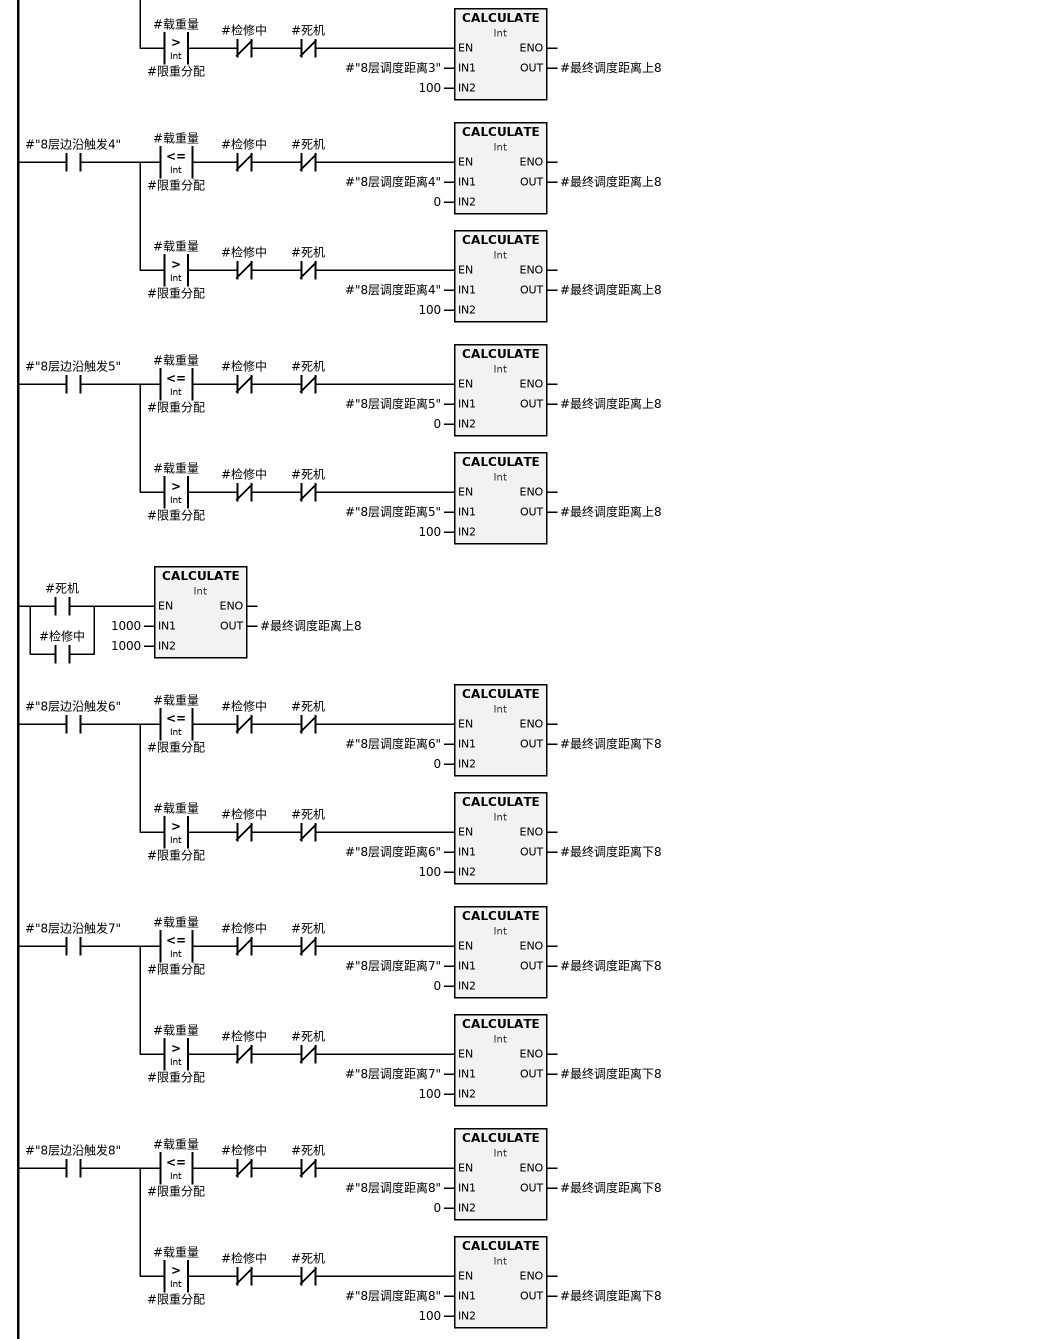
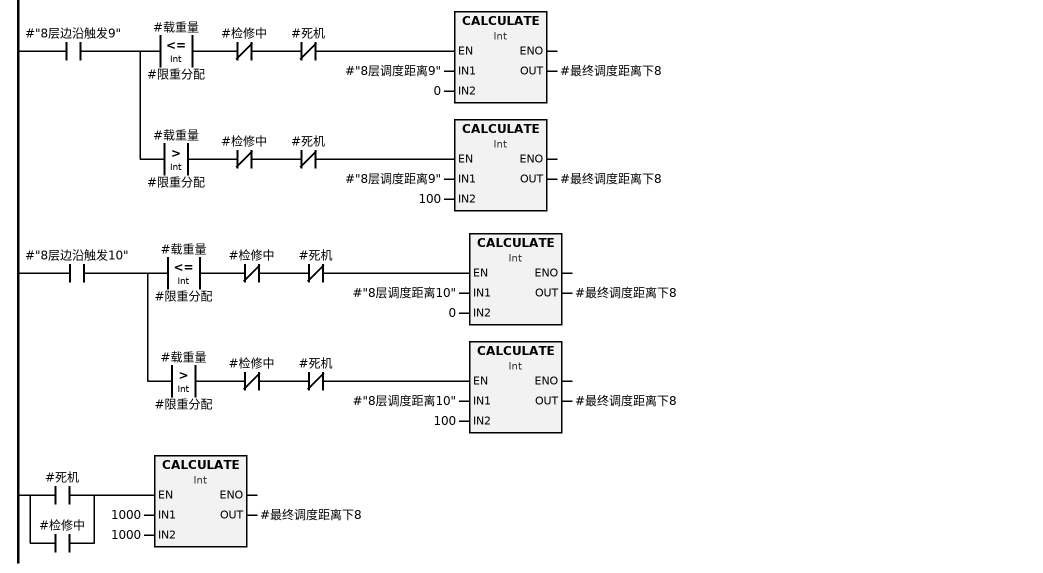
   RUNG wire#powerrail
      Contact( #上呼灯8 )
      wire#w1
      I_Contact( #上行指示 )
      I_Contact( #下行指示 )
      { S7_Templates := "SrcType := Int" } LE_Contact(in1 := #当前楼层, in2 := 8)
      wire#w2
      { S7_Templates := "SrcType := Int"; S7_Expression := "ABS(IN1-IN2)+IN3+IN3" } Calculate(in1 := #当前楼层, in2 := 8, in3 := #上行停站次数8, out => #"8层调度距离1")
      Coil( #"8层边沿触发1" )
   END_RUNG
   RUNG wire#w1
      Contact( #上行指示 )
      wire#w3
      { S7_Templates := "SrcType := Int" } EQ_Contact(in1 := 8, in2 := #当前楼层)
      Contact( #上下平层都为1 )
   END_RUNG wire#w2
   RUNG wire#w3
      { S7_Templates := "SrcType := Int" } GT_Contact(in1 := 8, in2 := #当前楼层)
   END_RUNG wire#w2
   RUNG wire#w1
      Contact( #下行指示 )
      wire#w4
      Contact( #外呼下面无目标8 )
      { S7_Templates := "SrcType := Int"; S7_Expression := "ABS(IN1-IN2)+IN3+IN3" } Calculate(in1 := #当前楼层, in2 := 8, in3 := #下行停站次数8, out => #"8层调度距离2")
      Coil( #"8层边沿触发2" )
   END_RUNG
   RUNG wire#w1
      I_Contact( #上行指示 )
      I_Contact( #下行指示 )
      { S7_Templates := "SrcType := Int" } GT_Contact(in1 := #当前楼层, in2 := 8)
   END_RUNG wire#w4
   RUNG wire#w1
      Contact( #下行指示 )
      Contact( #外呼下面有目标8 )
      { S7_Templates := "SrcType := Int"; S7_Expression := "ABS(IN3+IN3-IN1-IN2)+IN5+IN4+IN4+IN5+IN6" } Calculate(in1 := #当前楼层, in2 := 8, in3 := #外呼下面有目标最小数8, in4 := #上行停站次数8, in5 := #下行停站次数1, in6 := 2, out => #"8层调度距离3")
      Coil( #"8层边沿触发3" )
   END_RUNG
   RUNG wire#w1
      Contact( #上行指示 )
      wire#w5
      { S7_Templates := "SrcType := Int" } EQ_Contact(in1 := 8, in2 := #当前楼层)
      I_Contact( #上下平层都为1 )
      wire#w6
      Contact( #外呼下面有目标8 )
      { S7_Templates := "SrcType := Int"; S7_Expression := "ABS(IN3-IN1+IN3-IN6+IN2-IN6)+IN5+IN4+IN4+IN5+IN7+IN7" } Calculate(in1 := #当前楼层, in2 := 8, in3 := #外呼上面有目标最大数8, in4 := #上行停站次数10, in5 := #上行停站次数8, in6 := #外呼下面有目标最小数8, in7 := #下行停站次数1, in8 := 4, out => #"8层调度距离4")
      Coil( #"8层边沿触发4" )
   END_RUNG
   RUNG wire#w5
      { S7_Templates := "SrcType := Int" } LT_Contact(in1 := 8, in2 := #当前楼层)
   END_RUNG wire#w6
   RUNG wire#w6
      Contact( #外呼下面无目标8 )
      { S7_Templates := "SrcType := Int"; S7_Expression := "ABS(IN3-IN1+IN3-IN2)+IN5+IN4+IN4+IN5+IN6" } Calculate(in1 := #当前楼层, in2 := 8, in3 := #外呼上面有目标最大数8, in4 := #上行停站次数10, in5 := #下行停站次数8, in6 := 2, out => #"8层调度距离5")
      Coil( #"8层边沿触发5" )
   END_RUNG
   RUNG wire#powerrail
      Contact( #下呼灯8 )
      wire#w7
      I_Contact( #上行指示 )
      I_Contact( #下行指示 )
      { S7_Templates := "SrcType := Int" } GE_Contact(in1 := #当前楼层, in2 := 8)
      wire#w8
      { S7_Templates := "SrcType := Int"; S7_Expression := "ABS(IN1-IN2)+IN3+IN3" } Calculate(in1 := #当前楼层, in2 := 8, in3 := #下行停站次数8, out => #"8层调度距离6")
      Coil( #"8层边沿触发6" )
   END_RUNG
   RUNG wire#w7
      Contact( #下行指示 )
      wire#w9
      { S7_Templates := "SrcType := Int" } EQ_Contact(in1 := 8, in2 := #当前楼层)
      Contact( #上下平层都为1 )
   END_RUNG wire#w8
   RUNG wire#w9
      { S7_Templates := "SrcType := Int" } LT_Contact(in1 := 8, in2 := #当前楼层)
   END_RUNG wire#w8
   RUNG wire#w7
      Contact( #上行指示 )
      wire#w10
      Contact( #外呼上面无目标8 )
      { S7_Templates := "SrcType := Int"; S7_Expression := "ABS(IN1-IN2)+IN3+IN3" } Calculate(in1 := #当前楼层, in2 := 8, in3 := #上行停站次数8, out => #"8层调度距离7")
      Coil( #"8层边沿触发7" )
   END_RUNG
   RUNG wire#w7
      I_Contact( #上行指示 )
      I_Contact( #下行指示 )
      { S7_Templates := "SrcType := Int" } LT_Contact(in1 := #当前楼层, in2 := 8)
   END_RUNG wire#w10
   RUNG wire#w7
      Contact( #上行指示 )
      Contact( #外呼上面有目标8 )
      { S7_Templates := "SrcType := Int"; S7_Expression := "ABS(IN3+IN3-IN1-IN2)+IN4+IN5+IN4+IN5+IN6" } Calculate(in1 := #当前楼层, in2 := 8, in3 := #外呼上面有目标最大数8, in4 := #下行停站次数8, in5 := #上行停站次数10, in6 := 2, out => #"8层调度距离8")
      Coil( #"8层边沿触发8" )
   END_RUNG
   RUNG wire#w7
      Contact( #下行指示 )
      wire#w11
      { S7_Templates := "SrcType := Int" } EQ_Contact(in1 := 8, in2 := #当前楼层)
      I_Contact( #上下平层都为1 )
      wire#w12
      Contact( #外呼上面有目标8 )
      { S7_Templates := "SrcType := Int"; S7_Expression := "ABS(IN1-IN6+IN3-IN6+IN3-IN2)+IN5+IN4+IN4+IN5+IN7+IN7+IN8" } Calculate(in1 := #当前楼层, in2 := 8, in3 := #外呼上面有目标最大数8, in4 := #下行停站次数8, in5 := #下行停站次数1, in6 := #外呼下面有目标最小数8, in7 := #上行停站次数10, in8 := 4, out => #"8层调度距离9")
      Coil( #"8层边沿触发9" )
   END_RUNG
   RUNG wire#w11
      { S7_Templates := "SrcType := Int" } GT_Contact(in1 := 8, in2 := #当前楼层)
   END_RUNG wire#w12
   RUNG wire#w12
      Contact( #外呼上面无目标8 )
      { S7_Templates := "SrcType := Int"; S7_Expression := "ABS(IN1-IN3+IN2-IN3)+IN5+IN4+IN4+IN5+IN6" } Calculate(in1 := #当前楼层, in2 := 8, in3 := #外呼下面有目标最小数8, in4 := #上行停站次数8, in5 := #下行停站次数1, in6 := 2, out => #"8层调度距离10")
      Coil( #"8层边沿触发10" )
   END_RUNG
   RUNG wire#powerrail
      Contact( #"8层边沿触发1" )
      wire#w13
      { S7_Templates := "SrcType := Int" } LE_Contact(in1 := #载重量, in2 := #限重分配)
      I_Contact( #检修中 )
      I_Contact( #死机 )
      { S7_Templates := "SrcType := Int"; S7_Expression := "ABS(IN1+IN2)" } Calculate(in1 := #"8层调度距离1", in2 := 0, out => #最终调度距离上8)
   END_RUNG
   RUNG wire#w13
      { S7_Templates := "SrcType := Int" } GT_Contact(in1 := #载重量, in2 := #限重分配)
      I_Contact( #检修中 )
      I_Contact( #死机 )
      { S7_Templates := "SrcType := Int"; S7_Expression := "ABS(IN1+IN2)" } Calculate(in1 := #"8层调度距离1", in2 := 100, out => #最终调度距离上8)
   END_RUNG
   RUNG wire#powerrail
      Contact( #"8层边沿触发2" )
      wire#w14
      { S7_Templates := "SrcType := Int" } LE_Contact(in1 := #载重量, in2 := #限重分配)
      I_Contact( #检修中 )
      I_Contact( #死机 )
      { S7_Templates := "SrcType := Int"; S7_Expression := "ABS(IN1+IN2)" } Calculate(in1 := #"8层调度距离2", in2 := 0, out => #最终调度距离上8)
   END_RUNG
   RUNG wire#w14
      { S7_Templates := "SrcType := Int" } GT_Contact(in1 := #载重量, in2 := #限重分配)
      I_Contact( #检修中 )
      I_Contact( #死机 )
      { S7_Templates := "SrcType := Int"; S7_Expression := "ABS(IN1+IN2)" } Calculate(in1 := #"8层调度距离2", in2 := 100, out => #最终调度距离上8)
   END_RUNG
   RUNG wire#powerrail
      Contact( #"8层边沿触发3" )
      wire#w15
      { S7_Templates := "SrcType := Int" } LE_Contact(in1 := #载重量, in2 := #限重分配)
      I_Contact( #检修中 )
      I_Contact( #死机 )
      { S7_Templates := "SrcType := Int"; S7_Expression := "ABS(IN1+IN2)" } Calculate(in1 := #"8层调度距离3", in2 := 0, out => #最终调度距离上8)
   END_RUNG
   RUNG wire#w15
      { S7_Templates := "SrcType := Int" } GT_Contact(in1 := #载重量, in2 := #限重分配)
      I_Contact( #检修中 )
      I_Contact( #死机 )
      { S7_Templates := "SrcType := Int"; S7_Expression := "ABS(IN1+IN2)" } Calculate(in1 := #"8层调度距离3", in2 := 100, out => #最终调度距离上8)
   END_RUNG
   RUNG wire#powerrail
      Contact( #"8层边沿触发4" )
      wire#w16
      { S7_Templates := "SrcType := Int" } LE_Contact(in1 := #载重量, in2 := #限重分配)
      I_Contact( #检修中 )
      I_Contact( #死机 )
      { S7_Templates := "SrcType := Int"; S7_Expression := "ABS(IN1+IN2)" } Calculate(in1 := #"8层调度距离4", in2 := 0, out => #最终调度距离上8)
   END_RUNG
   RUNG wire#w16
      { S7_Templates := "SrcType := Int" } GT_Contact(in1 := #载重量, in2 := #限重分配)
      I_Contact( #检修中 )
      I_Contact( #死机 )
      { S7_Templates := "SrcType := Int"; S7_Expression := "ABS(IN1+IN2)" } Calculate(in1 := #"8层调度距离4", in2 := 100, out => #最终调度距离上8)
   END_RUNG
   RUNG wire#powerrail
      Contact( #"8层边沿触发5" )
      wire#w17
      { S7_Templates := "SrcType := Int" } LE_Contact(in1 := #载重量, in2 := #限重分配)
      I_Contact( #检修中 )
      I_Contact( #死机 )
      { S7_Templates := "SrcType := Int"; S7_Expression := "ABS(IN1+IN2)" } Calculate(in1 := #"8层调度距离5", in2 := 0, out => #最终调度距离上8)
   END_RUNG
   RUNG wire#w17
      { S7_Templates := "SrcType := Int" } GT_Contact(in1 := #载重量, in2 := #限重分配)
      I_Contact( #检修中 )
      I_Contact( #死机 )
      { S7_Templates := "SrcType := Int"; S7_Expression := "ABS(IN1+IN2)" } Calculate(in1 := #"8层调度距离5", in2 := 100, out => #最终调度距离上8)
   END_RUNG
   RUNG wire#powerrail
      Contact( #死机 )
      wire#w18
      { S7_Templates := "SrcType := Int"; S7_Expression := "ABS(IN1+IN2)" } Calculate(in1 := 1000, in2 := 1000, out => #最终调度距离上8)
   END_RUNG
   RUNG wire#powerrail
      Contact( #检修中 )
   END_RUNG wire#w18
   RUNG wire#powerrail
      Contact( #"8层边沿触发6" )
      wire#w19
      { S7_Templates := "SrcType := Int" } LE_Contact(in1 := #载重量, in2 := #限重分配)
      I_Contact( #检修中 )
      I_Contact( #死机 )
      { S7_Templates := "SrcType := Int"; S7_Expression := "ABS(IN1+IN2)" } Calculate(in1 := #"8层调度距离6", in2 := 0, out => #最终调度距离下8)
   END_RUNG
   RUNG wire#w19
      { S7_Templates := "SrcType := Int" } GT_Contact(in1 := #载重量, in2 := #限重分配)
      I_Contact( #检修中 )
      I_Contact( #死机 )
      { S7_Templates := "SrcType := Int"; S7_Expression := "ABS(IN1+IN2)" } Calculate(in1 := #"8层调度距离6", in2 := 100, out => #最终调度距离下8)
   END_RUNG
   RUNG wire#powerrail
      Contact( #"8层边沿触发7" )
      wire#w20
      { S7_Templates := "SrcType := Int" } LE_Contact(in1 := #载重量, in2 := #限重分配)
      I_Contact( #检修中 )
      I_Contact( #死机 )
      { S7_Templates := "SrcType := Int"; S7_Expression := "ABS(IN1+IN2)" } Calculate(in1 := #"8层调度距离7", in2 := 0, out => #最终调度距离下8)
   END_RUNG
   RUNG wire#w20
      { S7_Templates := "SrcType := Int" } GT_Contact(in1 := #载重量, in2 := #限重分配)
      I_Contact( #检修中 )
      I_Contact( #死机 )
      { S7_Templates := "SrcType := Int"; S7_Expression := "ABS(IN1+IN2)" } Calculate(in1 := #"8层调度距离7", in2 := 100, out => #最终调度距离下8)
   END_RUNG
   RUNG wire#powerrail
      Contact( #"8层边沿触发8" )
      wire#w21
      { S7_Templates := "SrcType := Int" } LE_Contact(in1 := #载重量, in2 := #限重分配)
      I_Contact( #检修中 )
      I_Contact( #死机 )
      { S7_Templates := "SrcType := Int"; S7_Expression := "ABS(IN1+IN2)" } Calculate(in1 := #"8层调度距离8", in2 := 0, out => #最终调度距离下8)
   END_RUNG
   RUNG wire#w21
      { S7_Templates := "SrcType := Int" } GT_Contact(in1 := #载重量, in2 := #限重分配)
      I_Contact( #检修中 )
      I_Contact( #死机 )
      { S7_Templates := "SrcType := Int"; S7_Expression := "ABS(IN1+IN2)" } Calculate(in1 := #"8层调度距离8", in2 := 100, out => #最终调度距离下8)
   END_RUNG
   RUNG wire#powerrail
      Contact( #"8层边沿触发9" )
      wire#w22
      { S7_Templates := "SrcType := Int" } LE_Contact(in1 := #载重量, in2 := #限重分配)
      I_Contact( #检修中 )
      I_Contact( #死机 )
      { S7_Templates := "SrcType := Int"; S7_Expression := "ABS(IN1+IN2)" } Calculate(in1 := #"8层调度距离9", in2 := 0, out => #最终调度距离下8)
   END_RUNG
   RUNG wire#w22
      { S7_Templates := "SrcType := Int" } GT_Contact(in1 := #载重量, in2 := #限重分配)
      I_Contact( #检修中 )
      I_Contact( #死机 )
      { S7_Templates := "SrcType := Int"; S7_Expression := "ABS(IN1+IN2)" } Calculate(in1 := #"8层调度距离9", in2 := 100, out => #最终调度距离下8)
   END_RUNG
   RUNG wire#powerrail
      Contact( #"8层边沿触发10" )
      wire#w23
      { S7_Templates := "SrcType := Int" } LE_Contact(in1 := #载重量, in2 := #限重分配)
      I_Contact( #检修中 )
      I_Contact( #死机 )
      { S7_Templates := "SrcType := Int"; S7_Expression := "ABS(IN1+IN2)" } Calculate(in1 := #"8层调度距离10", in2 := 0, out => #最终调度距离下8)
   END_RUNG
   RUNG wire#w23
      { S7_Templates := "SrcType := Int" } GT_Contact(in1 := #载重量, in2 := #限重分配)
      I_Contact( #检修中 )
      I_Contact( #死机 )
      { S7_Templates := "SrcType := Int"; S7_Expression := "ABS(IN1+IN2)" } Calculate(in1 := #"8层调度距离10", in2 := 100, out => #最终调度距离下8)
   END_RUNG
   RUNG wire#powerrail
      Contact( #死机 )
      wire#w24
      { S7_Templates := "SrcType := Int"; S7_Expression := "ABS(IN1+IN2)" } Calculate(in1 := 1000, in2 := 1000, out => #最终调度距离下8)
   END_RUNG
   RUNG wire#powerrail
      Contact( #检修中 )
   END_RUNG wire#w24
   // the same network as SCL:
   #_w1 := #上呼灯8 AND ((NOT #上行指示 AND NOT #下行指示 AND (#当前楼层 <= 8)) OR (#上行指示 AND (((8 = #当前楼层) AND #上下平层都为1) OR (8 > #当前楼层))));
   IF #_w1 THEN #"8层调度距离1" := ABS(#当前楼层-8)+#上行停站次数8+#上行停站次数8; END_IF;
   #"8层边沿触发1" := #_w1;
   #_w2 := #上呼灯8 AND (#下行指示 OR (NOT #上行指示 AND NOT #下行指示 AND (#当前楼层 > 8))) AND #外呼下面无目标8;
   IF #_w2 THEN #"8层调度距离2" := ABS(#当前楼层-8)+#下行停站次数8+#下行停站次数8; END_IF;
   #"8层边沿触发2" := #_w2;
   #_w3 := #上呼灯8 AND #下行指示 AND #外呼下面有目标8;
   IF #_w3 THEN
       #"8层调度距离3" := ABS(#外呼下面有目标最小数8+#外呼下面有目标最小数8-#当前楼层-8)+#下行停站次数1+#上行停站次数8+#上行停站次数8+#下行停站次数1+2;
   END_IF;
   #"8层边沿触发3" := #_w3;
   #_w4 := #上呼灯8 AND #上行指示 AND (((8 = #当前楼层) AND NOT #上下平层都为1) OR (8 < #当前楼层));
   #_w5 := #_w4 AND #外呼下面有目标8;
   IF #_w5 THEN
       #"8层调度距离4" := ABS(#外呼上面有目标最大数8-#当前楼层+#外呼上面有目标最大数8-#外呼下面有目标最小数8+8-#外呼下面有目标最小数8)+#上行停站次数8+#上行停站次数10+#上行停站次数10+#上行停站次数8+#下行停站次数1+#下行停站次数1;
   END_IF;
   #"8层边沿触发4" := #_w5;
   #_w6 := #_w4 AND #外呼下面无目标8;
   IF #_w6 THEN
       #"8层调度距离5" := ABS(#外呼上面有目标最大数8-#当前楼层+#外呼上面有目标最大数8-8)+#下行停站次数8+#上行停站次数10+#上行停站次数10+#下行停站次数8+2;
   END_IF;
   #"8层边沿触发5" := #_w6;
   #_w7 := #下呼灯8 AND ((NOT #上行指示 AND NOT #下行指示 AND (#当前楼层 >= 8)) OR (#下行指示 AND (((8 = #当前楼层) AND #上下平层都为1) OR (8 < #当前楼层))));
   IF #_w7 THEN #"8层调度距离6" := ABS(#当前楼层-8)+#下行停站次数8+#下行停站次数8; END_IF;
   #"8层边沿触发6" := #_w7;
   #_w8 := #下呼灯8 AND (#上行指示 OR (NOT #上行指示 AND NOT #下行指示 AND (#当前楼层 < 8))) AND #外呼上面无目标8;
   IF #_w8 THEN #"8层调度距离7" := ABS(#当前楼层-8)+#上行停站次数8+#上行停站次数8; END_IF;
   #"8层边沿触发7" := #_w8;
   #_w9 := #下呼灯8 AND #上行指示 AND #外呼上面有目标8;
   IF #_w9 THEN
       #"8层调度距离8" := ABS(#外呼上面有目标最大数8+#外呼上面有目标最大数8-#当前楼层-8)+#下行停站次数8+#上行停站次数10+#下行停站次数8+#上行停站次数10+2;
   END_IF;
   #"8层边沿触发8" := #_w9;
   #_w10 := #下呼灯8 AND #下行指示 AND (((8 = #当前楼层) AND NOT #上下平层都为1) OR (8 > #当前楼层));
   #_w11 := #_w10 AND #外呼上面有目标8;
   IF #_w11 THEN
       #"8层调度距离9" := ABS(#当前楼层-#外呼下面有目标最小数8+#外呼上面有目标最大数8-#外呼下面有目标最小数8+#外呼上面有目标最大数8-8)+#下行停站次数1+#下行停站次数8+#下行停站次数8+#下行停站次数1+#上行停站次数10+#上行停站次数10+4;
   END_IF;
   #"8层边沿触发9" := #_w11;
   #_w12 := #_w10 AND #外呼上面无目标8;
   IF #_w12 THEN
       #"8层调度距离10" := ABS(#当前楼层-#外呼下面有目标最小数8+8-#外呼下面有目标最小数8)+#下行停站次数1+#上行停站次数8+#上行停站次数8+#下行停站次数1+2;
   END_IF;
   #"8层边沿触发10" := #_w12;
   IF #"8层边沿触发1" AND (#载重量 <= #限重分配) AND NOT #检修中 AND NOT #死机 THEN #最终调度距离上8 := ABS(#"8层调度距离1"+0); END_IF;
   IF #"8层边沿触发1" AND (#载重量 > #限重分配) AND NOT #检修中 AND NOT #死机 THEN #最终调度距离上8 := ABS(#"8层调度距离1"+100); END_IF;
   IF #"8层边沿触发2" AND (#载重量 <= #限重分配) AND NOT #检修中 AND NOT #死机 THEN #最终调度距离上8 := ABS(#"8层调度距离2"+0); END_IF;
   IF #"8层边沿触发2" AND (#载重量 > #限重分配) AND NOT #检修中 AND NOT #死机 THEN #最终调度距离上8 := ABS(#"8层调度距离2"+100); END_IF;
   IF #"8层边沿触发3" AND (#载重量 <= #限重分配) AND NOT #检修中 AND NOT #死机 THEN #最终调度距离上8 := ABS(#"8层调度距离3"+0); END_IF;
   IF #"8层边沿触发3" AND (#载重量 > #限重分配) AND NOT #检修中 AND NOT #死机 THEN #最终调度距离上8 := ABS(#"8层调度距离3"+100); END_IF;
   IF #"8层边沿触发4" AND (#载重量 <= #限重分配) AND NOT #检修中 AND NOT #死机 THEN #最终调度距离上8 := ABS(#"8层调度距离4"+0); END_IF;
   IF #"8层边沿触发4" AND (#载重量 > #限重分配) AND NOT #检修中 AND NOT #死机 THEN #最终调度距离上8 := ABS(#"8层调度距离4"+100); END_IF;
   IF #"8层边沿触发5" AND (#载重量 <= #限重分配) AND NOT #检修中 AND NOT #死机 THEN #最终调度距离上8 := ABS(#"8层调度距离5"+0); END_IF;
   IF #"8层边沿触发5" AND (#载重量 > #限重分配) AND NOT #检修中 AND NOT #死机 THEN #最终调度距离上8 := ABS(#"8层调度距离5"+100); END_IF;
   IF #死机 OR #检修中 THEN #最终调度距离上8 := ABS(1000+1000); END_IF;
   IF #"8层边沿触发6" AND (#载重量 <= #限重分配) AND NOT #检修中 AND NOT #死机 THEN #最终调度距离下8 := ABS(#"8层调度距离6"+0); END_IF;
   IF #"8层边沿触发6" AND (#载重量 > #限重分配) AND NOT #检修中 AND NOT #死机 THEN #最终调度距离下8 := ABS(#"8层调度距离6"+100); END_IF;
   IF #"8层边沿触发7" AND (#载重量 <= #限重分配) AND NOT #检修中 AND NOT #死机 THEN #最终调度距离下8 := ABS(#"8层调度距离7"+0); END_IF;
   IF #"8层边沿触发7" AND (#载重量 > #限重分配) AND NOT #检修中 AND NOT #死机 THEN #最终调度距离下8 := ABS(#"8层调度距离7"+100); END_IF;
   IF #"8层边沿触发8" AND (#载重量 <= #限重分配) AND NOT #检修中 AND NOT #死机 THEN #最终调度距离下8 := ABS(#"8层调度距离8"+0); END_IF;
   IF #"8层边沿触发8" AND (#载重量 > #限重分配) AND NOT #检修中 AND NOT #死机 THEN #最终调度距离下8 := ABS(#"8层调度距离8"+100); END_IF;
   IF #"8层边沿触发9" AND (#载重量 <= #限重分配) AND NOT #检修中 AND NOT #死机 THEN #最终调度距离下8 := ABS(#"8层调度距离9"+0); END_IF;
   IF #"8层边沿触发9" AND (#载重量 > #限重分配) AND NOT #检修中 AND NOT #死机 THEN #最终调度距离下8 := ABS(#"8层调度距离9"+100); END_IF;
   IF #"8层边沿触发10" AND (#载重量 <= #限重分配) AND NOT #检修中 AND NOT #死机 THEN #最终调度距离下8 := ABS(#"8层调度距离10"+0); END_IF;
   IF #"8层边沿触发10" AND (#载重量 > #限重分配) AND NOT #检修中 AND NOT #死机 THEN #最终调度距离下8 := ABS(#"8层调度距离10"+100); END_IF;
   IF #死机 OR #检修中 THEN #最终调度距离下8 := ABS(1000+1000); END_IF;
END_REGION

REGION Network 8: 9层调度距离
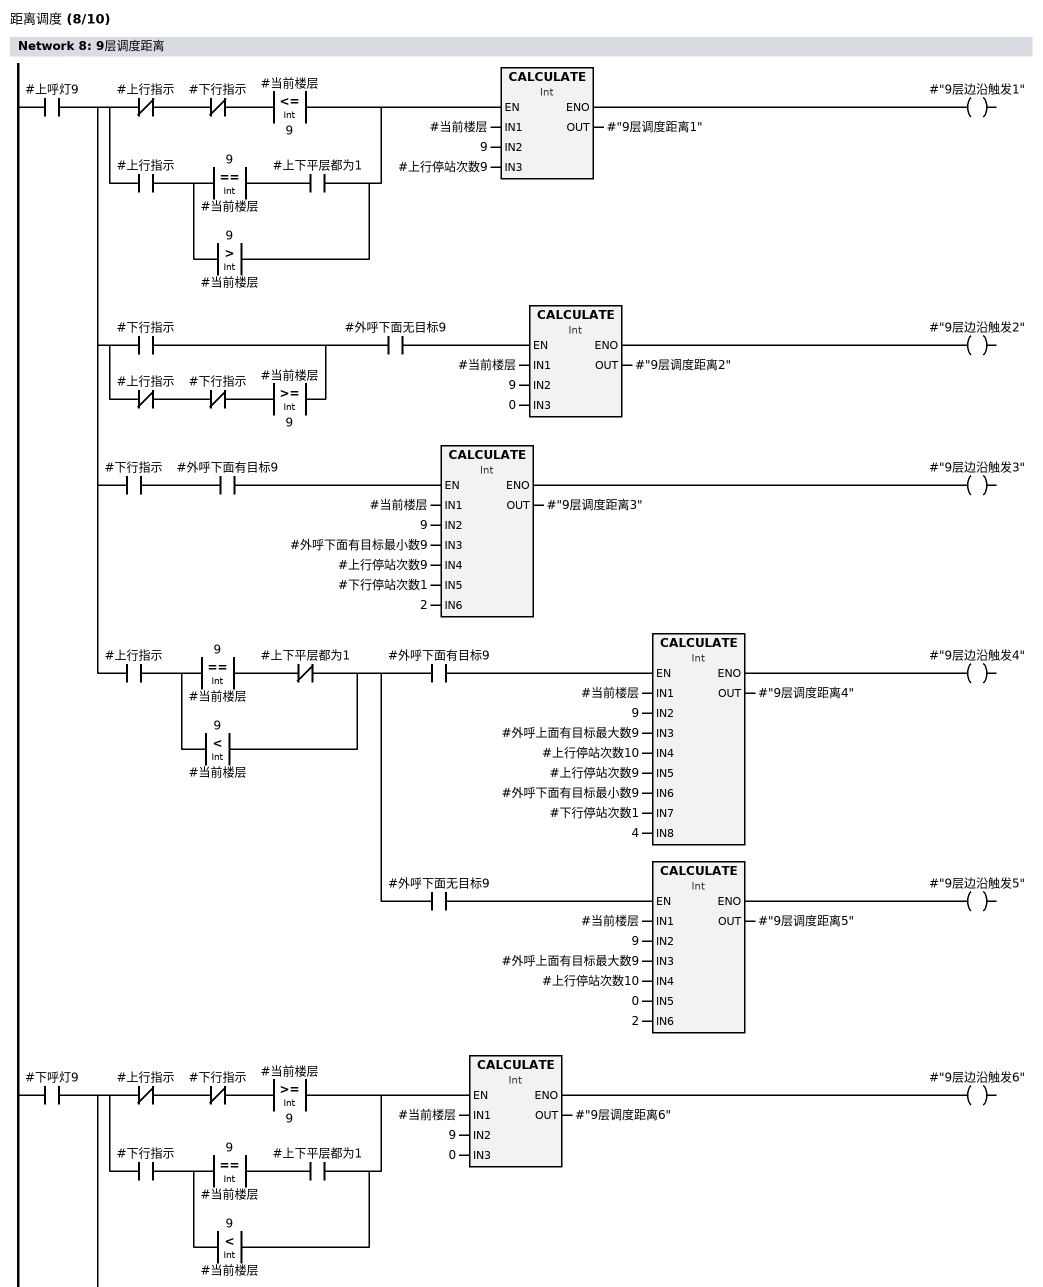
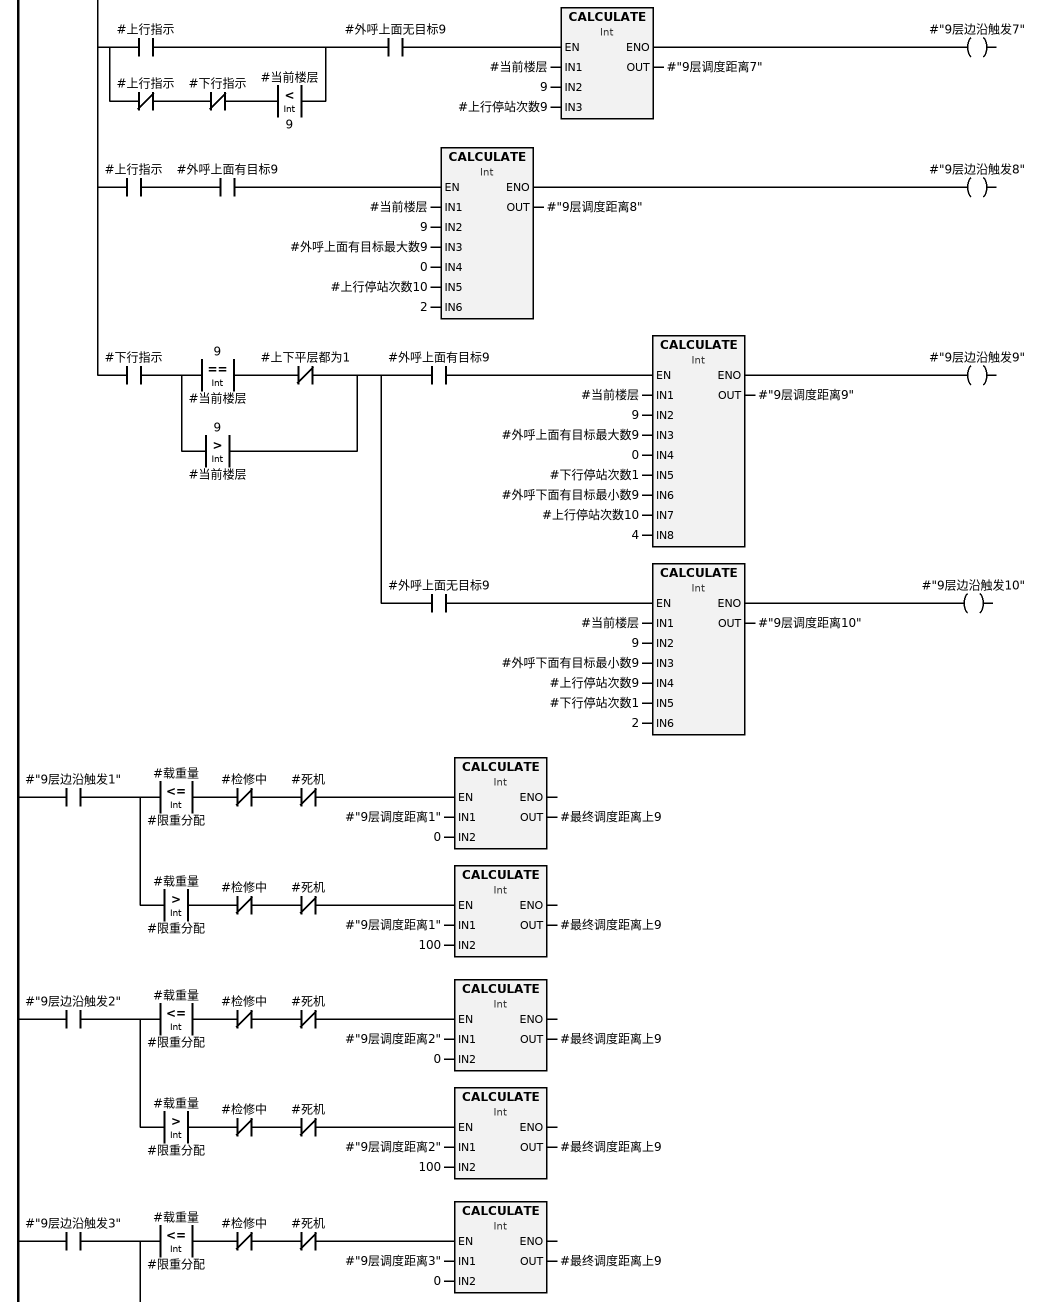
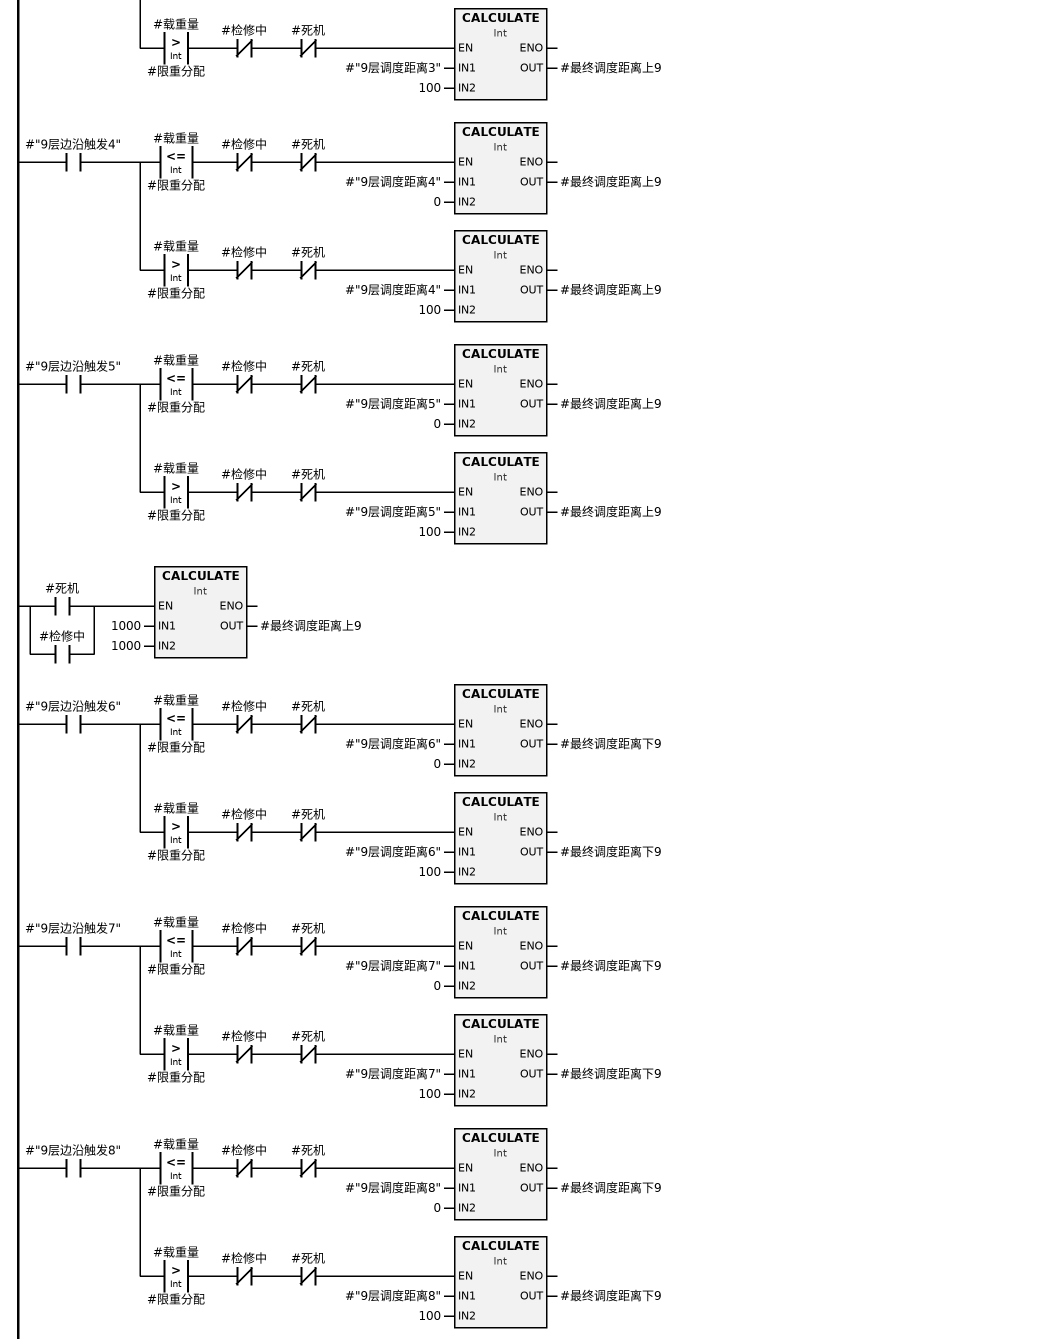
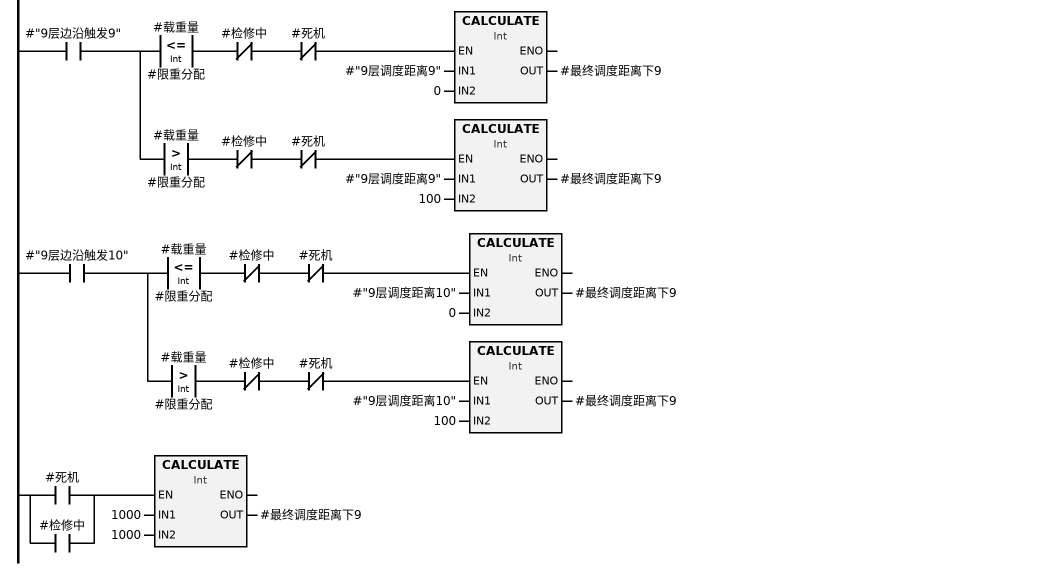
   RUNG wire#powerrail
      Contact( #上呼灯9 )
      wire#w1
      I_Contact( #上行指示 )
      I_Contact( #下行指示 )
      { S7_Templates := "SrcType := Int" } LE_Contact(in1 := #当前楼层, in2 := 9)
      wire#w2
      { S7_Templates := "SrcType := Int"; S7_Expression := "ABS(IN1-IN2)+IN3+IN3" } Calculate(in1 := #当前楼层, in2 := 9, in3 := #上行停站次数9, out => #"9层调度距离1")
      Coil( #"9层边沿触发1" )
   END_RUNG
   RUNG wire#w1
      Contact( #上行指示 )
      wire#w3
      { S7_Templates := "SrcType := Int" } EQ_Contact(in1 := 9, in2 := #当前楼层)
      Contact( #上下平层都为1 )
   END_RUNG wire#w2
   RUNG wire#w3
      { S7_Templates := "SrcType := Int" } GT_Contact(in1 := 9, in2 := #当前楼层)
   END_RUNG wire#w2
   RUNG wire#w1
      Contact( #下行指示 )
      wire#w4
      Contact( #外呼下面无目标9 )
      { S7_Templates := "SrcType := Int"; S7_Expression := "ABS(IN1-IN2)+IN3+IN3" } Calculate(in1 := #当前楼层, in2 := 9, in3 := 0, out => #"9层调度距离2")
      Coil( #"9层边沿触发2" )
   END_RUNG
   RUNG wire#w1
      I_Contact( #上行指示 )
      I_Contact( #下行指示 )
      { S7_Templates := "SrcType := Int" } GE_Contact(in1 := #当前楼层, in2 := 9)
   END_RUNG wire#w4
   RUNG wire#w1
      Contact( #下行指示 )
      Contact( #外呼下面有目标9 )
      { S7_Templates := "SrcType := Int"; S7_Expression := "ABS(IN3+IN3-IN1-IN2)+IN5+IN4+IN4+IN5+IN6" } Calculate(in1 := #当前楼层, in2 := 9, in3 := #外呼下面有目标最小数9, in4 := #上行停站次数9, in5 := #下行停站次数1, in6 := 2, out => #"9层调度距离3")
      Coil( #"9层边沿触发3" )
   END_RUNG
   RUNG wire#w1
      Contact( #上行指示 )
      wire#w5
      { S7_Templates := "SrcType := Int" } EQ_Contact(in1 := 9, in2 := #当前楼层)
      I_Contact( #上下平层都为1 )
      wire#w6
      Contact( #外呼下面有目标9 )
      { S7_Templates := "SrcType := Int"; S7_Expression := "ABS(IN3-IN1+IN3-IN6+IN2-IN6)+IN5+IN4+IN4+IN5+IN7+IN7+IN8" } Calculate(in1 := #当前楼层, in2 := 9, in3 := #外呼上面有目标最大数9, in4 := #上行停站次数10, in5 := #上行停站次数9, in6 := #外呼下面有目标最小数9, in7 := #下行停站次数1, in8 := 4, out => #"9层调度距离4")
      Coil( #"9层边沿触发4" )
   END_RUNG
   RUNG wire#w5
      { S7_Templates := "SrcType := Int" } LT_Contact(in1 := 9, in2 := #当前楼层)
   END_RUNG wire#w6
   RUNG wire#w6
      Contact( #外呼下面无目标9 )
      { S7_Templates := "SrcType := Int"; S7_Expression := "ABS(IN3-IN1+IN3-IN2)+IN5+IN4+IN4+IN5+IN6" } Calculate(in1 := #当前楼层, in2 := 9, in3 := #外呼上面有目标最大数9, in4 := #上行停站次数10, in5 := 0, in6 := 2, out => #"9层调度距离5")
      Coil( #"9层边沿触发5" )
   END_RUNG
   RUNG wire#powerrail
      Contact( #下呼灯9 )
      wire#w7
      I_Contact( #上行指示 )
      I_Contact( #下行指示 )
      { S7_Templates := "SrcType := Int" } GE_Contact(in1 := #当前楼层, in2 := 9)
      wire#w8
      { S7_Templates := "SrcType := Int"; S7_Expression := "ABS(IN1-IN2)+IN3+IN3" } Calculate(in1 := #当前楼层, in2 := 9, in3 := 0, out => #"9层调度距离6")
      Coil( #"9层边沿触发6" )
   END_RUNG
   RUNG wire#w7
      Contact( #下行指示 )
      wire#w9
      { S7_Templates := "SrcType := Int" } EQ_Contact(in1 := 9, in2 := #当前楼层)
      Contact( #上下平层都为1 )
   END_RUNG wire#w8
   RUNG wire#w9
      { S7_Templates := "SrcType := Int" } LT_Contact(in1 := 9, in2 := #当前楼层)
   END_RUNG wire#w8
   RUNG wire#w7
      Contact( #上行指示 )
      wire#w10
      Contact( #外呼上面无目标9 )
      { S7_Templates := "SrcType := Int"; S7_Expression := "ABS(IN1-IN2)+IN3+IN3" } Calculate(in1 := #当前楼层, in2 := 9, in3 := #上行停站次数9, out => #"9层调度距离7")
      Coil( #"9层边沿触发7" )
   END_RUNG
   RUNG wire#w7
      I_Contact( #上行指示 )
      I_Contact( #下行指示 )
      { S7_Templates := "SrcType := Int" } LT_Contact(in1 := #当前楼层, in2 := 9)
   END_RUNG wire#w10
   RUNG wire#w7
      Contact( #上行指示 )
      Contact( #外呼上面有目标9 )
      { S7_Templates := "SrcType := Int"; S7_Expression := "ABS(IN3+IN3-IN1-IN2)+IN4+IN5+IN4+IN5+IN6" } Calculate(in1 := #当前楼层, in2 := 9, in3 := #外呼上面有目标最大数9, in4 := 0, in5 := #上行停站次数10, in6 := 2, out => #"9层调度距离8")
      Coil( #"9层边沿触发8" )
   END_RUNG
   RUNG wire#w7
      Contact( #下行指示 )
      wire#w11
      { S7_Templates := "SrcType := Int" } EQ_Contact(in1 := 9, in2 := #当前楼层)
      I_Contact( #上下平层都为1 )
      wire#w12
      Contact( #外呼上面有目标9 )
      { S7_Templates := "SrcType := Int"; S7_Expression := "ABS(IN1-IN6+IN3-IN6+IN3-IN2)+IN5+IN4+IN4+IN5+IN7+IN7+IN8" } Calculate(in1 := #当前楼层, in2 := 9, in3 := #外呼上面有目标最大数9, in4 := 0, in5 := #下行停站次数1, in6 := #外呼下面有目标最小数9, in7 := #上行停站次数10, in8 := 4, out => #"9层调度距离9")
      Coil( #"9层边沿触发9" )
   END_RUNG
   RUNG wire#w11
      { S7_Templates := "SrcType := Int" } GT_Contact(in1 := 9, in2 := #当前楼层)
   END_RUNG wire#w12
   RUNG wire#w12
      Contact( #外呼上面无目标9 )
      { S7_Templates := "SrcType := Int"; S7_Expression := "ABS(IN1-IN3+IN2-IN3)+IN5+IN4+IN4+IN5+IN6" } Calculate(in1 := #当前楼层, in2 := 9, in3 := #外呼下面有目标最小数9, in4 := #上行停站次数9, in5 := #下行停站次数1, in6 := 2, out => #"9层调度距离10")
      Coil( #"9层边沿触发10" )
   END_RUNG
   RUNG wire#powerrail
      Contact( #"9层边沿触发1" )
      wire#w13
      { S7_Templates := "SrcType := Int" } LE_Contact(in1 := #载重量, in2 := #限重分配)
      I_Contact( #检修中 )
      I_Contact( #死机 )
      { S7_Templates := "SrcType := Int"; S7_Expression := "ABS(IN1+IN2)" } Calculate(in1 := #"9层调度距离1", in2 := 0, out => #最终调度距离上9)
   END_RUNG
   RUNG wire#w13
      { S7_Templates := "SrcType := Int" } GT_Contact(in1 := #载重量, in2 := #限重分配)
      I_Contact( #检修中 )
      I_Contact( #死机 )
      { S7_Templates := "SrcType := Int"; S7_Expression := "ABS(IN1+IN2)" } Calculate(in1 := #"9层调度距离1", in2 := 100, out => #最终调度距离上9)
   END_RUNG
   RUNG wire#powerrail
      Contact( #"9层边沿触发2" )
      wire#w14
      { S7_Templates := "SrcType := Int" } LE_Contact(in1 := #载重量, in2 := #限重分配)
      I_Contact( #检修中 )
      I_Contact( #死机 )
      { S7_Templates := "SrcType := Int"; S7_Expression := "ABS(IN1+IN2)" } Calculate(in1 := #"9层调度距离2", in2 := 0, out => #最终调度距离上9)
   END_RUNG
   RUNG wire#w14
      { S7_Templates := "SrcType := Int" } GT_Contact(in1 := #载重量, in2 := #限重分配)
      I_Contact( #检修中 )
      I_Contact( #死机 )
      { S7_Templates := "SrcType := Int"; S7_Expression := "ABS(IN1+IN2)" } Calculate(in1 := #"9层调度距离2", in2 := 100, out => #最终调度距离上9)
   END_RUNG
   RUNG wire#powerrail
      Contact( #"9层边沿触发3" )
      wire#w15
      { S7_Templates := "SrcType := Int" } LE_Contact(in1 := #载重量, in2 := #限重分配)
      I_Contact( #检修中 )
      I_Contact( #死机 )
      { S7_Templates := "SrcType := Int"; S7_Expression := "ABS(IN1+IN2)" } Calculate(in1 := #"9层调度距离3", in2 := 0, out => #最终调度距离上9)
   END_RUNG
   RUNG wire#w15
      { S7_Templates := "SrcType := Int" } GT_Contact(in1 := #载重量, in2 := #限重分配)
      I_Contact( #检修中 )
      I_Contact( #死机 )
      { S7_Templates := "SrcType := Int"; S7_Expression := "ABS(IN1+IN2)" } Calculate(in1 := #"9层调度距离3", in2 := 100, out => #最终调度距离上9)
   END_RUNG
   RUNG wire#powerrail
      Contact( #"9层边沿触发4" )
      wire#w16
      { S7_Templates := "SrcType := Int" } LE_Contact(in1 := #载重量, in2 := #限重分配)
      I_Contact( #检修中 )
      I_Contact( #死机 )
      { S7_Templates := "SrcType := Int"; S7_Expression := "ABS(IN1+IN2)" } Calculate(in1 := #"9层调度距离4", in2 := 0, out => #最终调度距离上9)
   END_RUNG
   RUNG wire#w16
      { S7_Templates := "SrcType := Int" } GT_Contact(in1 := #载重量, in2 := #限重分配)
      I_Contact( #检修中 )
      I_Contact( #死机 )
      { S7_Templates := "SrcType := Int"; S7_Expression := "ABS(IN1+IN2)" } Calculate(in1 := #"9层调度距离4", in2 := 100, out => #最终调度距离上9)
   END_RUNG
   RUNG wire#powerrail
      Contact( #"9层边沿触发5" )
      wire#w17
      { S7_Templates := "SrcType := Int" } LE_Contact(in1 := #载重量, in2 := #限重分配)
      I_Contact( #检修中 )
      I_Contact( #死机 )
      { S7_Templates := "SrcType := Int"; S7_Expression := "ABS(IN1+IN2)" } Calculate(in1 := #"9层调度距离5", in2 := 0, out => #最终调度距离上9)
   END_RUNG
   RUNG wire#w17
      { S7_Templates := "SrcType := Int" } GT_Contact(in1 := #载重量, in2 := #限重分配)
      I_Contact( #检修中 )
      I_Contact( #死机 )
      { S7_Templates := "SrcType := Int"; S7_Expression := "ABS(IN1+IN2)" } Calculate(in1 := #"9层调度距离5", in2 := 100, out => #最终调度距离上9)
   END_RUNG
   RUNG wire#powerrail
      Contact( #死机 )
      wire#w18
      { S7_Templates := "SrcType := Int"; S7_Expression := "ABS(IN1+IN2)" } Calculate(in1 := 1000, in2 := 1000, out => #最终调度距离上9)
   END_RUNG
   RUNG wire#powerrail
      Contact( #检修中 )
   END_RUNG wire#w18
   RUNG wire#powerrail
      Contact( #"9层边沿触发6" )
      wire#w19
      { S7_Templates := "SrcType := Int" } LE_Contact(in1 := #载重量, in2 := #限重分配)
      I_Contact( #检修中 )
      I_Contact( #死机 )
      { S7_Templates := "SrcType := Int"; S7_Expression := "ABS(IN1+IN2)" } Calculate(in1 := #"9层调度距离6", in2 := 0, out => #最终调度距离下9)
   END_RUNG
   RUNG wire#w19
      { S7_Templates := "SrcType := Int" } GT_Contact(in1 := #载重量, in2 := #限重分配)
      I_Contact( #检修中 )
      I_Contact( #死机 )
      { S7_Templates := "SrcType := Int"; S7_Expression := "ABS(IN1+IN2)" } Calculate(in1 := #"9层调度距离6", in2 := 100, out => #最终调度距离下9)
   END_RUNG
   RUNG wire#powerrail
      Contact( #"9层边沿触发7" )
      wire#w20
      { S7_Templates := "SrcType := Int" } LE_Contact(in1 := #载重量, in2 := #限重分配)
      I_Contact( #检修中 )
      I_Contact( #死机 )
      { S7_Templates := "SrcType := Int"; S7_Expression := "ABS(IN1+IN2)" } Calculate(in1 := #"9层调度距离7", in2 := 0, out => #最终调度距离下9)
   END_RUNG
   RUNG wire#w20
      { S7_Templates := "SrcType := Int" } GT_Contact(in1 := #载重量, in2 := #限重分配)
      I_Contact( #检修中 )
      I_Contact( #死机 )
      { S7_Templates := "SrcType := Int"; S7_Expression := "ABS(IN1+IN2)" } Calculate(in1 := #"9层调度距离7", in2 := 100, out => #最终调度距离下9)
   END_RUNG
   RUNG wire#powerrail
      Contact( #"9层边沿触发8" )
      wire#w21
      { S7_Templates := "SrcType := Int" } LE_Contact(in1 := #载重量, in2 := #限重分配)
      I_Contact( #检修中 )
      I_Contact( #死机 )
      { S7_Templates := "SrcType := Int"; S7_Expression := "ABS(IN1+IN2)" } Calculate(in1 := #"9层调度距离8", in2 := 0, out => #最终调度距离下9)
   END_RUNG
   RUNG wire#w21
      { S7_Templates := "SrcType := Int" } GT_Contact(in1 := #载重量, in2 := #限重分配)
      I_Contact( #检修中 )
      I_Contact( #死机 )
      { S7_Templates := "SrcType := Int"; S7_Expression := "ABS(IN1+IN2)" } Calculate(in1 := #"9层调度距离8", in2 := 100, out => #最终调度距离下9)
   END_RUNG
   RUNG wire#powerrail
      Contact( #"9层边沿触发9" )
      wire#w22
      { S7_Templates := "SrcType := Int" } LE_Contact(in1 := #载重量, in2 := #限重分配)
      I_Contact( #检修中 )
      I_Contact( #死机 )
      { S7_Templates := "SrcType := Int"; S7_Expression := "ABS(IN1+IN2)" } Calculate(in1 := #"9层调度距离9", in2 := 0, out => #最终调度距离下9)
   END_RUNG
   RUNG wire#w22
      { S7_Templates := "SrcType := Int" } GT_Contact(in1 := #载重量, in2 := #限重分配)
      I_Contact( #检修中 )
      I_Contact( #死机 )
      { S7_Templates := "SrcType := Int"; S7_Expression := "ABS(IN1+IN2)" } Calculate(in1 := #"9层调度距离9", in2 := 100, out => #最终调度距离下9)
   END_RUNG
   RUNG wire#powerrail
      Contact( #"9层边沿触发10" )
      wire#w23
      { S7_Templates := "SrcType := Int" } LE_Contact(in1 := #载重量, in2 := #限重分配)
      I_Contact( #检修中 )
      I_Contact( #死机 )
      { S7_Templates := "SrcType := Int"; S7_Expression := "ABS(IN1+IN2)" } Calculate(in1 := #"9层调度距离10", in2 := 0, out => #最终调度距离下9)
   END_RUNG
   RUNG wire#w23
      { S7_Templates := "SrcType := Int" } GT_Contact(in1 := #载重量, in2 := #限重分配)
      I_Contact( #检修中 )
      I_Contact( #死机 )
      { S7_Templates := "SrcType := Int"; S7_Expression := "ABS(IN1+IN2)" } Calculate(in1 := #"9层调度距离10", in2 := 100, out => #最终调度距离下9)
   END_RUNG
   RUNG wire#powerrail
      Contact( #死机 )
      wire#w24
      { S7_Templates := "SrcType := Int"; S7_Expression := "ABS(IN1+IN2)" } Calculate(in1 := 1000, in2 := 1000, out => #最终调度距离下9)
   END_RUNG
   RUNG wire#powerrail
      Contact( #检修中 )
   END_RUNG wire#w24
   // the same network as SCL:
   #_w1 := #上呼灯9 AND ((NOT #上行指示 AND NOT #下行指示 AND (#当前楼层 <= 9)) OR (#上行指示 AND (((9 = #当前楼层) AND #上下平层都为1) OR (9 > #当前楼层))));
   IF #_w1 THEN #"9层调度距离1" := ABS(#当前楼层-9)+#上行停站次数9+#上行停站次数9; END_IF;
   #"9层边沿触发1" := #_w1;
   #_w2 := #上呼灯9 AND (#下行指示 OR (NOT #上行指示 AND NOT #下行指示 AND (#当前楼层 >= 9))) AND #外呼下面无目标9;
   IF #_w2 THEN #"9层调度距离2" := ABS(#当前楼层-9)+0+0; END_IF;
   #"9层边沿触发2" := #_w2;
   #_w3 := #上呼灯9 AND #下行指示 AND #外呼下面有目标9;
   IF #_w3 THEN
       #"9层调度距离3" := ABS(#外呼下面有目标最小数9+#外呼下面有目标最小数9-#当前楼层-9)+#下行停站次数1+#上行停站次数9+#上行停站次数9+#下行停站次数1+2;
   END_IF;
   #"9层边沿触发3" := #_w3;
   #_w4 := #上呼灯9 AND #上行指示 AND (((9 = #当前楼层) AND NOT #上下平层都为1) OR (9 < #当前楼层));
   #_w5 := #_w4 AND #外呼下面有目标9;
   IF #_w5 THEN
       #"9层调度距离4" := ABS(#外呼上面有目标最大数9-#当前楼层+#外呼上面有目标最大数9-#外呼下面有目标最小数9+9-#外呼下面有目标最小数9)+#上行停站次数9+#上行停站次数10+#上行停站次数10+#上行停站次数9+#下行停站次数1+#下行停站次数1+4;
   END_IF;
   #"9层边沿触发4" := #_w5;
   #_w6 := #_w4 AND #外呼下面无目标9;
   IF #_w6 THEN #"9层调度距离5" := ABS(#外呼上面有目标最大数9-#当前楼层+#外呼上面有目标最大数9-9)+0+#上行停站次数10+#上行停站次数10+0+2; END_IF;
   #"9层边沿触发5" := #_w6;
   #_w7 := #下呼灯9 AND ((NOT #上行指示 AND NOT #下行指示 AND (#当前楼层 >= 9)) OR (#下行指示 AND (((9 = #当前楼层) AND #上下平层都为1) OR (9 < #当前楼层))));
   IF #_w7 THEN #"9层调度距离6" := ABS(#当前楼层-9)+0+0; END_IF;
   #"9层边沿触发6" := #_w7;
   #_w8 := #下呼灯9 AND (#上行指示 OR (NOT #上行指示 AND NOT #下行指示 AND (#当前楼层 < 9))) AND #外呼上面无目标9;
   IF #_w8 THEN #"9层调度距离7" := ABS(#当前楼层-9)+#上行停站次数9+#上行停站次数9; END_IF;
   #"9层边沿触发7" := #_w8;
   #_w9 := #下呼灯9 AND #上行指示 AND #外呼上面有目标9;
   IF #_w9 THEN #"9层调度距离8" := ABS(#外呼上面有目标最大数9+#外呼上面有目标最大数9-#当前楼层-9)+0+#上行停站次数10+0+#上行停站次数10+2; END_IF;
   #"9层边沿触发8" := #_w9;
   #_w10 := #下呼灯9 AND #下行指示 AND (((9 = #当前楼层) AND NOT #上下平层都为1) OR (9 > #当前楼层));
   #_w11 := #_w10 AND #外呼上面有目标9;
   IF #_w11 THEN
       #"9层调度距离9" := ABS(#当前楼层-#外呼下面有目标最小数9+#外呼上面有目标最大数9-#外呼下面有目标最小数9+#外呼上面有目标最大数9-9)+#下行停站次数1+0+0+#下行停站次数1+#上行停站次数10+#上行停站次数10+4;
   END_IF;
   #"9层边沿触发9" := #_w11;
   #_w12 := #_w10 AND #外呼上面无目标9;
   IF #_w12 THEN
       #"9层调度距离10" := ABS(#当前楼层-#外呼下面有目标最小数9+9-#外呼下面有目标最小数9)+#下行停站次数1+#上行停站次数9+#上行停站次数9+#下行停站次数1+2;
   END_IF;
   #"9层边沿触发10" := #_w12;
   IF #"9层边沿触发1" AND (#载重量 <= #限重分配) AND NOT #检修中 AND NOT #死机 THEN #最终调度距离上9 := ABS(#"9层调度距离1"+0); END_IF;
   IF #"9层边沿触发1" AND (#载重量 > #限重分配) AND NOT #检修中 AND NOT #死机 THEN #最终调度距离上9 := ABS(#"9层调度距离1"+100); END_IF;
   IF #"9层边沿触发2" AND (#载重量 <= #限重分配) AND NOT #检修中 AND NOT #死机 THEN #最终调度距离上9 := ABS(#"9层调度距离2"+0); END_IF;
   IF #"9层边沿触发2" AND (#载重量 > #限重分配) AND NOT #检修中 AND NOT #死机 THEN #最终调度距离上9 := ABS(#"9层调度距离2"+100); END_IF;
   IF #"9层边沿触发3" AND (#载重量 <= #限重分配) AND NOT #检修中 AND NOT #死机 THEN #最终调度距离上9 := ABS(#"9层调度距离3"+0); END_IF;
   IF #"9层边沿触发3" AND (#载重量 > #限重分配) AND NOT #检修中 AND NOT #死机 THEN #最终调度距离上9 := ABS(#"9层调度距离3"+100); END_IF;
   IF #"9层边沿触发4" AND (#载重量 <= #限重分配) AND NOT #检修中 AND NOT #死机 THEN #最终调度距离上9 := ABS(#"9层调度距离4"+0); END_IF;
   IF #"9层边沿触发4" AND (#载重量 > #限重分配) AND NOT #检修中 AND NOT #死机 THEN #最终调度距离上9 := ABS(#"9层调度距离4"+100); END_IF;
   IF #"9层边沿触发5" AND (#载重量 <= #限重分配) AND NOT #检修中 AND NOT #死机 THEN #最终调度距离上9 := ABS(#"9层调度距离5"+0); END_IF;
   IF #"9层边沿触发5" AND (#载重量 > #限重分配) AND NOT #检修中 AND NOT #死机 THEN #最终调度距离上9 := ABS(#"9层调度距离5"+100); END_IF;
   IF #死机 OR #检修中 THEN #最终调度距离上9 := ABS(1000+1000); END_IF;
   IF #"9层边沿触发6" AND (#载重量 <= #限重分配) AND NOT #检修中 AND NOT #死机 THEN #最终调度距离下9 := ABS(#"9层调度距离6"+0); END_IF;
   IF #"9层边沿触发6" AND (#载重量 > #限重分配) AND NOT #检修中 AND NOT #死机 THEN #最终调度距离下9 := ABS(#"9层调度距离6"+100); END_IF;
   IF #"9层边沿触发7" AND (#载重量 <= #限重分配) AND NOT #检修中 AND NOT #死机 THEN #最终调度距离下9 := ABS(#"9层调度距离7"+0); END_IF;
   IF #"9层边沿触发7" AND (#载重量 > #限重分配) AND NOT #检修中 AND NOT #死机 THEN #最终调度距离下9 := ABS(#"9层调度距离7"+100); END_IF;
   IF #"9层边沿触发8" AND (#载重量 <= #限重分配) AND NOT #检修中 AND NOT #死机 THEN #最终调度距离下9 := ABS(#"9层调度距离8"+0); END_IF;
   IF #"9层边沿触发8" AND (#载重量 > #限重分配) AND NOT #检修中 AND NOT #死机 THEN #最终调度距离下9 := ABS(#"9层调度距离8"+100); END_IF;
   IF #"9层边沿触发9" AND (#载重量 <= #限重分配) AND NOT #检修中 AND NOT #死机 THEN #最终调度距离下9 := ABS(#"9层调度距离9"+0); END_IF;
   IF #"9层边沿触发9" AND (#载重量 > #限重分配) AND NOT #检修中 AND NOT #死机 THEN #最终调度距离下9 := ABS(#"9层调度距离9"+100); END_IF;
   IF #"9层边沿触发10" AND (#载重量 <= #限重分配) AND NOT #检修中 AND NOT #死机 THEN #最终调度距离下9 := ABS(#"9层调度距离10"+0); END_IF;
   IF #"9层边沿触发10" AND (#载重量 > #限重分配) AND NOT #检修中 AND NOT #死机 THEN #最终调度距离下9 := ABS(#"9层调度距离10"+100); END_IF;
   IF #死机 OR #检修中 THEN #最终调度距离下9 := ABS(1000+1000); END_IF;
END_REGION

REGION Network 9: 1层调度距离
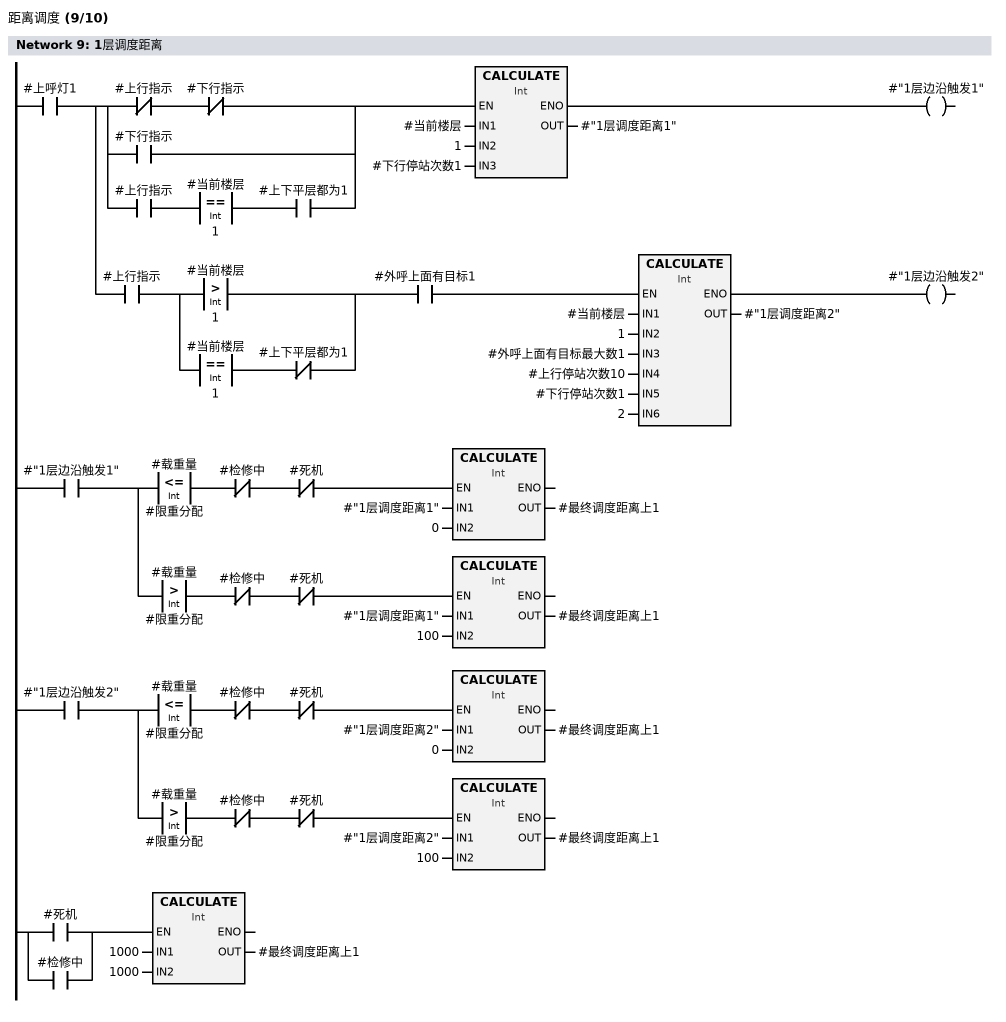
   RUNG wire#powerrail
      Contact( #上呼灯1 )
      wire#w1
      I_Contact( #上行指示 )
      I_Contact( #下行指示 )
      wire#w2
      { S7_Templates := "SrcType := Int"; S7_Expression := "ABS(IN1-IN2)+IN3+IN3" } Calculate(in1 := #当前楼层, in2 := 1, in3 := #下行停站次数1, out => #"1层调度距离1")
      Coil( #"1层边沿触发1" )
   END_RUNG
   RUNG wire#w1
      Contact( #下行指示 )
   END_RUNG wire#w2
   RUNG wire#w1
      Contact( #上行指示 )
      { S7_Templates := "SrcType := Int" } EQ_Contact(in1 := #当前楼层, in2 := 1)
      Contact( #上下平层都为1 )
   END_RUNG wire#w2
   RUNG wire#w1
      Contact( #上行指示 )
      wire#w3
      { S7_Templates := "SrcType := Int" } GT_Contact(in1 := #当前楼层, in2 := 1)
      wire#w4
      Contact( #外呼上面有目标1 )
      { S7_Templates := "SrcType := Int"; S7_Expression := "ABS(IN3+IN3-IN2-IN1)+IN4+IN5+IN4+IN5+IN6" } Calculate(in1 := #当前楼层, in2 := 1, in3 := #外呼上面有目标最大数1, in4 := #上行停站次数10, in5 := #下行停站次数1, in6 := 2, out => #"1层调度距离2")
      Coil( #"1层边沿触发2" )
   END_RUNG
   RUNG wire#w3
      { S7_Templates := "SrcType := Int" } EQ_Contact(in1 := #当前楼层, in2 := 1)
      I_Contact( #上下平层都为1 )
   END_RUNG wire#w4
   RUNG wire#powerrail
      Contact( #"1层边沿触发1" )
      wire#w5
      { S7_Templates := "SrcType := Int" } LE_Contact(in1 := #载重量, in2 := #限重分配)
      I_Contact( #检修中 )
      I_Contact( #死机 )
      { S7_Templates := "SrcType := Int"; S7_Expression := "ABS(IN1+IN2)" } Calculate(in1 := #"1层调度距离1", in2 := 0, out => #最终调度距离上1)
   END_RUNG
   RUNG wire#w5
      { S7_Templates := "SrcType := Int" } GT_Contact(in1 := #载重量, in2 := #限重分配)
      I_Contact( #检修中 )
      I_Contact( #死机 )
      { S7_Templates := "SrcType := Int"; S7_Expression := "ABS(IN1+IN2)" } Calculate(in1 := #"1层调度距离1", in2 := 100, out => #最终调度距离上1)
   END_RUNG
   RUNG wire#powerrail
      Contact( #"1层边沿触发2" )
      wire#w6
      { S7_Templates := "SrcType := Int" } LE_Contact(in1 := #载重量, in2 := #限重分配)
      I_Contact( #检修中 )
      I_Contact( #死机 )
      { S7_Templates := "SrcType := Int"; S7_Expression := "ABS(IN1+IN2)" } Calculate(in1 := #"1层调度距离2", in2 := 0, out => #最终调度距离上1)
   END_RUNG
   RUNG wire#w6
      { S7_Templates := "SrcType := Int" } GT_Contact(in1 := #载重量, in2 := #限重分配)
      I_Contact( #检修中 )
      I_Contact( #死机 )
      { S7_Templates := "SrcType := Int"; S7_Expression := "ABS(IN1+IN2)" } Calculate(in1 := #"1层调度距离2", in2 := 100, out => #最终调度距离上1)
   END_RUNG
   RUNG wire#powerrail
      Contact( #死机 )
      wire#w7
      { S7_Templates := "SrcType := Int"; S7_Expression := "ABS(IN1+IN2)" } Calculate(in1 := 1000, in2 := 1000, out => #最终调度距离上1)
   END_RUNG
   RUNG wire#powerrail
      Contact( #检修中 )
   END_RUNG wire#w7
   // the same network as SCL:
   #_w1 := #上呼灯1 AND ((NOT #上行指示 AND NOT #下行指示) OR #下行指示 OR (#上行指示 AND (#当前楼层 = 1) AND #上下平层都为1));
   IF #_w1 THEN #"1层调度距离1" := ABS(#当前楼层-1)+#下行停站次数1+#下行停站次数1; END_IF;
   #"1层边沿触发1" := #_w1;
   #_w2 := #上呼灯1 AND #上行指示 AND ((#当前楼层 > 1) OR ((#当前楼层 = 1) AND NOT #上下平层都为1)) AND #外呼上面有目标1;
   IF #_w2 THEN
       #"1层调度距离2" := ABS(#外呼上面有目标最大数1+#外呼上面有目标最大数1-1-#当前楼层)+#上行停站次数10+#下行停站次数1+#上行停站次数10+#下行停站次数1+2;
   END_IF;
   #"1层边沿触发2" := #_w2;
   IF #"1层边沿触发1" AND (#载重量 <= #限重分配) AND NOT #检修中 AND NOT #死机 THEN #最终调度距离上1 := ABS(#"1层调度距离1"+0); END_IF;
   IF #"1层边沿触发1" AND (#载重量 > #限重分配) AND NOT #检修中 AND NOT #死机 THEN #最终调度距离上1 := ABS(#"1层调度距离1"+100); END_IF;
   IF #"1层边沿触发2" AND (#载重量 <= #限重分配) AND NOT #检修中 AND NOT #死机 THEN #最终调度距离上1 := ABS(#"1层调度距离2"+0); END_IF;
   IF #"1层边沿触发2" AND (#载重量 > #限重分配) AND NOT #检修中 AND NOT #死机 THEN #最终调度距离上1 := ABS(#"1层调度距离2"+100); END_IF;
   IF #死机 OR #检修中 THEN #最终调度距离上1 := ABS(1000+1000); END_IF;
END_REGION

REGION Network 10: 10层调度距离
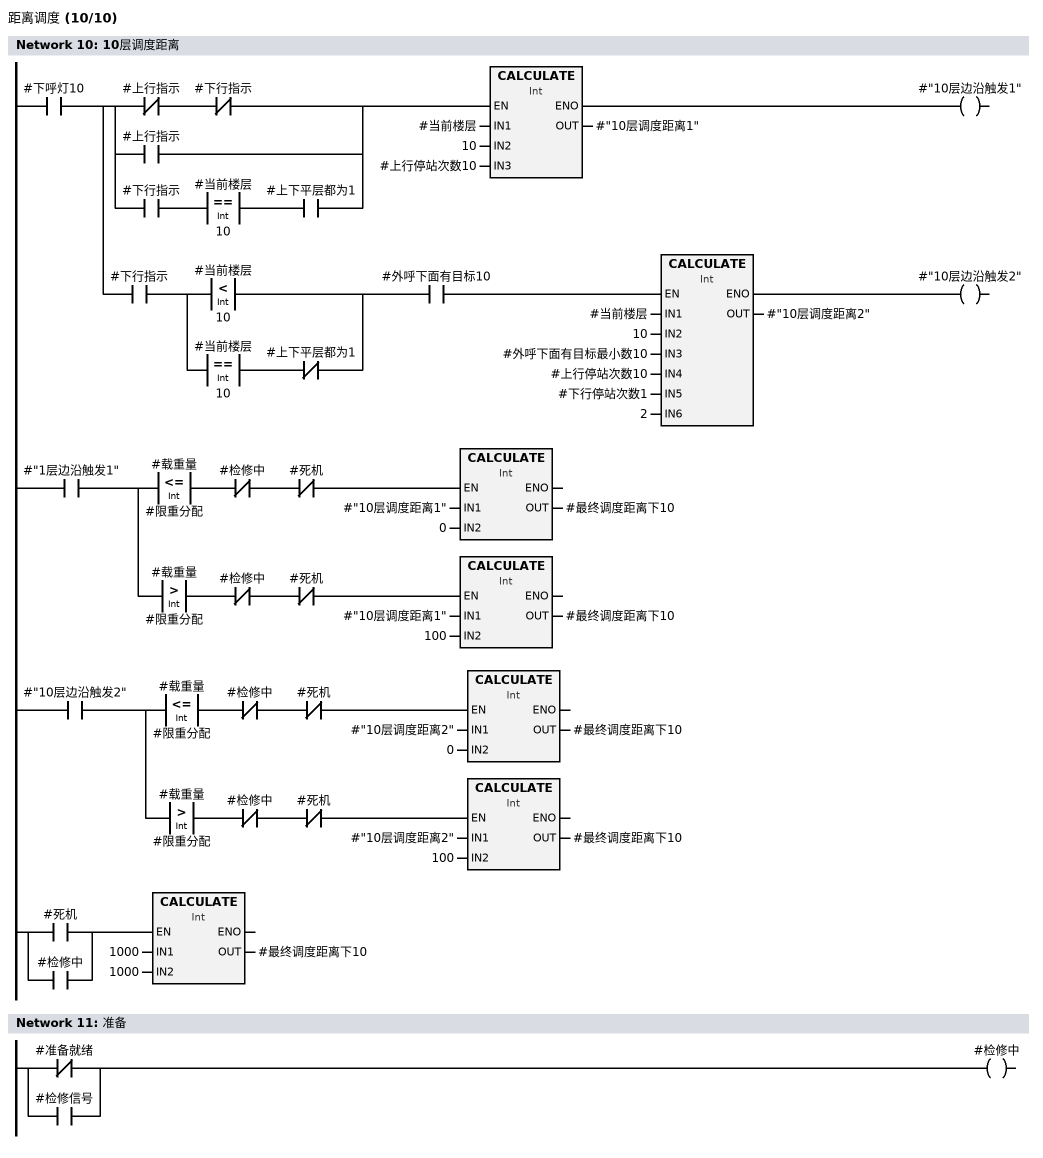
   RUNG wire#powerrail
      Contact( #下呼灯10 )
      wire#w1
      I_Contact( #上行指示 )
      I_Contact( #下行指示 )
      wire#w2
      { S7_Templates := "SrcType := Int"; S7_Expression := "ABS(IN1-IN2)+IN3+IN3" } Calculate(in1 := #当前楼层, in2 := 10, in3 := #上行停站次数10, out => #"10层调度距离1")
      Coil( #"10层边沿触发1" )
   END_RUNG
   RUNG wire#w1
      Contact( #上行指示 )
   END_RUNG wire#w2
   RUNG wire#w1
      Contact( #下行指示 )
      { S7_Templates := "SrcType := Int" } EQ_Contact(in1 := #当前楼层, in2 := 10)
      Contact( #上下平层都为1 )
   END_RUNG wire#w2
   RUNG wire#w1
      Contact( #下行指示 )
      wire#w3
      { S7_Templates := "SrcType := Int" } LT_Contact(in1 := #当前楼层, in2 := 10)
      wire#w4
      Contact( #外呼下面有目标10 )
      { S7_Templates := "SrcType := Int"; S7_Expression := "ABS(IN3+IN3-IN1-IN2)+IN4+IN4+IN5+IN5+IN6" } Calculate(in1 := #当前楼层, in2 := 10, in3 := #外呼下面有目标最小数10, in4 := #上行停站次数10, in5 := #下行停站次数1, in6 := 2, out => #"10层调度距离2")
      Coil( #"10层边沿触发2" )
   END_RUNG
   RUNG wire#w3
      { S7_Templates := "SrcType := Int" } EQ_Contact(in1 := #当前楼层, in2 := 10)
      I_Contact( #上下平层都为1 )
   END_RUNG wire#w4
   RUNG wire#powerrail
      Contact( #"1层边沿触发1" )
      wire#w5
      { S7_Templates := "SrcType := Int" } LE_Contact(in1 := #载重量, in2 := #限重分配)
      I_Contact( #检修中 )
      I_Contact( #死机 )
      { S7_Templates := "SrcType := Int"; S7_Expression := "ABS(IN1+IN2)" } Calculate(in1 := #"10层调度距离1", in2 := 0, out => #最终调度距离下10)
   END_RUNG
   RUNG wire#w5
      { S7_Templates := "SrcType := Int" } GT_Contact(in1 := #载重量, in2 := #限重分配)
      I_Contact( #检修中 )
      I_Contact( #死机 )
      { S7_Templates := "SrcType := Int"; S7_Expression := "ABS(IN1+IN2)" } Calculate(in1 := #"10层调度距离1", in2 := 100, out => #最终调度距离下10)
   END_RUNG
   RUNG wire#powerrail
      Contact( #"10层边沿触发2" )
      wire#w6
      { S7_Templates := "SrcType := Int" } LE_Contact(in1 := #载重量, in2 := #限重分配)
      I_Contact( #检修中 )
      I_Contact( #死机 )
      { S7_Templates := "SrcType := Int"; S7_Expression := "ABS(IN1+IN2)" } Calculate(in1 := #"10层调度距离2", in2 := 0, out => #最终调度距离下10)
   END_RUNG
   RUNG wire#w6
      { S7_Templates := "SrcType := Int" } GT_Contact(in1 := #载重量, in2 := #限重分配)
      I_Contact( #检修中 )
      I_Contact( #死机 )
      { S7_Templates := "SrcType := Int"; S7_Expression := "ABS(IN1+IN2)" } Calculate(in1 := #"10层调度距离2", in2 := 100, out => #最终调度距离下10)
   END_RUNG
   RUNG wire#powerrail
      Contact( #死机 )
      wire#w7
      { S7_Templates := "SrcType := Int"; S7_Expression := "ABS(IN1+IN2)" } Calculate(in1 := 1000, in2 := 1000, out => #最终调度距离下10)
   END_RUNG
   RUNG wire#powerrail
      Contact( #检修中 )
   END_RUNG wire#w7
   // the same network as SCL:
   #_w1 := #下呼灯10 AND ((NOT #上行指示 AND NOT #下行指示) OR #上行指示 OR (#下行指示 AND (#当前楼层 = 10) AND #上下平层都为1));
   IF #_w1 THEN #"10层调度距离1" := ABS(#当前楼层-10)+#上行停站次数10+#上行停站次数10; END_IF;
   #"10层边沿触发1" := #_w1;
   #_w2 := #下呼灯10 AND #下行指示 AND ((#当前楼层 < 10) OR ((#当前楼层 = 10) AND NOT #上下平层都为1)) AND #外呼下面有目标10;
   IF #_w2 THEN
       #"10层调度距离2" := ABS(#外呼下面有目标最小数10+#外呼下面有目标最小数10-#当前楼层-10)+#上行停站次数10+#上行停站次数10+#下行停站次数1+#下行停站次数1+2;
   END_IF;
   #"10层边沿触发2" := #_w2;
   IF #"1层边沿触发1" AND (#载重量 <= #限重分配) AND NOT #检修中 AND NOT #死机 THEN #最终调度距离下10 := ABS(#"10层调度距离1"+0); END_IF;
   IF #"1层边沿触发1" AND (#载重量 > #限重分配) AND NOT #检修中 AND NOT #死机 THEN #最终调度距离下10 := ABS(#"10层调度距离1"+100); END_IF;
   IF #"10层边沿触发2" AND (#载重量 <= #限重分配) AND NOT #检修中 AND NOT #死机 THEN #最终调度距离下10 := ABS(#"10层调度距离2"+0); END_IF;
   IF #"10层边沿触发2" AND (#载重量 > #限重分配) AND NOT #检修中 AND NOT #死机 THEN
       #最终调度距离下10 := ABS(#"10层调度距离2"+100);
   END_IF;
   IF #死机 OR #检修中 THEN #最终调度距离下10 := ABS(1000+1000); END_IF;
END_REGION

REGION Network 11: 准备
   RUNG wire#powerrail
      I_Contact( #准备就绪 )
      wire#w1
      Coil( #检修中 )
   END_RUNG
   RUNG wire#powerrail
      Contact( #检修信号 )
   END_RUNG wire#w1
   // the same network as SCL:
   #检修中 := NOT #准备就绪 OR #检修信号;
END_REGION
END_FUNCTION_BLOCK

FUNCTION_BLOCK "停层次数判断"   // FB33, LAD
{ S7_Optimized_Access := 'TRUE' }
VERSION : 0.1
   VAR_INPUT
      停梯截断完成开门 : Bool;
      上呼分配1 : Bool;
      上呼分配2 : Bool;
      上呼分配3 : Bool;
      上呼分配4 : Bool;
      上呼分配5 : Bool;
      上呼分配6 : Bool;
      上呼分配7 : Bool;
      上呼分配8 : Bool;
      上呼分配9 : Bool;
      下呼分配2 : Bool;
      下呼分配3 : Bool;
      下呼分配4 : Bool;
      下呼分配5 : Bool;
      下呼分配6 : Bool;
      下呼分配7 : Bool;
      下呼分配8 : Bool;
      下呼分配9 : Bool;
      下呼分配10 : Bool;
      内呼1 : Bool;
      内呼2 : Bool;
      内呼3 : Bool;
      内呼4 : Bool;
      内呼5 : Bool;
      内呼6 : Bool;
      内呼7 : Bool;
      内呼8 : Bool;
      内呼9 : Bool;
      内呼10 : Bool;
      当前楼层 : Int;
   END_VAR
   VAR_OUTPUT
      上行停站次数3 : Int;
      上行停站次数4 : Int;
      上行停站次数5 : Int;
      上行停站次数6 : Int;
      上行停站次数7 : Int;
      上行停站次数8 : Int;
      上行停站次数9 : Int;
      上行停站次数10 : Int;
      上行需折返停站次数10 : Int;
      下行停站次数1 : Int;
      下行停站次数2 : Int;
      下行停站次数3 : Int;
      下行停站次数4 : Int;
      下行停站次数5 : Int;
      下行停站次数6 : Int;
      下行停站次数7 : Int;
      下行停站次数8 : Int;
      下行需折返停站次数1 : Int;
   END_VAR
   VAR RETAIN
      IEC_Counter_0_Instance : CTUD_INT;
   END_VAR
   VAR
      上行过程需到达楼层2 : Bool;
      上行过程需到达楼层3 : Bool;
      上行过程需到达楼层4 : Bool;
      上行过程需到达楼层5 : Bool;
      上行过程需到达楼层6 : Bool;
      上行过程需到达楼层7 : Bool;
      上行过程需到达楼层8 : Bool;
      上行过程需到达楼层9 : Bool;
      上行过程需到达楼层10 : Bool;
      下行过程需到达楼层1 : Bool;
      下行过程需到达楼层2 : Bool;
      下行过程需到达楼层3 : Bool;
      下行过程需到达楼层4 : Bool;
      下行过程需到达楼层5 : Bool;
      下行过程需到达楼层6 : Bool;
      下行过程需到达楼层7 : Bool;
      下行过程需到达楼层8 : Bool;
      下行过程需到达楼层9 : Bool;
      上行计数1次1 : Int;
      上行计数1次2 : Int;
      上行计数1次3 : Int;
      上行计数1次4 : Int;
      上行计数1次5 : Int;
      上行计数1次6 : Int;
      上行计数1次7 : Int;
      上行计数1次8 : Int;
      上行计数1次9 : Int;
      上行计数1次10 : Int;
      下行计数一次1 : Int;
      下行计数一次2 : Int;
      下行计数一次3 : Int;
      下行计数一次4 : Int;
      下行计数一次5 : Int;
      下行计数一次6 : Int;
      下行计数一次7 : Int;
      下行计数一次8 : Int;
      下行计数一次9 : Int;
      下行计数一次10 : Int;
   END_VAR
   VAR RETAIN
      "IEC_Co unte r_0_Instance" : CTUD_INT;
      IEC_Counter_9_Instance : CTUD_INT;
      IEC_Counter_10_Instance : CTUD_INT;
      IEC_Counter_10_Instance上 : CTUD_INT;
      IEC_Counter_9_Instance上 : CTUD_INT;
      "IEC_Co unte r_1_Instance下" : CTUD_INT;
      "IEC_Co unte r_2_Instance下" : CTUD_INT;
      IEC_Counter_8_Instance上 : CTUD_INT;
      "IEC_Co unte r_3_Instance下" : CTUD_INT;
      IEC_Counter_7_Instance上 : CTUD_INT;
      IEC_Counter_6_Instance上 : CTUD_INT;
      IEC_Counter_5_Instance上 : CTUD_INT;
      IEC_Counter_4_Instance上 : CTUD_INT;
      IEC_Counter_3_Instance上 : CTUD_INT;
      "IEC_Co unte r_4_Instance下" : CTUD_INT;
      "IEC_Co unte r_5_Instance下" : CTUD_INT;
      "IEC_Co unte r_6_Instance下" : CTUD_INT;
      "IEC_Co unte r_7_Instance下" : CTUD_INT;
      "IEC_Co unte r_8_Instance下" : CTUD_INT;
   END_VAR
BEGIN

REGION Network 1: 上行目标转化
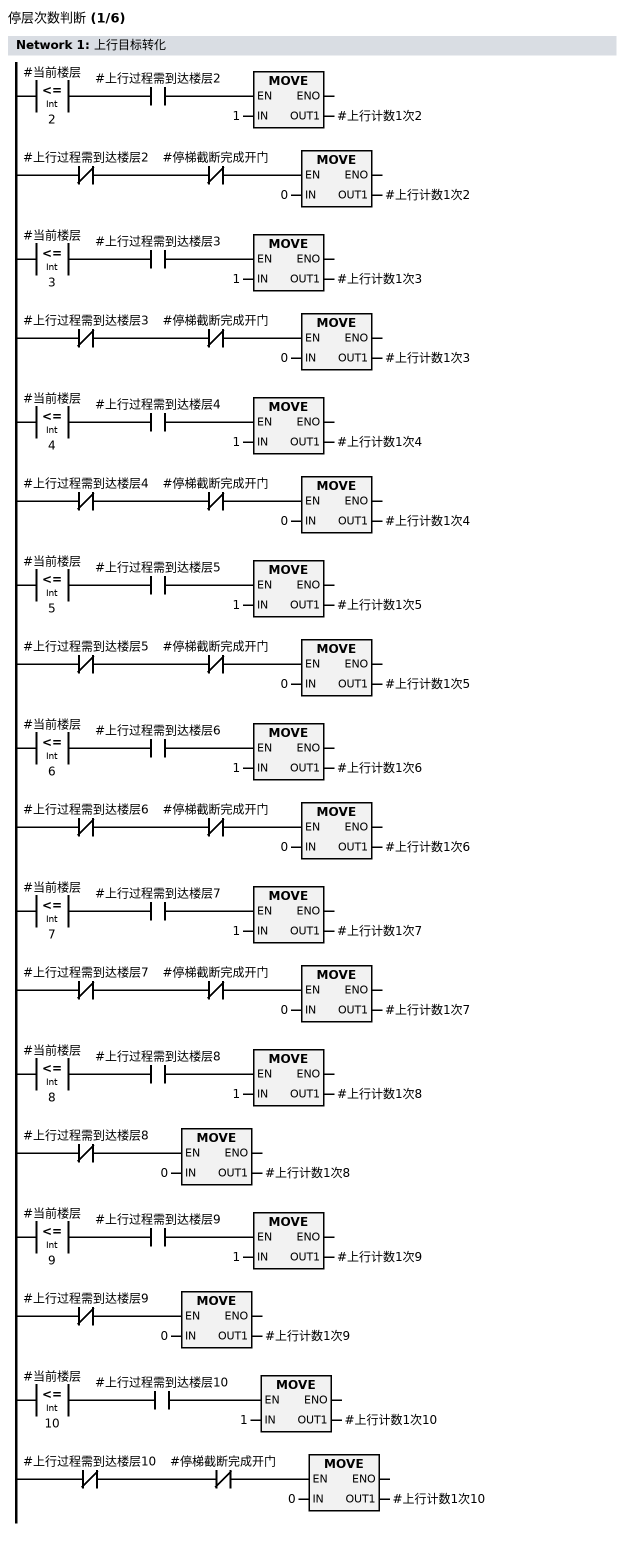
   RUNG wire#powerrail
      { S7_Templates := "SrcType := Int" } LE_Contact(in1 := #当前楼层, in2 := 2)
      Contact( #上行过程需到达楼层2 )
      Move(in := 1, out1 => #上行计数1次2)
   END_RUNG
   RUNG wire#powerrail
      I_Contact( #上行过程需到达楼层2 )
      I_Contact( #停梯截断完成开门 )
      Move(in := 0, out1 => #上行计数1次2)
   END_RUNG
   RUNG wire#powerrail
      { S7_Templates := "SrcType := Int" } LE_Contact(in1 := #当前楼层, in2 := 3)
      Contact( #上行过程需到达楼层3 )
      Move(in := 1, out1 => #上行计数1次3)
   END_RUNG
   RUNG wire#powerrail
      I_Contact( #上行过程需到达楼层3 )
      I_Contact( #停梯截断完成开门 )
      Move(in := 0, out1 => #上行计数1次3)
   END_RUNG
   RUNG wire#powerrail
      { S7_Templates := "SrcType := Int" } LE_Contact(in1 := #当前楼层, in2 := 4)
      Contact( #上行过程需到达楼层4 )
      Move(in := 1, out1 => #上行计数1次4)
   END_RUNG
   RUNG wire#powerrail
      I_Contact( #上行过程需到达楼层4 )
      I_Contact( #停梯截断完成开门 )
      Move(in := 0, out1 => #上行计数1次4)
   END_RUNG
   RUNG wire#powerrail
      { S7_Templates := "SrcType := Int" } LE_Contact(in1 := #当前楼层, in2 := 5)
      Contact( #上行过程需到达楼层5 )
      Move(in := 1, out1 => #上行计数1次5)
   END_RUNG
   RUNG wire#powerrail
      I_Contact( #上行过程需到达楼层5 )
      I_Contact( #停梯截断完成开门 )
      Move(in := 0, out1 => #上行计数1次5)
   END_RUNG
   RUNG wire#powerrail
      { S7_Templates := "SrcType := Int" } LE_Contact(in1 := #当前楼层, in2 := 6)
      Contact( #上行过程需到达楼层6 )
      Move(in := 1, out1 => #上行计数1次6)
   END_RUNG
   RUNG wire#powerrail
      I_Contact( #上行过程需到达楼层6 )
      I_Contact( #停梯截断完成开门 )
      Move(in := 0, out1 => #上行计数1次6)
   END_RUNG
   RUNG wire#powerrail
      { S7_Templates := "SrcType := Int" } LE_Contact(in1 := #当前楼层, in2 := 7)
      Contact( #上行过程需到达楼层7 )
      Move(in := 1, out1 => #上行计数1次7)
   END_RUNG
   RUNG wire#powerrail
      I_Contact( #上行过程需到达楼层7 )
      I_Contact( #停梯截断完成开门 )
      Move(in := 0, out1 => #上行计数1次7)
   END_RUNG
   RUNG wire#powerrail
      { S7_Templates := "SrcType := Int" } LE_Contact(in1 := #当前楼层, in2 := 8)
      Contact( #上行过程需到达楼层8 )
      Move(in := 1, out1 => #上行计数1次8)
   END_RUNG
   RUNG wire#powerrail
      I_Contact( #上行过程需到达楼层8 )
      Move(in := 0, out1 => #上行计数1次8)
   END_RUNG
   RUNG wire#powerrail
      { S7_Templates := "SrcType := Int" } LE_Contact(in1 := #当前楼层, in2 := 9)
      Contact( #上行过程需到达楼层9 )
      Move(in := 1, out1 => #上行计数1次9)
   END_RUNG
   RUNG wire#powerrail
      I_Contact( #上行过程需到达楼层9 )
      Move(in := 0, out1 => #上行计数1次9)
   END_RUNG
   RUNG wire#powerrail
      { S7_Templates := "SrcType := Int" } LE_Contact(in1 := #当前楼层, in2 := 10)
      Contact( #上行过程需到达楼层10 )
      Move(in := 1, out1 => #上行计数1次10)
   END_RUNG
   RUNG wire#powerrail
      I_Contact( #上行过程需到达楼层10 )
      I_Contact( #停梯截断完成开门 )
      Move(in := 0, out1 => #上行计数1次10)
   END_RUNG
   // the same network as SCL:
   IF (#当前楼层 <= 2) AND #上行过程需到达楼层2 THEN #上行计数1次2 := 1; END_IF;
   IF NOT #上行过程需到达楼层2 AND NOT #停梯截断完成开门 THEN #上行计数1次2 := 0; END_IF;
   IF (#当前楼层 <= 3) AND #上行过程需到达楼层3 THEN #上行计数1次3 := 1; END_IF;
   IF NOT #上行过程需到达楼层3 AND NOT #停梯截断完成开门 THEN #上行计数1次3 := 0; END_IF;
   IF (#当前楼层 <= 4) AND #上行过程需到达楼层4 THEN #上行计数1次4 := 1; END_IF;
   IF NOT #上行过程需到达楼层4 AND NOT #停梯截断完成开门 THEN #上行计数1次4 := 0; END_IF;
   IF (#当前楼层 <= 5) AND #上行过程需到达楼层5 THEN #上行计数1次5 := 1; END_IF;
   IF NOT #上行过程需到达楼层5 AND NOT #停梯截断完成开门 THEN #上行计数1次5 := 0; END_IF;
   IF (#当前楼层 <= 6) AND #上行过程需到达楼层6 THEN #上行计数1次6 := 1; END_IF;
   IF NOT #上行过程需到达楼层6 AND NOT #停梯截断完成开门 THEN #上行计数1次6 := 0; END_IF;
   IF (#当前楼层 <= 7) AND #上行过程需到达楼层7 THEN #上行计数1次7 := 1; END_IF;
   IF NOT #上行过程需到达楼层7 AND NOT #停梯截断完成开门 THEN #上行计数1次7 := 0; END_IF;
   IF (#当前楼层 <= 8) AND #上行过程需到达楼层8 THEN #上行计数1次8 := 1; END_IF;
   IF NOT #上行过程需到达楼层8 THEN #上行计数1次8 := 0; END_IF;
   IF (#当前楼层 <= 9) AND #上行过程需到达楼层9 THEN #上行计数1次9 := 1; END_IF;
   IF NOT #上行过程需到达楼层9 THEN #上行计数1次9 := 0; END_IF;
   IF (#当前楼层 <= 10) AND #上行过程需到达楼层10 THEN #上行计数1次10 := 1; END_IF;
   IF NOT #上行过程需到达楼层10 AND NOT #停梯截断完成开门 THEN #上行计数1次10 := 0; END_IF;
END_REGION

REGION Network 2: 上行计
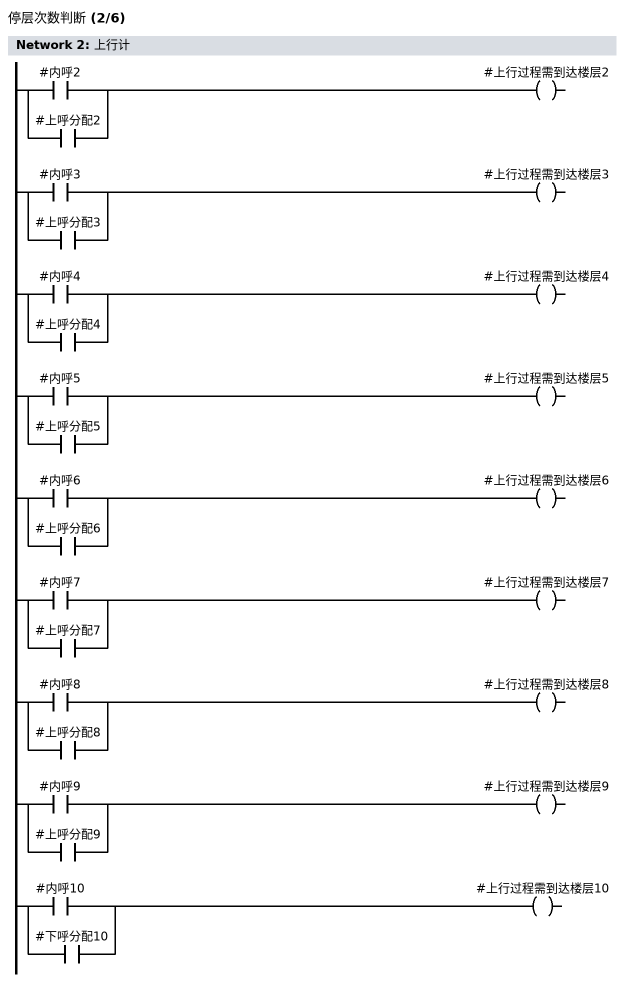
   RUNG wire#powerrail
      Contact( #内呼2 )
      wire#w1
      Coil( #上行过程需到达楼层2 )
   END_RUNG
   RUNG wire#powerrail
      Contact( #上呼分配2 )
   END_RUNG wire#w1
   RUNG wire#powerrail
      Contact( #内呼3 )
      wire#w2
      Coil( #上行过程需到达楼层3 )
   END_RUNG
   RUNG wire#powerrail
      Contact( #上呼分配3 )
   END_RUNG wire#w2
   RUNG wire#powerrail
      Contact( #内呼4 )
      wire#w3
      Coil( #上行过程需到达楼层4 )
   END_RUNG
   RUNG wire#powerrail
      Contact( #上呼分配4 )
   END_RUNG wire#w3
   RUNG wire#powerrail
      Contact( #内呼5 )
      wire#w4
      Coil( #上行过程需到达楼层5 )
   END_RUNG
   RUNG wire#powerrail
      Contact( #上呼分配5 )
   END_RUNG wire#w4
   RUNG wire#powerrail
      Contact( #内呼6 )
      wire#w5
      Coil( #上行过程需到达楼层6 )
   END_RUNG
   RUNG wire#powerrail
      Contact( #上呼分配6 )
   END_RUNG wire#w5
   RUNG wire#powerrail
      Contact( #内呼7 )
      wire#w6
      Coil( #上行过程需到达楼层7 )
   END_RUNG
   RUNG wire#powerrail
      Contact( #上呼分配7 )
   END_RUNG wire#w6
   RUNG wire#powerrail
      Contact( #内呼8 )
      wire#w7
      Coil( #上行过程需到达楼层8 )
   END_RUNG
   RUNG wire#powerrail
      Contact( #上呼分配8 )
   END_RUNG wire#w7
   RUNG wire#powerrail
      Contact( #内呼9 )
      wire#w8
      Coil( #上行过程需到达楼层9 )
   END_RUNG
   RUNG wire#powerrail
      Contact( #上呼分配9 )
   END_RUNG wire#w8
   RUNG wire#powerrail
      Contact( #内呼10 )
      wire#w9
      Coil( #上行过程需到达楼层10 )
   END_RUNG
   RUNG wire#powerrail
      Contact( #下呼分配10 )
   END_RUNG wire#w9
   // the same network as SCL:
   #上行过程需到达楼层2 := #内呼2 OR #上呼分配2;
   #上行过程需到达楼层3 := #内呼3 OR #上呼分配3;
   #上行过程需到达楼层4 := #内呼4 OR #上呼分配4;
   #上行过程需到达楼层5 := #内呼5 OR #上呼分配5;
   #上行过程需到达楼层6 := #内呼6 OR #上呼分配6;
   #上行过程需到达楼层7 := #内呼7 OR #上呼分配7;
   #上行过程需到达楼层8 := #内呼8 OR #上呼分配8;
   #上行过程需到达楼层9 := #内呼9 OR #上呼分配9;
   #上行过程需到达楼层10 := #内呼10 OR #下呼分配10;
END_REGION

REGION Network 3: 上行目标3--10层
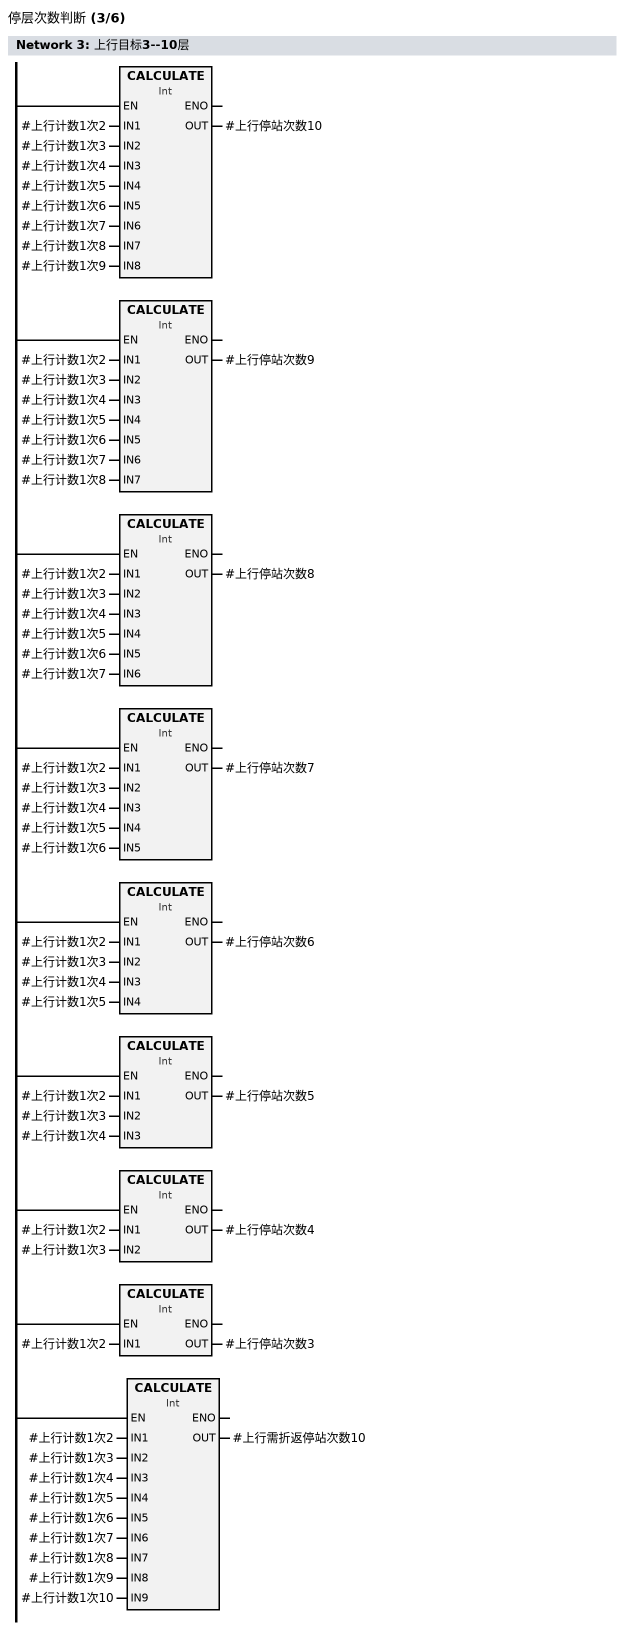
   RUNG wire#powerrail
      { S7_Templates := "SrcType := Int"; S7_Expression := "ABS(IN1+IN2+IN3+IN4+IN5+IN6+IN7+IN8)" } Calculate(in1 := #上行计数1次2, in2 := #上行计数1次3, in3 := #上行计数1次4, in4 := #上行计数1次5, in5 := #上行计数1次6, in6 := #上行计数1次7, in7 := #上行计数1次8, in8 := #上行计数1次9, out => #上行停站次数10)
   END_RUNG
   RUNG wire#powerrail
      { S7_Templates := "SrcType := Int"; S7_Expression := "ABS(IN1+IN2+IN3+IN4+IN5+IN6+IN7)" } Calculate(in1 := #上行计数1次2, in2 := #上行计数1次3, in3 := #上行计数1次4, in4 := #上行计数1次5, in5 := #上行计数1次6, in6 := #上行计数1次7, in7 := #上行计数1次8, out => #上行停站次数9)
   END_RUNG
   RUNG wire#powerrail
      { S7_Templates := "SrcType := Int"; S7_Expression := "ABS(IN1+IN2+IN3+IN4+IN5+IN6)" } Calculate(in1 := #上行计数1次2, in2 := #上行计数1次3, in3 := #上行计数1次4, in4 := #上行计数1次5, in5 := #上行计数1次6, in6 := #上行计数1次7, out => #上行停站次数8)
   END_RUNG
   RUNG wire#powerrail
      { S7_Templates := "SrcType := Int"; S7_Expression := "ABS(IN1+IN2+IN3+IN4+IN5)" } Calculate(in1 := #上行计数1次2, in2 := #上行计数1次3, in3 := #上行计数1次4, in4 := #上行计数1次5, in5 := #上行计数1次6, out => #上行停站次数7)
   END_RUNG
   RUNG wire#powerrail
      { S7_Templates := "SrcType := Int"; S7_Expression := "ABS(IN1+IN2+IN3+IN4)" } Calculate(in1 := #上行计数1次2, in2 := #上行计数1次3, in3 := #上行计数1次4, in4 := #上行计数1次5, out => #上行停站次数6)
   END_RUNG
   RUNG wire#powerrail
      { S7_Templates := "SrcType := Int"; S7_Expression := "ABS(IN1+IN2+IN3)" } Calculate(in1 := #上行计数1次2, in2 := #上行计数1次3, in3 := #上行计数1次4, out => #上行停站次数5)
   END_RUNG
   RUNG wire#powerrail
      { S7_Templates := "SrcType := Int"; S7_Expression := "ABS(IN1+IN2)" } Calculate(in1 := #上行计数1次2, in2 := #上行计数1次3, out => #上行停站次数4)
   END_RUNG
   RUNG wire#powerrail
      { S7_Templates := "SrcType := Int"; S7_Expression := "ABS(IN1)" } Calculate(in1 := #上行计数1次2, out => #上行停站次数3)
   END_RUNG
   RUNG wire#powerrail
      { S7_Templates := "SrcType := Int"; S7_Expression := "ABS(IN1+IN2+IN3+IN4+IN5+IN6+IN7+IN8+IN9)" } Calculate(in1 := #上行计数1次2, in2 := #上行计数1次3, in3 := #上行计数1次4, in4 := #上行计数1次5, in5 := #上行计数1次6, in6 := #上行计数1次7, in7 := #上行计数1次8, in8 := #上行计数1次9, in9 := #上行计数1次10, out => #上行需折返停站次数10)
   END_RUNG
   // the same network as SCL:
   #上行停站次数10 := ABS(#上行计数1次2+#上行计数1次3+#上行计数1次4+#上行计数1次5+#上行计数1次6+#上行计数1次7+#上行计数1次8+#上行计数1次9);
   #上行停站次数9 := ABS(#上行计数1次2+#上行计数1次3+#上行计数1次4+#上行计数1次5+#上行计数1次6+#上行计数1次7+#上行计数1次8);
   #上行停站次数8 := ABS(#上行计数1次2+#上行计数1次3+#上行计数1次4+#上行计数1次5+#上行计数1次6+#上行计数1次7);
   #上行停站次数7 := ABS(#上行计数1次2+#上行计数1次3+#上行计数1次4+#上行计数1次5+#上行计数1次6);
   #上行停站次数6 := ABS(#上行计数1次2+#上行计数1次3+#上行计数1次4+#上行计数1次5);
   #上行停站次数5 := ABS(#上行计数1次2+#上行计数1次3+#上行计数1次4);
   #上行停站次数4 := ABS(#上行计数1次2+#上行计数1次3);
   #上行停站次数3 := ABS(#上行计数1次2);
   #上行需折返停站次数10 := ABS(#上行计数1次2+#上行计数1次3+#上行计数1次4+#上行计数1次5+#上行计数1次6+#上行计数1次7+#上行计数1次8+#上行计数1次9+#上行计数1次10);
END_REGION

REGION Network 4: 下行目标转化
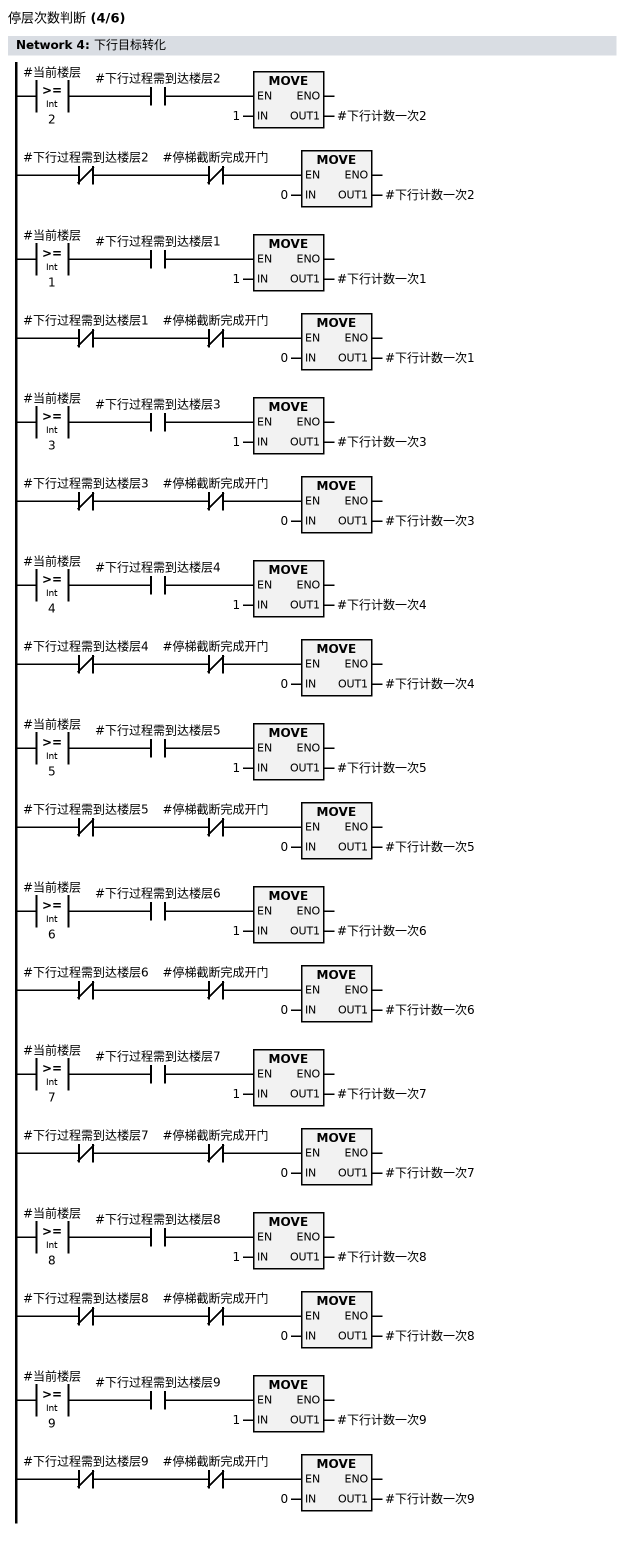
   RUNG wire#powerrail
      { S7_Templates := "SrcType := Int" } GE_Contact(in1 := #当前楼层, in2 := 2)
      Contact( #下行过程需到达楼层2 )
      Move(in := 1, out1 => #下行计数一次2)
   END_RUNG
   RUNG wire#powerrail
      I_Contact( #下行过程需到达楼层2 )
      I_Contact( #停梯截断完成开门 )
      Move(in := 0, out1 => #下行计数一次2)
   END_RUNG
   RUNG wire#powerrail
      { S7_Templates := "SrcType := Int" } GE_Contact(in1 := #当前楼层, in2 := 1)
      Contact( #下行过程需到达楼层1 )
      Move(in := 1, out1 => #下行计数一次1)
   END_RUNG
   RUNG wire#powerrail
      I_Contact( #下行过程需到达楼层1 )
      I_Contact( #停梯截断完成开门 )
      Move(in := 0, out1 => #下行计数一次1)
   END_RUNG
   RUNG wire#powerrail
      { S7_Templates := "SrcType := Int" } GE_Contact(in1 := #当前楼层, in2 := 3)
      Contact( #下行过程需到达楼层3 )
      Move(in := 1, out1 => #下行计数一次3)
   END_RUNG
   RUNG wire#powerrail
      I_Contact( #下行过程需到达楼层3 )
      I_Contact( #停梯截断完成开门 )
      Move(in := 0, out1 => #下行计数一次3)
   END_RUNG
   RUNG wire#powerrail
      { S7_Templates := "SrcType := Int" } GE_Contact(in1 := #当前楼层, in2 := 4)
      Contact( #下行过程需到达楼层4 )
      Move(in := 1, out1 => #下行计数一次4)
   END_RUNG
   RUNG wire#powerrail
      I_Contact( #下行过程需到达楼层4 )
      I_Contact( #停梯截断完成开门 )
      Move(in := 0, out1 => #下行计数一次4)
   END_RUNG
   RUNG wire#powerrail
      { S7_Templates := "SrcType := Int" } GE_Contact(in1 := #当前楼层, in2 := 5)
      Contact( #下行过程需到达楼层5 )
      Move(in := 1, out1 => #下行计数一次5)
   END_RUNG
   RUNG wire#powerrail
      I_Contact( #下行过程需到达楼层5 )
      I_Contact( #停梯截断完成开门 )
      Move(in := 0, out1 => #下行计数一次5)
   END_RUNG
   RUNG wire#powerrail
      { S7_Templates := "SrcType := Int" } GE_Contact(in1 := #当前楼层, in2 := 6)
      Contact( #下行过程需到达楼层6 )
      Move(in := 1, out1 => #下行计数一次6)
   END_RUNG
   RUNG wire#powerrail
      I_Contact( #下行过程需到达楼层6 )
      I_Contact( #停梯截断完成开门 )
      Move(in := 0, out1 => #下行计数一次6)
   END_RUNG
   RUNG wire#powerrail
      { S7_Templates := "SrcType := Int" } GE_Contact(in1 := #当前楼层, in2 := 7)
      Contact( #下行过程需到达楼层7 )
      Move(in := 1, out1 => #下行计数一次7)
   END_RUNG
   RUNG wire#powerrail
      I_Contact( #下行过程需到达楼层7 )
      I_Contact( #停梯截断完成开门 )
      Move(in := 0, out1 => #下行计数一次7)
   END_RUNG
   RUNG wire#powerrail
      { S7_Templates := "SrcType := Int" } GE_Contact(in1 := #当前楼层, in2 := 8)
      Contact( #下行过程需到达楼层8 )
      Move(in := 1, out1 => #下行计数一次8)
   END_RUNG
   RUNG wire#powerrail
      I_Contact( #下行过程需到达楼层8 )
      I_Contact( #停梯截断完成开门 )
      Move(in := 0, out1 => #下行计数一次8)
   END_RUNG
   RUNG wire#powerrail
      { S7_Templates := "SrcType := Int" } GE_Contact(in1 := #当前楼层, in2 := 9)
      Contact( #下行过程需到达楼层9 )
      Move(in := 1, out1 => #下行计数一次9)
   END_RUNG
   RUNG wire#powerrail
      I_Contact( #下行过程需到达楼层9 )
      I_Contact( #停梯截断完成开门 )
      Move(in := 0, out1 => #下行计数一次9)
   END_RUNG
   // the same network as SCL:
   IF (#当前楼层 >= 2) AND #下行过程需到达楼层2 THEN #下行计数一次2 := 1; END_IF;
   IF NOT #下行过程需到达楼层2 AND NOT #停梯截断完成开门 THEN #下行计数一次2 := 0; END_IF;
   IF (#当前楼层 >= 1) AND #下行过程需到达楼层1 THEN #下行计数一次1 := 1; END_IF;
   IF NOT #下行过程需到达楼层1 AND NOT #停梯截断完成开门 THEN #下行计数一次1 := 0; END_IF;
   IF (#当前楼层 >= 3) AND #下行过程需到达楼层3 THEN #下行计数一次3 := 1; END_IF;
   IF NOT #下行过程需到达楼层3 AND NOT #停梯截断完成开门 THEN #下行计数一次3 := 0; END_IF;
   IF (#当前楼层 >= 4) AND #下行过程需到达楼层4 THEN #下行计数一次4 := 1; END_IF;
   IF NOT #下行过程需到达楼层4 AND NOT #停梯截断完成开门 THEN #下行计数一次4 := 0; END_IF;
   IF (#当前楼层 >= 5) AND #下行过程需到达楼层5 THEN #下行计数一次5 := 1; END_IF;
   IF NOT #下行过程需到达楼层5 AND NOT #停梯截断完成开门 THEN #下行计数一次5 := 0; END_IF;
   IF (#当前楼层 >= 6) AND #下行过程需到达楼层6 THEN #下行计数一次6 := 1; END_IF;
   IF NOT #下行过程需到达楼层6 AND NOT #停梯截断完成开门 THEN #下行计数一次6 := 0; END_IF;
   IF (#当前楼层 >= 7) AND #下行过程需到达楼层7 THEN #下行计数一次7 := 1; END_IF;
   IF NOT #下行过程需到达楼层7 AND NOT #停梯截断完成开门 THEN #下行计数一次7 := 0; END_IF;
   IF (#当前楼层 >= 8) AND #下行过程需到达楼层8 THEN #下行计数一次8 := 1; END_IF;
   IF NOT #下行过程需到达楼层8 AND NOT #停梯截断完成开门 THEN #下行计数一次8 := 0; END_IF;
   IF (#当前楼层 >= 9) AND #下行过程需到达楼层9 THEN #下行计数一次9 := 1; END_IF;
   IF NOT #下行过程需到达楼层9 AND NOT #停梯截断完成开门 THEN #下行计数一次9 := 0; END_IF;
END_REGION

REGION Network 5: 下行计
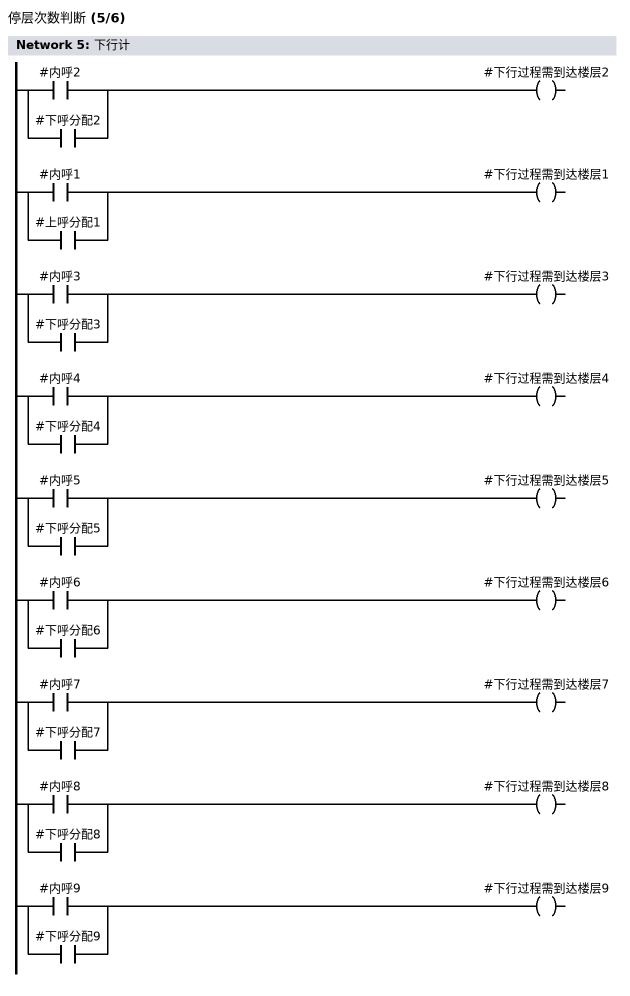
   RUNG wire#powerrail
      Contact( #内呼2 )
      wire#w1
      Coil( #下行过程需到达楼层2 )
   END_RUNG
   RUNG wire#powerrail
      Contact( #下呼分配2 )
   END_RUNG wire#w1
   RUNG wire#powerrail
      Contact( #内呼1 )
      wire#w2
      Coil( #下行过程需到达楼层1 )
   END_RUNG
   RUNG wire#powerrail
      Contact( #上呼分配1 )
   END_RUNG wire#w2
   RUNG wire#powerrail
      Contact( #内呼3 )
      wire#w3
      Coil( #下行过程需到达楼层3 )
   END_RUNG
   RUNG wire#powerrail
      Contact( #下呼分配3 )
   END_RUNG wire#w3
   RUNG wire#powerrail
      Contact( #内呼4 )
      wire#w4
      Coil( #下行过程需到达楼层4 )
   END_RUNG
   RUNG wire#powerrail
      Contact( #下呼分配4 )
   END_RUNG wire#w4
   RUNG wire#powerrail
      Contact( #内呼5 )
      wire#w5
      Coil( #下行过程需到达楼层5 )
   END_RUNG
   RUNG wire#powerrail
      Contact( #下呼分配5 )
   END_RUNG wire#w5
   RUNG wire#powerrail
      Contact( #内呼6 )
      wire#w6
      Coil( #下行过程需到达楼层6 )
   END_RUNG
   RUNG wire#powerrail
      Contact( #下呼分配6 )
   END_RUNG wire#w6
   RUNG wire#powerrail
      Contact( #内呼7 )
      wire#w7
      Coil( #下行过程需到达楼层7 )
   END_RUNG
   RUNG wire#powerrail
      Contact( #下呼分配7 )
   END_RUNG wire#w7
   RUNG wire#powerrail
      Contact( #内呼8 )
      wire#w8
      Coil( #下行过程需到达楼层8 )
   END_RUNG
   RUNG wire#powerrail
      Contact( #下呼分配8 )
   END_RUNG wire#w8
   RUNG wire#powerrail
      Contact( #内呼9 )
      wire#w9
      Coil( #下行过程需到达楼层9 )
   END_RUNG
   RUNG wire#powerrail
      Contact( #下呼分配9 )
   END_RUNG wire#w9
   // the same network as SCL:
   #下行过程需到达楼层2 := #内呼2 OR #下呼分配2;
   #下行过程需到达楼层1 := #内呼1 OR #上呼分配1;
   #下行过程需到达楼层3 := #内呼3 OR #下呼分配3;
   #下行过程需到达楼层4 := #内呼4 OR #下呼分配4;
   #下行过程需到达楼层5 := #内呼5 OR #下呼分配5;
   #下行过程需到达楼层6 := #内呼6 OR #下呼分配6;
   #下行过程需到达楼层7 := #内呼7 OR #下呼分配7;
   #下行过程需到达楼层8 := #内呼8 OR #下呼分配8;
   #下行过程需到达楼层9 := #内呼9 OR #下呼分配9;
END_REGION

REGION Network 6: 下行目标1--8层
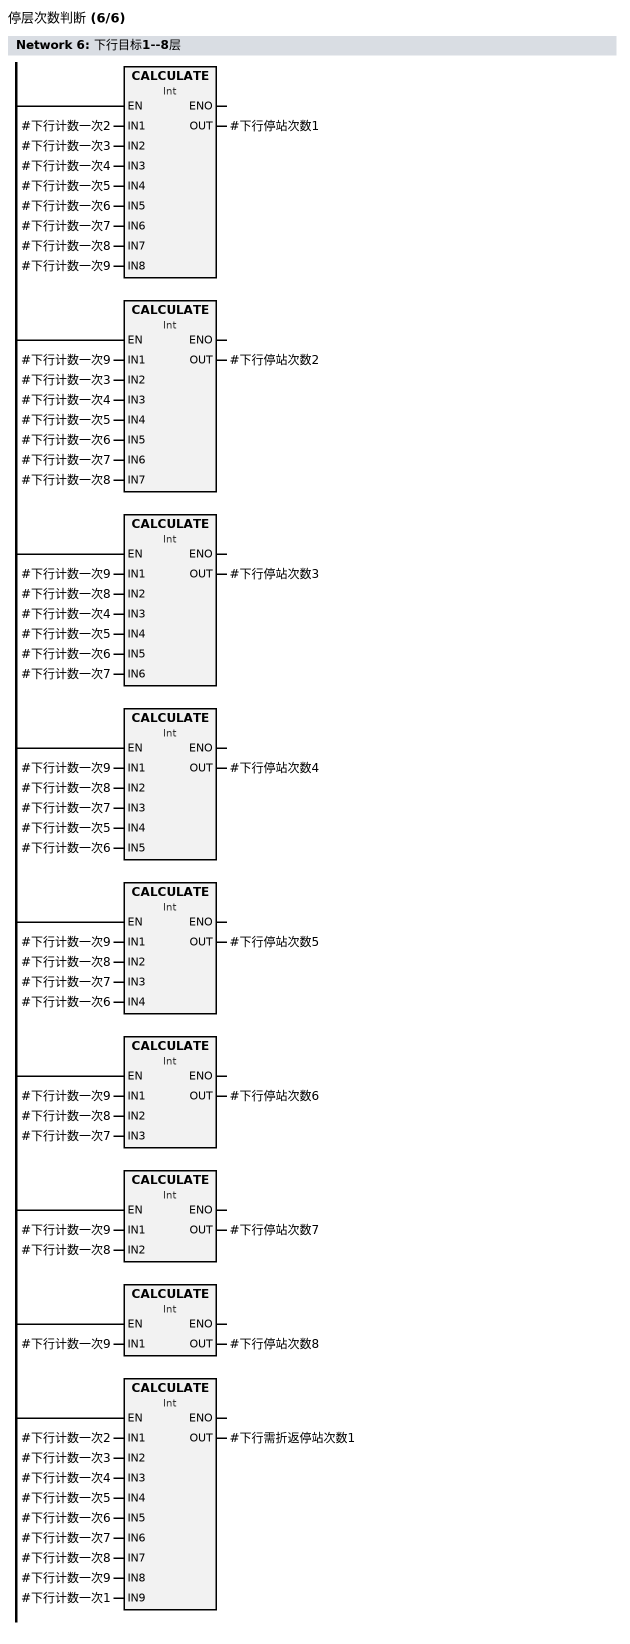
   RUNG wire#powerrail
      { S7_Templates := "SrcType := Int"; S7_Expression := "ABS(IN1+IN2+IN3+IN4+IN5+IN6+IN7+IN8)" } Calculate(in1 := #下行计数一次2, in2 := #下行计数一次3, in3 := #下行计数一次4, in4 := #下行计数一次5, in5 := #下行计数一次6, in6 := #下行计数一次7, in7 := #下行计数一次8, in8 := #下行计数一次9, out => #下行停站次数1)
   END_RUNG
   RUNG wire#powerrail
      { S7_Templates := "SrcType := Int"; S7_Expression := "ABS(IN1+IN2+IN3+IN4+IN5+IN6+IN7)" } Calculate(in1 := #下行计数一次9, in2 := #下行计数一次3, in3 := #下行计数一次4, in4 := #下行计数一次5, in5 := #下行计数一次6, in6 := #下行计数一次7, in7 := #下行计数一次8, out => #下行停站次数2)
   END_RUNG
   RUNG wire#powerrail
      { S7_Templates := "SrcType := Int"; S7_Expression := "ABS(IN1+IN2+IN3+IN4+IN5+IN6)" } Calculate(in1 := #下行计数一次9, in2 := #下行计数一次8, in3 := #下行计数一次4, in4 := #下行计数一次5, in5 := #下行计数一次6, in6 := #下行计数一次7, out => #下行停站次数3)
   END_RUNG
   RUNG wire#powerrail
      { S7_Templates := "SrcType := Int"; S7_Expression := "ABS(IN1+IN2+IN3+IN4+IN5)" } Calculate(in1 := #下行计数一次9, in2 := #下行计数一次8, in3 := #下行计数一次7, in4 := #下行计数一次5, in5 := #下行计数一次6, out => #下行停站次数4)
   END_RUNG
   RUNG wire#powerrail
      { S7_Templates := "SrcType := Int"; S7_Expression := "ABS(IN1+IN2+IN3+IN4)" } Calculate(in1 := #下行计数一次9, in2 := #下行计数一次8, in3 := #下行计数一次7, in4 := #下行计数一次6, out => #下行停站次数5)
   END_RUNG
   RUNG wire#powerrail
      { S7_Templates := "SrcType := Int"; S7_Expression := "ABS(IN1+IN2+IN3)" } Calculate(in1 := #下行计数一次9, in2 := #下行计数一次8, in3 := #下行计数一次7, out => #下行停站次数6)
   END_RUNG
   RUNG wire#powerrail
      { S7_Templates := "SrcType := Int"; S7_Expression := "ABS(IN1+IN2)" } Calculate(in1 := #下行计数一次9, in2 := #下行计数一次8, out => #下行停站次数7)
   END_RUNG
   RUNG wire#powerrail
      { S7_Templates := "SrcType := Int"; S7_Expression := "ABS(IN1)" } Calculate(in1 := #下行计数一次9, out => #下行停站次数8)
   END_RUNG
   RUNG wire#powerrail
      { S7_Templates := "SrcType := Int"; S7_Expression := "ABS(IN1+IN2+IN3+IN4+IN5+IN6+IN7+IN8+IN9)" } Calculate(in1 := #下行计数一次2, in2 := #下行计数一次3, in3 := #下行计数一次4, in4 := #下行计数一次5, in5 := #下行计数一次6, in6 := #下行计数一次7, in7 := #下行计数一次8, in8 := #下行计数一次9, in9 := #下行计数一次1, out => #下行需折返停站次数1)
   END_RUNG
   // the same network as SCL:
   #下行停站次数1 := ABS(#下行计数一次2+#下行计数一次3+#下行计数一次4+#下行计数一次5+#下行计数一次6+#下行计数一次7+#下行计数一次8+#下行计数一次9);
   #下行停站次数2 := ABS(#下行计数一次9+#下行计数一次3+#下行计数一次4+#下行计数一次5+#下行计数一次6+#下行计数一次7+#下行计数一次8);
   #下行停站次数3 := ABS(#下行计数一次9+#下行计数一次8+#下行计数一次4+#下行计数一次5+#下行计数一次6+#下行计数一次7);
   #下行停站次数4 := ABS(#下行计数一次9+#下行计数一次8+#下行计数一次7+#下行计数一次5+#下行计数一次6);
   #下行停站次数5 := ABS(#下行计数一次9+#下行计数一次8+#下行计数一次7+#下行计数一次6);
   #下行停站次数6 := ABS(#下行计数一次9+#下行计数一次8+#下行计数一次7);
   #下行停站次数7 := ABS(#下行计数一次9+#下行计数一次8);
   #下行停站次数8 := ABS(#下行计数一次9);
   #下行需折返停站次数1 := ABS(#下行计数一次2+#下行计数一次3+#下行计数一次4+#下行计数一次5+#下行计数一次6+#下行计数一次7+#下行计数一次8+#下行计数一次9+#下行计数一次1);
END_REGION
END_FUNCTION_BLOCK

FUNCTION_BLOCK "初始化"   // FB36, LAD
{ S7_Optimized_Access := 'TRUE' }
VERSION : 0.1
   VAR_INPUT
      自动运行信号 : Bool;
      初始化方向上行 : Bool;
      "1号梯上端站第1限位" : Bool;
      "1号梯下端站第1限位" : Bool;
      初始化方向下行 : Bool;
      当前楼层数 : Int;
      初始化楼层数 : Int := 1;
      检修信号 : Bool;
      高速延时 : Time;
      是否高速 : Bool;
      两平层同时为1 : Bool;
      检修楼层数 : Int;
   END_VAR
   VAR_OUTPUT
      初始化上行接触器 : Bool;
      初始化下行接触器 : Bool;
      "1号梯电机启动信号" : Bool;
      初始化低速运行 : Bool;
      准备就绪信号 : Bool;
      是否到达端限 : Bool;
      初始化将要停梯 : Bool;
      到达初始化楼层 : Bool;
      初始化高速运行 : Bool;
      "1号梯上行指示" : Bool;
      "1号梯下行指示" : Bool;
   END_VAR
   VAR
      检修方向上行 : Bool;
      检修方向下行 : Bool;
      完成过一次初始化 : Bool;
      现在在检修 : Bool;
      连接1 : Bool;
      连接2 : Bool;
      连接3 : Bool;
      连接4 : Bool;
      连接5 : Bool;
      连接6 : Bool;
      连接7 : Bool;
      连接8 : Bool;
      连接9 : Bool;
      "延迟 制动" : TON_TIME;
      稍后 : TON_TIME;
      确保初始化停稳 : TON_TIME;
      IEC_Timer_0_Instance : TON_TIME;
      IEC_Timer_0_Instance_1 : TON_TIME;
      IEC_Timer_0_Instance_2 : TON_TIME;
      记录检修 : Bool;
      中间连接 : Bool;
      检修完成 : Bool;
      "稍 后" : TON_TIME;
   END_VAR
   VAR RETAIN
      IEC_Counter_0_Instance : CTU_INT;
   END_VAR
   VAR
      IEC_Timer_0_Instance_3 : TP_TIME;
      IEC_Timer_0_Instance_4 : TON_TIME;
   END_VAR
   VAR RETAIN
      IEC_Counter_0_Instance_1 : CTU_INT;
   END_VAR
   VAR
      IEC_Timer_0_Instance_5 : TP_TIME;
      IEC_Timer_0_Instance_6 : TP_TIME;
      IEC_Timer_0_Instance_7 : TP_TIME;
      IEC_Timer_0_Instance_8 : TON_TIME;
      IEC_Timer_0_Instance_9 : TON_TIME;
      IEC_Timer_0_Instance_10 : TON_TIME;
   END_VAR
   VAR_TEMP   // added for the SCL form of the ladder/FBD networks
      _w1 : Bool;
      _w2 : Bool;
      _w3 : Bool;
      _w4 : Bool;
      _w5 : Bool;
      _w6 : Bool;
   END_VAR
BEGIN

REGION Network 1: 启动信号
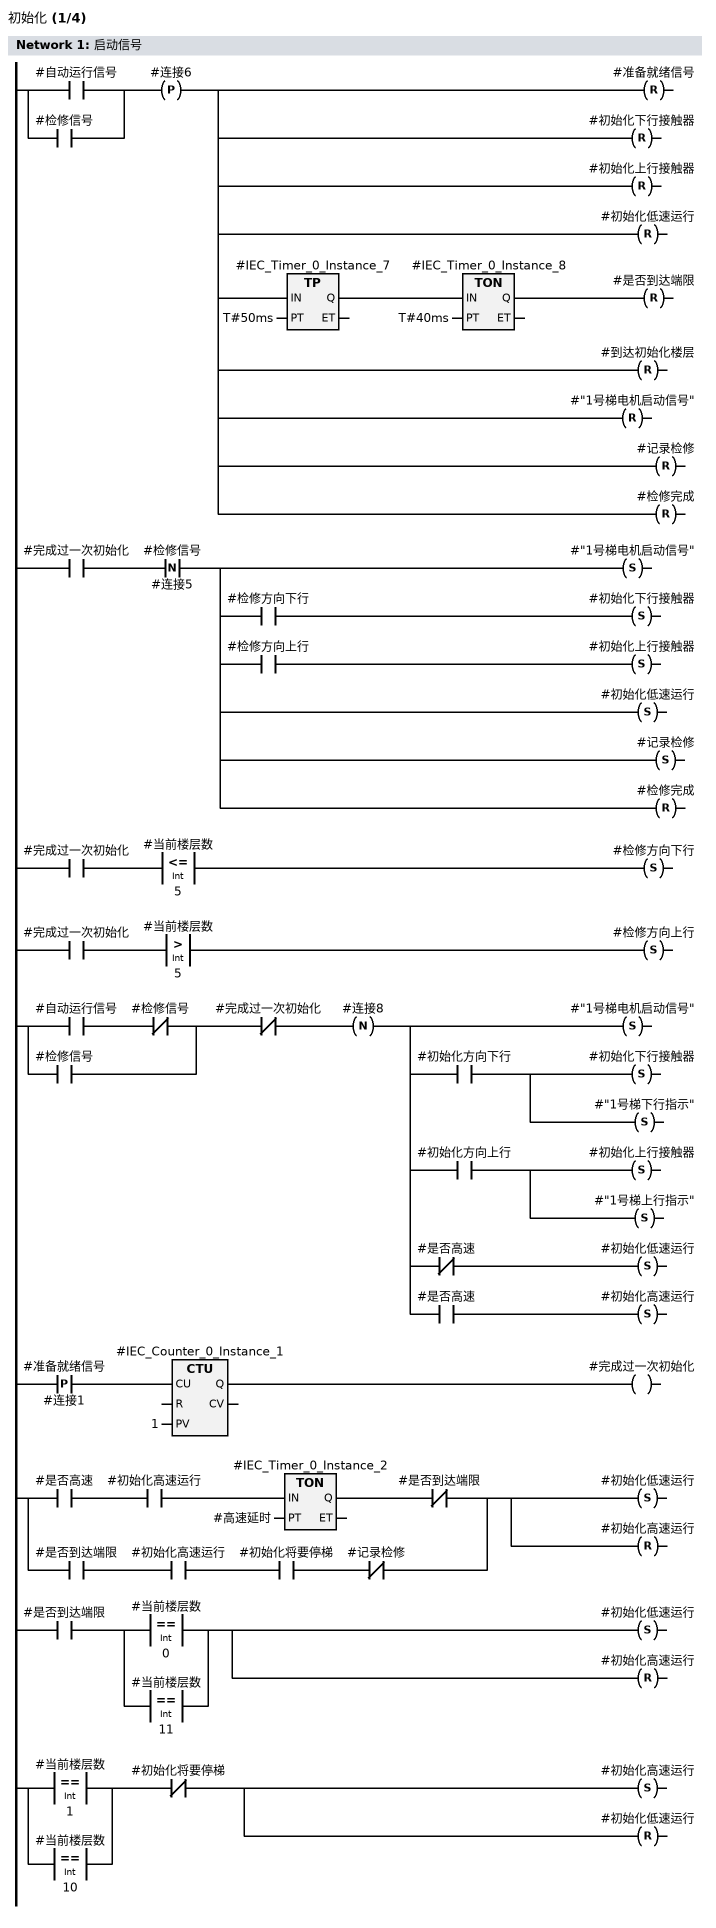
   #_w1 := #自动运行信号 OR #检修信号;
   #_w2 := #_w1 AND NOT #连接6;   // rising edge
   #连接6 := #_w1;
   IF #_w2 THEN
       #准备就绪信号 := FALSE;
       #初始化下行接触器 := FALSE;
       #初始化上行接触器 := FALSE;
       #初始化低速运行 := FALSE;
   END_IF;
   #IEC_Timer_0_Instance_7(IN := #_w2, PT := T#50ms);   // TP
   #IEC_Timer_0_Instance_8(IN := #IEC_Timer_0_Instance_7.Q, PT := T#40ms);   // TON
   IF #IEC_Timer_0_Instance_8.Q THEN #是否到达端限 := FALSE; END_IF;
   IF #_w2 THEN
       #到达初始化楼层 := FALSE;
       #"1号梯电机启动信号" := FALSE;
       #记录检修 := FALSE;
       #检修完成 := FALSE;
   END_IF;
   #_w3 := #完成过一次初始化 AND NOT #检修信号 AND #连接5;   // falling edge of #检修信号
   #连接5 := #检修信号;
   IF #_w3 THEN #"1号梯电机启动信号" := TRUE; END_IF;
   IF #_w3 AND #检修方向下行 THEN #初始化下行接触器 := TRUE; END_IF;
   IF #_w3 AND #检修方向上行 THEN #初始化上行接触器 := TRUE; END_IF;
   IF #_w3 THEN
       #初始化低速运行 := TRUE;
       #记录检修 := TRUE;
       #检修完成 := FALSE;
   END_IF;
   IF #完成过一次初始化 AND (#当前楼层数 <= 5) THEN #检修方向下行 := TRUE; END_IF;
   IF #完成过一次初始化 AND (#当前楼层数 > 5) THEN #检修方向上行 := TRUE; END_IF;
   #_w4 := ((#自动运行信号 AND NOT #检修信号) OR #检修信号) AND NOT #完成过一次初始化;
   #_w5 := NOT #_w4 AND #连接8;   // falling edge
   #连接8 := #_w4;
   IF #_w5 THEN #"1号梯电机启动信号" := TRUE; END_IF;
   IF #_w5 AND #初始化方向下行 THEN
       #初始化下行接触器 := TRUE;
       #"1号梯下行指示" := TRUE;
   END_IF;
   IF #_w5 AND #初始化方向上行 THEN
       #初始化上行接触器 := TRUE;
       #"1号梯上行指示" := TRUE;
   END_IF;
   IF #_w5 AND NOT #是否高速 THEN #初始化低速运行 := TRUE; END_IF;
   IF #_w5 AND #是否高速 THEN #初始化高速运行 := TRUE; END_IF;
   #_w6 := #准备就绪信号 AND NOT #连接1;   // rising edge of #准备就绪信号
   #连接1 := #准备就绪信号;
   #IEC_Counter_0_Instance_1(CU := #_w6, PV := 1);   // CTU
   #完成过一次初始化 := #IEC_Counter_0_Instance_1.Q;
   #IEC_Timer_0_Instance_2(IN := #是否高速 AND #初始化高速运行, PT := #高速延时);   // TON
   IF (#IEC_Timer_0_Instance_2.Q AND NOT #是否到达端限) OR (#是否到达端限 AND #初始化高速运行 AND #初始化将要停梯 AND NOT #记录检修) THEN
       #初始化低速运行 := TRUE;
       #初始化高速运行 := FALSE;
   END_IF;
   IF #是否到达端限 AND ((#当前楼层数 = 0) OR (#当前楼层数 = 11)) THEN
       #初始化低速运行 := TRUE;
       #初始化高速运行 := FALSE;
   END_IF;
   IF ((#当前楼层数 = 1) OR (#当前楼层数 = 10)) AND NOT #初始化将要停梯 THEN
       #初始化高速运行 := TRUE;
       #初始化低速运行 := FALSE;
   END_IF;
END_REGION

REGION Network 2: 到达端限，开始计算楼层
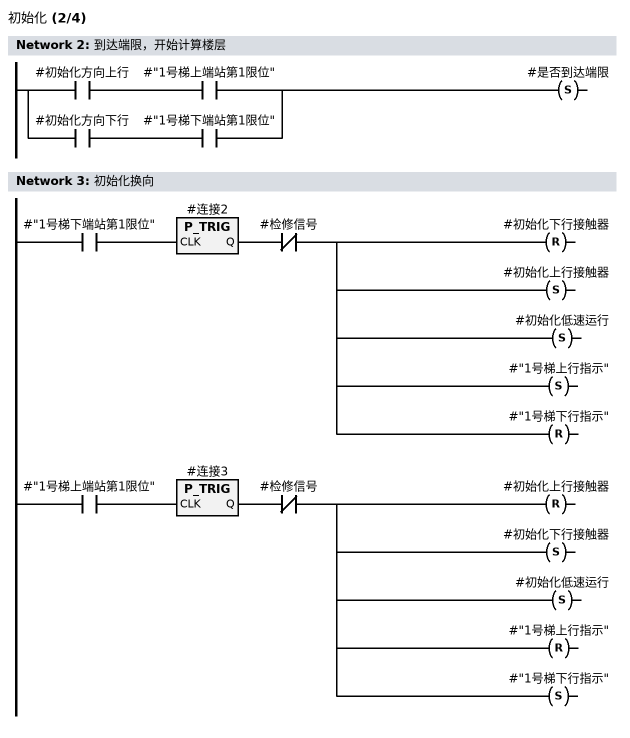
   RUNG wire#powerrail
      Contact( #初始化方向上行 )
      Contact( #"1号梯上端站第1限位" )
      wire#w1
      S_Coil( #是否到达端限 )
   END_RUNG
   RUNG wire#powerrail
      Contact( #初始化方向下行 )
      Contact( #"1号梯下端站第1限位" )
   END_RUNG wire#w1
   // the same network as SCL:
   IF (#初始化方向上行 AND #"1号梯上端站第1限位") OR (#初始化方向下行 AND #"1号梯下端站第1限位") THEN #是否到达端限 := TRUE; END_IF;
END_REGION

REGION Network 3: 初始化换向
   RUNG wire#powerrail
      Contact( #"1号梯下端站第1限位" )
      P_Trig( #连接2 )
      I_Contact( #检修信号 )
      wire#w1
      R_Coil( #初始化下行接触器 )
   END_RUNG
   RUNG wire#w1
      S_Coil( #初始化上行接触器 )
   END_RUNG
   RUNG wire#w1
      S_Coil( #初始化低速运行 )
   END_RUNG
   RUNG wire#w1
      S_Coil( #"1号梯上行指示" )
   END_RUNG
   RUNG wire#w1
      R_Coil( #"1号梯下行指示" )
   END_RUNG
   RUNG wire#powerrail
      Contact( #"1号梯上端站第1限位" )
      P_Trig( #连接3 )
      I_Contact( #检修信号 )
      wire#w2
      R_Coil( #初始化上行接触器 )
   END_RUNG
   RUNG wire#w2
      S_Coil( #初始化下行接触器 )
   END_RUNG
   RUNG wire#w2
      S_Coil( #初始化低速运行 )
   END_RUNG
   RUNG wire#w2
      R_Coil( #"1号梯上行指示" )
   END_RUNG
   RUNG wire#w2
      S_Coil( #"1号梯下行指示" )
   END_RUNG
   // the same network as SCL:
   #_w1 := #"1号梯下端站第1限位" AND NOT #连接2;   // rising edge
   #连接2 := #"1号梯下端站第1限位";
   IF #_w1 AND NOT #检修信号 THEN
       #初始化下行接触器 := FALSE;
       #初始化上行接触器 := TRUE;
       #初始化低速运行 := TRUE;
       #"1号梯上行指示" := TRUE;
       #"1号梯下行指示" := FALSE;
   END_IF;
   #_w2 := #"1号梯上端站第1限位" AND NOT #连接3;   // rising edge
   #连接3 := #"1号梯上端站第1限位";
   IF #_w2 AND NOT #检修信号 THEN
       #初始化上行接触器 := FALSE;
       #初始化下行接触器 := TRUE;
       #初始化低速运行 := TRUE;
       #"1号梯上行指示" := FALSE;
       #"1号梯下行指示" := TRUE;
   END_IF;
END_REGION

REGION Network 4: 初始化结束停车
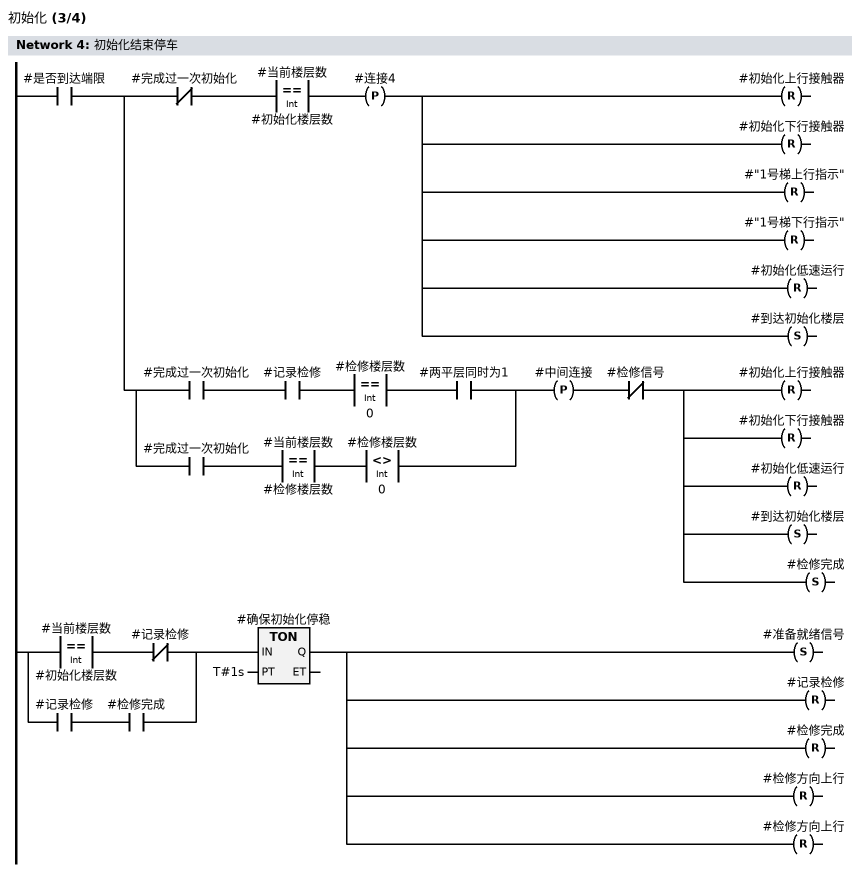
   #_w1 := #是否到达端限 AND NOT #完成过一次初始化 AND (#当前楼层数 = #初始化楼层数);
   #_w2 := #_w1 AND NOT #连接4;   // rising edge
   #连接4 := #_w1;
   IF #_w2 THEN
       #初始化上行接触器 := FALSE;
       #初始化下行接触器 := FALSE;
       #"1号梯上行指示" := FALSE;
       #"1号梯下行指示" := FALSE;
       #初始化低速运行 := FALSE;
       #到达初始化楼层 := TRUE;
   END_IF;
   #_w3 := #是否到达端限 AND ((#完成过一次初始化 AND #记录检修 AND (#检修楼层数 = 0) AND #两平层同时为1) OR (#完成过一次初始化 AND (#当前楼层数 = #检修楼层数) AND (#检修楼层数 <> 0)));
   #_w4 := #_w3 AND NOT #中间连接;   // rising edge
   #中间连接 := #_w3;
   IF #_w4 AND NOT #检修信号 THEN
       #初始化上行接触器 := FALSE;
       #初始化下行接触器 := FALSE;
       #初始化低速运行 := FALSE;
       #到达初始化楼层 := TRUE;
       #检修完成 := TRUE;
   END_IF;
   #确保初始化停稳(IN := ((#当前楼层数 = #初始化楼层数) AND NOT #记录检修) OR (#记录检修 AND #检修完成), PT := T#1s);   // TON
   IF #确保初始化停稳.Q THEN
       #准备就绪信号 := TRUE;
       #记录检修 := FALSE;
       #检修完成 := FALSE;
       #检修方向上行 := FALSE;
       #检修方向上行 := FALSE;
   END_IF;
END_REGION

REGION Network 5: 初始化刹车
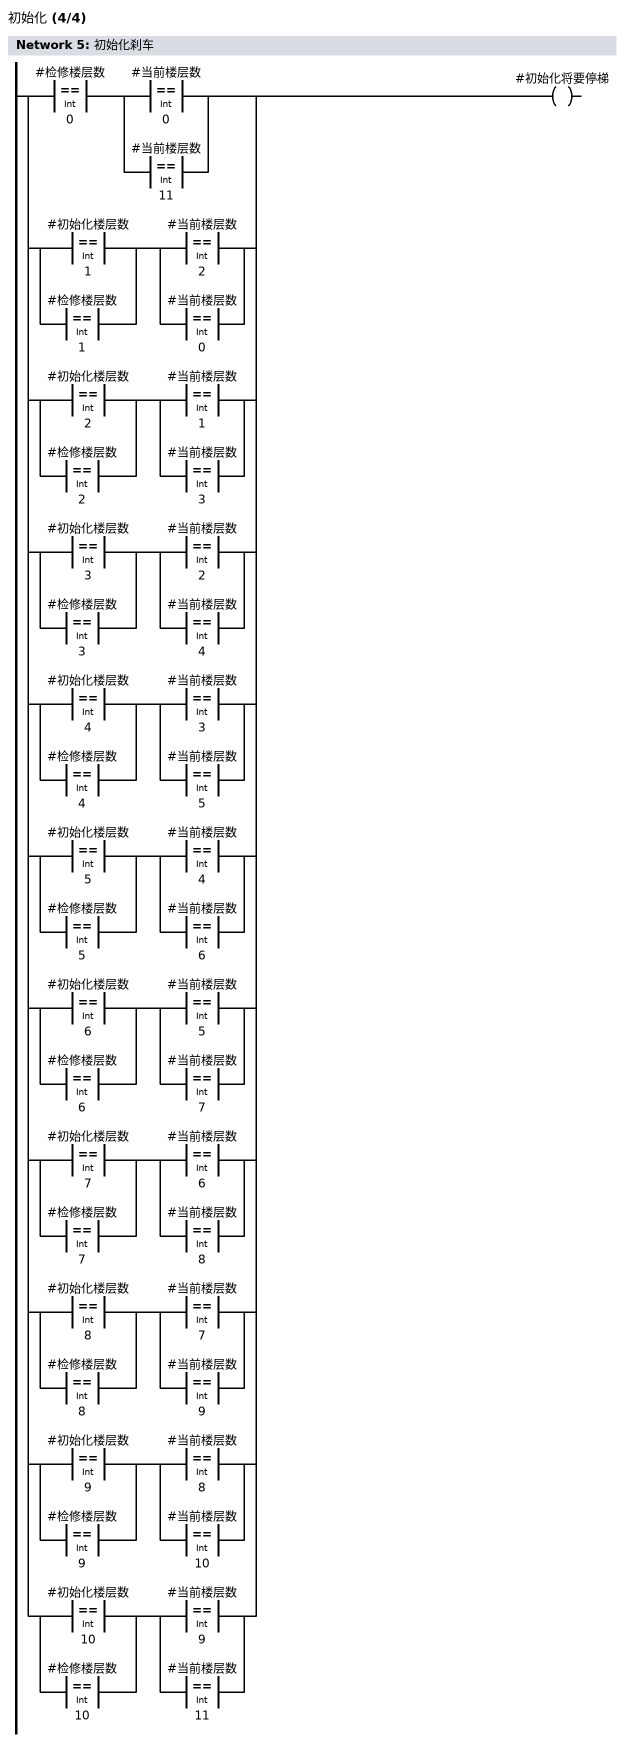
   RUNG wire#powerrail
      { S7_Templates := "SrcType := Int" } EQ_Contact(in1 := #检修楼层数, in2 := 0)
      wire#w1
      { S7_Templates := "SrcType := Int" } EQ_Contact(in1 := #当前楼层数, in2 := 0)
      wire#w2
      Coil( #初始化将要停梯 )
   END_RUNG
   RUNG wire#w1
      { S7_Templates := "SrcType := Int" } EQ_Contact(in1 := #当前楼层数, in2 := 11)
   END_RUNG wire#w2
   RUNG wire#powerrail
      { S7_Templates := "SrcType := Int" } EQ_Contact(in1 := #初始化楼层数, in2 := 1)
      wire#w3
      { S7_Templates := "SrcType := Int" } EQ_Contact(in1 := #当前楼层数, in2 := 2)
   END_RUNG wire#w2
   RUNG wire#powerrail
      { S7_Templates := "SrcType := Int" } EQ_Contact(in1 := #检修楼层数, in2 := 1)
   END_RUNG wire#w3
   RUNG wire#w3
      { S7_Templates := "SrcType := Int" } EQ_Contact(in1 := #当前楼层数, in2 := 0)
   END_RUNG wire#w2
   RUNG wire#powerrail
      { S7_Templates := "SrcType := Int" } EQ_Contact(in1 := #初始化楼层数, in2 := 2)
      wire#w4
      { S7_Templates := "SrcType := Int" } EQ_Contact(in1 := #当前楼层数, in2 := 1)
   END_RUNG wire#w2
   RUNG wire#powerrail
      { S7_Templates := "SrcType := Int" } EQ_Contact(in1 := #检修楼层数, in2 := 2)
   END_RUNG wire#w4
   RUNG wire#w4
      { S7_Templates := "SrcType := Int" } EQ_Contact(in1 := #当前楼层数, in2 := 3)
   END_RUNG wire#w2
   RUNG wire#powerrail
      { S7_Templates := "SrcType := Int" } EQ_Contact(in1 := #初始化楼层数, in2 := 3)
      wire#w5
      { S7_Templates := "SrcType := Int" } EQ_Contact(in1 := #当前楼层数, in2 := 2)
   END_RUNG wire#w2
   RUNG wire#powerrail
      { S7_Templates := "SrcType := Int" } EQ_Contact(in1 := #检修楼层数, in2 := 3)
   END_RUNG wire#w5
   RUNG wire#w5
      { S7_Templates := "SrcType := Int" } EQ_Contact(in1 := #当前楼层数, in2 := 4)
   END_RUNG wire#w2
   RUNG wire#powerrail
      { S7_Templates := "SrcType := Int" } EQ_Contact(in1 := #初始化楼层数, in2 := 4)
      wire#w6
      { S7_Templates := "SrcType := Int" } EQ_Contact(in1 := #当前楼层数, in2 := 3)
   END_RUNG wire#w2
   RUNG wire#powerrail
      { S7_Templates := "SrcType := Int" } EQ_Contact(in1 := #检修楼层数, in2 := 4)
   END_RUNG wire#w6
   RUNG wire#w6
      { S7_Templates := "SrcType := Int" } EQ_Contact(in1 := #当前楼层数, in2 := 5)
   END_RUNG wire#w2
   RUNG wire#powerrail
      { S7_Templates := "SrcType := Int" } EQ_Contact(in1 := #初始化楼层数, in2 := 5)
      wire#w7
      { S7_Templates := "SrcType := Int" } EQ_Contact(in1 := #当前楼层数, in2 := 4)
   END_RUNG wire#w2
   RUNG wire#powerrail
      { S7_Templates := "SrcType := Int" } EQ_Contact(in1 := #检修楼层数, in2 := 5)
   END_RUNG wire#w7
   RUNG wire#w7
      { S7_Templates := "SrcType := Int" } EQ_Contact(in1 := #当前楼层数, in2 := 6)
   END_RUNG wire#w2
   RUNG wire#powerrail
      { S7_Templates := "SrcType := Int" } EQ_Contact(in1 := #初始化楼层数, in2 := 6)
      wire#w8
      { S7_Templates := "SrcType := Int" } EQ_Contact(in1 := #当前楼层数, in2 := 5)
   END_RUNG wire#w2
   RUNG wire#powerrail
      { S7_Templates := "SrcType := Int" } EQ_Contact(in1 := #检修楼层数, in2 := 6)
   END_RUNG wire#w8
   RUNG wire#w8
      { S7_Templates := "SrcType := Int" } EQ_Contact(in1 := #当前楼层数, in2 := 7)
   END_RUNG wire#w2
   RUNG wire#powerrail
      { S7_Templates := "SrcType := Int" } EQ_Contact(in1 := #初始化楼层数, in2 := 7)
      wire#w9
      { S7_Templates := "SrcType := Int" } EQ_Contact(in1 := #当前楼层数, in2 := 6)
   END_RUNG wire#w2
   RUNG wire#powerrail
      { S7_Templates := "SrcType := Int" } EQ_Contact(in1 := #检修楼层数, in2 := 7)
   END_RUNG wire#w9
   RUNG wire#w9
      { S7_Templates := "SrcType := Int" } EQ_Contact(in1 := #当前楼层数, in2 := 8)
   END_RUNG wire#w2
   RUNG wire#powerrail
      { S7_Templates := "SrcType := Int" } EQ_Contact(in1 := #初始化楼层数, in2 := 8)
      wire#w10
      { S7_Templates := "SrcType := Int" } EQ_Contact(in1 := #当前楼层数, in2 := 7)
   END_RUNG wire#w2
   RUNG wire#powerrail
      { S7_Templates := "SrcType := Int" } EQ_Contact(in1 := #检修楼层数, in2 := 8)
   END_RUNG wire#w10
   RUNG wire#w10
      { S7_Templates := "SrcType := Int" } EQ_Contact(in1 := #当前楼层数, in2 := 9)
   END_RUNG wire#w2
   RUNG wire#powerrail
      { S7_Templates := "SrcType := Int" } EQ_Contact(in1 := #初始化楼层数, in2 := 9)
      wire#w11
      { S7_Templates := "SrcType := Int" } EQ_Contact(in1 := #当前楼层数, in2 := 8)
   END_RUNG wire#w2
   RUNG wire#powerrail
      { S7_Templates := "SrcType := Int" } EQ_Contact(in1 := #检修楼层数, in2 := 9)
   END_RUNG wire#w11
   RUNG wire#w11
      { S7_Templates := "SrcType := Int" } EQ_Contact(in1 := #当前楼层数, in2 := 10)
   END_RUNG wire#w2
   RUNG wire#powerrail
      { S7_Templates := "SrcType := Int" } EQ_Contact(in1 := #初始化楼层数, in2 := 10)
      wire#w12
      { S7_Templates := "SrcType := Int" } EQ_Contact(in1 := #当前楼层数, in2 := 9)
   END_RUNG wire#w2
   RUNG wire#powerrail
      { S7_Templates := "SrcType := Int" } EQ_Contact(in1 := #检修楼层数, in2 := 10)
   END_RUNG wire#w12
   RUNG wire#w12
      { S7_Templates := "SrcType := Int" } EQ_Contact(in1 := #当前楼层数, in2 := 11)
   END_RUNG wire#w2
   // the same network as SCL:
   #初始化将要停梯 := ((#检修楼层数 = 0) AND ((#当前楼层数 = 0) OR (#当前楼层数 = 11))) OR (((#初始化楼层数 = 1) OR (#检修楼层数 = 1)) AND ((#当前楼层数 = 2) OR (#当前楼层数 = 0))) OR (((#初始化楼层数 = 2) OR (#检修楼层数 = 2)) AND ((#当前楼层数 = 1) OR (#当前楼层数 = 3))) OR (((#初始化楼层数 = 3) OR (#检修楼层数 = 3)) AND ((#当前楼层数 = 2) OR (#当前楼层数 = 4))) OR (((#初始化楼层数 = 4) OR (#检修楼层数 = 4)) AND ((#当前楼层数 = 3) OR (#当前楼层数 = 5))) OR (((#初始化楼层数 = 5) OR (#检修楼层数 = 5)) AND ((#当前楼层数 = 4) OR (#当前楼层数 = 6))) OR (((#初始化楼层数 = 6) OR (#检修楼层数 = 6)) AND ((#当前楼层数 = 5) OR (#当前楼层数 = 7))) OR (((#初始化楼层数 = 7) OR (#检修楼层数 = 7)) AND ((#当前楼层数 = 6) OR (#当前楼层数 = 8))) OR (((#初始化楼层数 = 8) OR (#检修楼层数 = 8)) AND ((#当前楼层数 = 7) OR (#当前楼层数 = 9))) OR (((#初始化楼层数 = 9) OR (#检修楼层数 = 9)) AND ((#当前楼层数 = 8) OR (#当前楼层数 = 10))) OR (((#初始化楼层数 = 10) OR (#检修楼层数 = 10)) AND ((#当前楼层数 = 9) OR (#当前楼层数 = 11)));
END_REGION
END_FUNCTION_BLOCK

FUNCTION "比较筛选分配" : Void   // FC1, LAD
{ S7_Optimized_Access := 'TRUE' }
VERSION : 0.1
BEGIN

REGION Network 1: 1层上呼
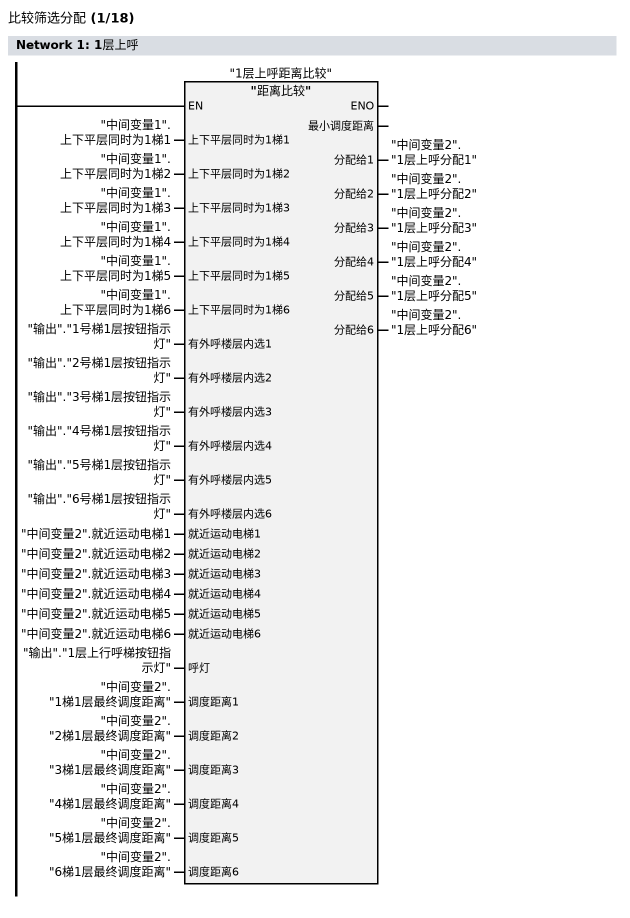
   RUNG wire#powerrail
      "1层上呼距离比较"(上下平层同时为1梯1 := "中间变量1".上下平层同时为1梯1, 上下平层同时为1梯2 := "中间变量1".上下平层同时为1梯2, 上下平层同时为1梯3 := "中间变量1".上下平层同时为1梯3, 上下平层同时为1梯4 := "中间变量1".上下平层同时为1梯4, 上下平层同时为1梯5 := "中间变量1".上下平层同时为1梯5, 上下平层同时为1梯6 := "中间变量1".上下平层同时为1梯6, 有外呼楼层内选1 := "输出"."1号梯1层按钮指示灯", 有外呼楼层内选2 := "输出"."2号梯1层按钮指示灯", 有外呼楼层内选3 := "输出"."3号梯1层按钮指示灯", 有外呼楼层内选4 := "输出"."4号梯1层按钮指示灯", 有外呼楼层内选5 := "输出"."5号梯1层按钮指示灯", 有外呼楼层内选6 := "输出"."6号梯1层按钮指示灯", 就近运动电梯1 := "中间变量2".就近运动电梯1, 就近运动电梯2 := "中间变量2".就近运动电梯2, 就近运动电梯3 := "中间变量2".就近运动电梯3, 就近运动电梯4 := "中间变量2".就近运动电梯4, 就近运动电梯5 := "中间变量2".就近运动电梯5, 就近运动电梯6 := "中间变量2".就近运动电梯6, 呼灯 := "输出"."1层上行呼梯按钮指示灯", 调度距离1 := "中间变量2"."1梯1层最终调度距离", 调度距离2 := "中间变量2"."2梯1层最终调度距离", 调度距离3 := "中间变量2"."3梯1层最终调度距离", 调度距离4 := "中间变量2"."4梯1层最终调度距离", 调度距离5 := "中间变量2"."5梯1层最终调度距离", 调度距离6 := "中间变量2"."6梯1层最终调度距离", 最小调度距离 =>, 分配给1 => "中间变量2"."1层上呼分配1", 分配给2 => "中间变量2"."1层上呼分配2", 分配给3 => "中间变量2"."1层上呼分配3", 分配给4 => "中间变量2"."1层上呼分配4", 分配给5 => "中间变量2"."1层上呼分配5", 分配给6 => "中间变量2"."1层上呼分配6")
   END_RUNG
   // the same network as SCL:
   "1层上呼距离比较"(上下平层同时为1梯1 := "中间变量1".上下平层同时为1梯1,   // "距离比较"
              上下平层同时为1梯2 := "中间变量1".上下平层同时为1梯2,
              上下平层同时为1梯3 := "中间变量1".上下平层同时为1梯3,
              上下平层同时为1梯4 := "中间变量1".上下平层同时为1梯4,
              上下平层同时为1梯5 := "中间变量1".上下平层同时为1梯5,
              上下平层同时为1梯6 := "中间变量1".上下平层同时为1梯6,
              有外呼楼层内选1 := "输出"."1号梯1层按钮指示灯",
              有外呼楼层内选2 := "输出"."2号梯1层按钮指示灯",
              有外呼楼层内选3 := "输出"."3号梯1层按钮指示灯",
              有外呼楼层内选4 := "输出"."4号梯1层按钮指示灯",
              有外呼楼层内选5 := "输出"."5号梯1层按钮指示灯",
              有外呼楼层内选6 := "输出"."6号梯1层按钮指示灯",
              就近运动电梯1 := "中间变量2".就近运动电梯1,
              就近运动电梯2 := "中间变量2".就近运动电梯2,
              就近运动电梯3 := "中间变量2".就近运动电梯3,
              就近运动电梯4 := "中间变量2".就近运动电梯4,
              就近运动电梯5 := "中间变量2".就近运动电梯5,
              就近运动电梯6 := "中间变量2".就近运动电梯6,
              呼灯 := "输出"."1层上行呼梯按钮指示灯",
              调度距离1 := "中间变量2"."1梯1层最终调度距离",
              调度距离2 := "中间变量2"."2梯1层最终调度距离",
              调度距离3 := "中间变量2"."3梯1层最终调度距离",
              调度距离4 := "中间变量2"."4梯1层最终调度距离",
              调度距离5 := "中间变量2"."5梯1层最终调度距离",
              调度距离6 := "中间变量2"."6梯1层最终调度距离",
              分配给1 => "中间变量2"."1层上呼分配1",
              分配给2 => "中间变量2"."1层上呼分配2",
              分配给3 => "中间变量2"."1层上呼分配3",
              分配给4 => "中间变量2"."1层上呼分配4",
              分配给5 => "中间变量2"."1层上呼分配5",
              分配给6 => "中间变量2"."1层上呼分配6");
END_REGION

REGION Network 2: 2层上呼
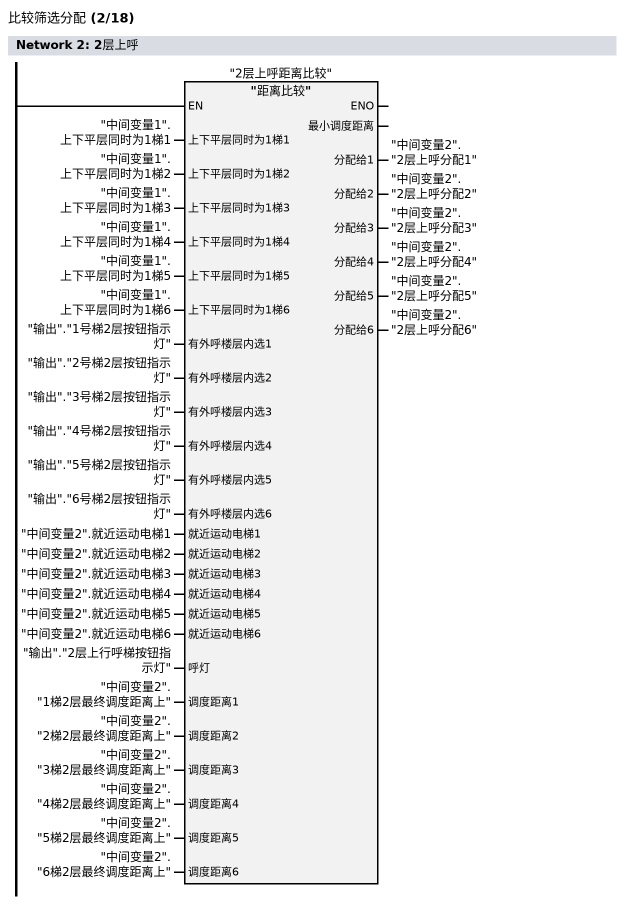
   RUNG wire#powerrail
      "2层上呼距离比较"(上下平层同时为1梯1 := "中间变量1".上下平层同时为1梯1, 上下平层同时为1梯2 := "中间变量1".上下平层同时为1梯2, 上下平层同时为1梯3 := "中间变量1".上下平层同时为1梯3, 上下平层同时为1梯4 := "中间变量1".上下平层同时为1梯4, 上下平层同时为1梯5 := "中间变量1".上下平层同时为1梯5, 上下平层同时为1梯6 := "中间变量1".上下平层同时为1梯6, 有外呼楼层内选1 := "输出"."1号梯2层按钮指示灯", 有外呼楼层内选2 := "输出"."2号梯2层按钮指示灯", 有外呼楼层内选3 := "输出"."3号梯2层按钮指示灯", 有外呼楼层内选4 := "输出"."4号梯2层按钮指示灯", 有外呼楼层内选5 := "输出"."5号梯2层按钮指示灯", 有外呼楼层内选6 := "输出"."6号梯2层按钮指示灯", 就近运动电梯1 := "中间变量2".就近运动电梯1, 就近运动电梯2 := "中间变量2".就近运动电梯2, 就近运动电梯3 := "中间变量2".就近运动电梯3, 就近运动电梯4 := "中间变量2".就近运动电梯4, 就近运动电梯5 := "中间变量2".就近运动电梯5, 就近运动电梯6 := "中间变量2".就近运动电梯6, 呼灯 := "输出"."2层上行呼梯按钮指示灯", 调度距离1 := "中间变量2"."1梯2层最终调度距离上", 调度距离2 := "中间变量2"."2梯2层最终调度距离上", 调度距离3 := "中间变量2"."3梯2层最终调度距离上", 调度距离4 := "中间变量2"."4梯2层最终调度距离上", 调度距离5 := "中间变量2"."5梯2层最终调度距离上", 调度距离6 := "中间变量2"."6梯2层最终调度距离上", 最小调度距离 =>, 分配给1 => "中间变量2"."2层上呼分配1", 分配给2 => "中间变量2"."2层上呼分配2", 分配给3 => "中间变量2"."2层上呼分配3", 分配给4 => "中间变量2"."2层上呼分配4", 分配给5 => "中间变量2"."2层上呼分配5", 分配给6 => "中间变量2"."2层上呼分配6")
   END_RUNG
   // the same network as SCL:
   "2层上呼距离比较"(上下平层同时为1梯1 := "中间变量1".上下平层同时为1梯1,   // "距离比较"
              上下平层同时为1梯2 := "中间变量1".上下平层同时为1梯2,
              上下平层同时为1梯3 := "中间变量1".上下平层同时为1梯3,
              上下平层同时为1梯4 := "中间变量1".上下平层同时为1梯4,
              上下平层同时为1梯5 := "中间变量1".上下平层同时为1梯5,
              上下平层同时为1梯6 := "中间变量1".上下平层同时为1梯6,
              有外呼楼层内选1 := "输出"."1号梯2层按钮指示灯",
              有外呼楼层内选2 := "输出"."2号梯2层按钮指示灯",
              有外呼楼层内选3 := "输出"."3号梯2层按钮指示灯",
              有外呼楼层内选4 := "输出"."4号梯2层按钮指示灯",
              有外呼楼层内选5 := "输出"."5号梯2层按钮指示灯",
              有外呼楼层内选6 := "输出"."6号梯2层按钮指示灯",
              就近运动电梯1 := "中间变量2".就近运动电梯1,
              就近运动电梯2 := "中间变量2".就近运动电梯2,
              就近运动电梯3 := "中间变量2".就近运动电梯3,
              就近运动电梯4 := "中间变量2".就近运动电梯4,
              就近运动电梯5 := "中间变量2".就近运动电梯5,
              就近运动电梯6 := "中间变量2".就近运动电梯6,
              呼灯 := "输出"."2层上行呼梯按钮指示灯",
              调度距离1 := "中间变量2"."1梯2层最终调度距离上",
              调度距离2 := "中间变量2"."2梯2层最终调度距离上",
              调度距离3 := "中间变量2"."3梯2层最终调度距离上",
              调度距离4 := "中间变量2"."4梯2层最终调度距离上",
              调度距离5 := "中间变量2"."5梯2层最终调度距离上",
              调度距离6 := "中间变量2"."6梯2层最终调度距离上",
              分配给1 => "中间变量2"."2层上呼分配1",
              分配给2 => "中间变量2"."2层上呼分配2",
              分配给3 => "中间变量2"."2层上呼分配3",
              分配给4 => "中间变量2"."2层上呼分配4",
              分配给5 => "中间变量2"."2层上呼分配5",
              分配给6 => "中间变量2"."2层上呼分配6");
END_REGION

REGION Network 3: 2层下呼
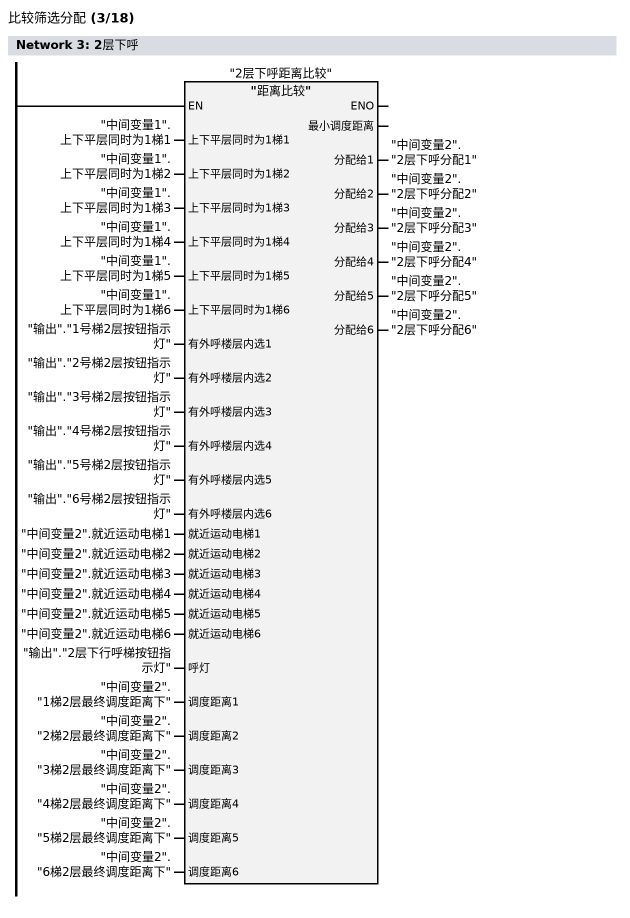
   RUNG wire#powerrail
      "2层下呼距离比较"(上下平层同时为1梯1 := "中间变量1".上下平层同时为1梯1, 上下平层同时为1梯2 := "中间变量1".上下平层同时为1梯2, 上下平层同时为1梯3 := "中间变量1".上下平层同时为1梯3, 上下平层同时为1梯4 := "中间变量1".上下平层同时为1梯4, 上下平层同时为1梯5 := "中间变量1".上下平层同时为1梯5, 上下平层同时为1梯6 := "中间变量1".上下平层同时为1梯6, 有外呼楼层内选1 := "输出"."1号梯2层按钮指示灯", 有外呼楼层内选2 := "输出"."2号梯2层按钮指示灯", 有外呼楼层内选3 := "输出"."3号梯2层按钮指示灯", 有外呼楼层内选4 := "输出"."4号梯2层按钮指示灯", 有外呼楼层内选5 := "输出"."5号梯2层按钮指示灯", 有外呼楼层内选6 := "输出"."6号梯2层按钮指示灯", 就近运动电梯1 := "中间变量2".就近运动电梯1, 就近运动电梯2 := "中间变量2".就近运动电梯2, 就近运动电梯3 := "中间变量2".就近运动电梯3, 就近运动电梯4 := "中间变量2".就近运动电梯4, 就近运动电梯5 := "中间变量2".就近运动电梯5, 就近运动电梯6 := "中间变量2".就近运动电梯6, 呼灯 := "输出"."2层下行呼梯按钮指示灯", 调度距离1 := "中间变量2"."1梯2层最终调度距离下", 调度距离2 := "中间变量2"."2梯2层最终调度距离下", 调度距离3 := "中间变量2"."3梯2层最终调度距离下", 调度距离4 := "中间变量2"."4梯2层最终调度距离下", 调度距离5 := "中间变量2"."5梯2层最终调度距离下", 调度距离6 := "中间变量2"."6梯2层最终调度距离下", 最小调度距离 =>, 分配给1 => "中间变量2"."2层下呼分配1", 分配给2 => "中间变量2"."2层下呼分配2", 分配给3 => "中间变量2"."2层下呼分配3", 分配给4 => "中间变量2"."2层下呼分配4", 分配给5 => "中间变量2"."2层下呼分配5", 分配给6 => "中间变量2"."2层下呼分配6")
   END_RUNG
   // the same network as SCL:
   "2层下呼距离比较"(上下平层同时为1梯1 := "中间变量1".上下平层同时为1梯1,   // "距离比较"
              上下平层同时为1梯2 := "中间变量1".上下平层同时为1梯2,
              上下平层同时为1梯3 := "中间变量1".上下平层同时为1梯3,
              上下平层同时为1梯4 := "中间变量1".上下平层同时为1梯4,
              上下平层同时为1梯5 := "中间变量1".上下平层同时为1梯5,
              上下平层同时为1梯6 := "中间变量1".上下平层同时为1梯6,
              有外呼楼层内选1 := "输出"."1号梯2层按钮指示灯",
              有外呼楼层内选2 := "输出"."2号梯2层按钮指示灯",
              有外呼楼层内选3 := "输出"."3号梯2层按钮指示灯",
              有外呼楼层内选4 := "输出"."4号梯2层按钮指示灯",
              有外呼楼层内选5 := "输出"."5号梯2层按钮指示灯",
              有外呼楼层内选6 := "输出"."6号梯2层按钮指示灯",
              就近运动电梯1 := "中间变量2".就近运动电梯1,
              就近运动电梯2 := "中间变量2".就近运动电梯2,
              就近运动电梯3 := "中间变量2".就近运动电梯3,
              就近运动电梯4 := "中间变量2".就近运动电梯4,
              就近运动电梯5 := "中间变量2".就近运动电梯5,
              就近运动电梯6 := "中间变量2".就近运动电梯6,
              呼灯 := "输出"."2层下行呼梯按钮指示灯",
              调度距离1 := "中间变量2"."1梯2层最终调度距离下",
              调度距离2 := "中间变量2"."2梯2层最终调度距离下",
              调度距离3 := "中间变量2"."3梯2层最终调度距离下",
              调度距离4 := "中间变量2"."4梯2层最终调度距离下",
              调度距离5 := "中间变量2"."5梯2层最终调度距离下",
              调度距离6 := "中间变量2"."6梯2层最终调度距离下",
              分配给1 => "中间变量2"."2层下呼分配1",
              分配给2 => "中间变量2"."2层下呼分配2",
              分配给3 => "中间变量2"."2层下呼分配3",
              分配给4 => "中间变量2"."2层下呼分配4",
              分配给5 => "中间变量2"."2层下呼分配5",
              分配给6 => "中间变量2"."2层下呼分配6");
END_REGION

REGION Network 4: 3层上呼
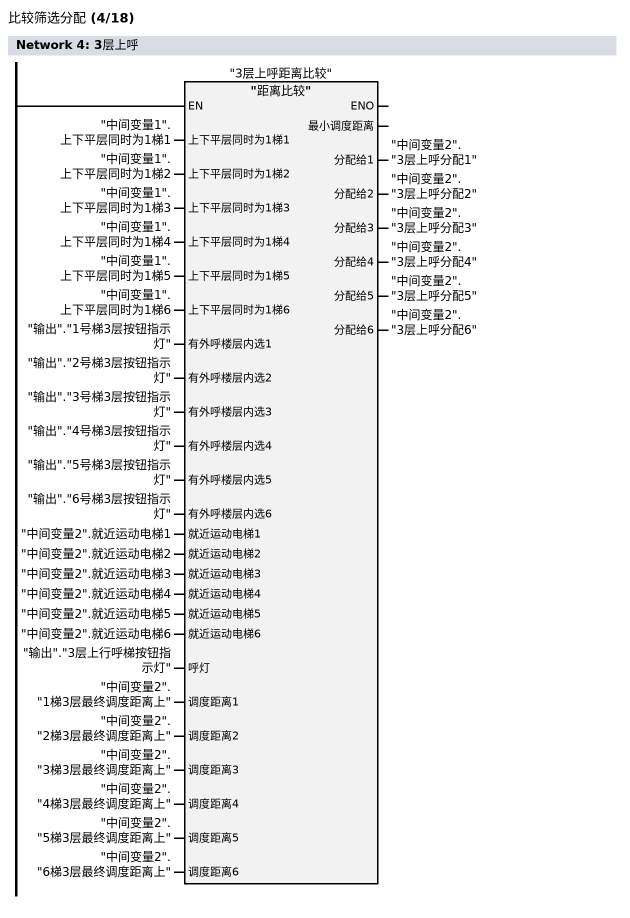
   RUNG wire#powerrail
      "3层上呼距离比较"(上下平层同时为1梯1 := "中间变量1".上下平层同时为1梯1, 上下平层同时为1梯2 := "中间变量1".上下平层同时为1梯2, 上下平层同时为1梯3 := "中间变量1".上下平层同时为1梯3, 上下平层同时为1梯4 := "中间变量1".上下平层同时为1梯4, 上下平层同时为1梯5 := "中间变量1".上下平层同时为1梯5, 上下平层同时为1梯6 := "中间变量1".上下平层同时为1梯6, 有外呼楼层内选1 := "输出"."1号梯3层按钮指示灯", 有外呼楼层内选2 := "输出"."2号梯3层按钮指示灯", 有外呼楼层内选3 := "输出"."3号梯3层按钮指示灯", 有外呼楼层内选4 := "输出"."4号梯3层按钮指示灯", 有外呼楼层内选5 := "输出"."5号梯3层按钮指示灯", 有外呼楼层内选6 := "输出"."6号梯3层按钮指示灯", 就近运动电梯1 := "中间变量2".就近运动电梯1, 就近运动电梯2 := "中间变量2".就近运动电梯2, 就近运动电梯3 := "中间变量2".就近运动电梯3, 就近运动电梯4 := "中间变量2".就近运动电梯4, 就近运动电梯5 := "中间变量2".就近运动电梯5, 就近运动电梯6 := "中间变量2".就近运动电梯6, 呼灯 := "输出"."3层上行呼梯按钮指示灯", 调度距离1 := "中间变量2"."1梯3层最终调度距离上", 调度距离2 := "中间变量2"."2梯3层最终调度距离上", 调度距离3 := "中间变量2"."3梯3层最终调度距离上", 调度距离4 := "中间变量2"."4梯3层最终调度距离上", 调度距离5 := "中间变量2"."5梯3层最终调度距离上", 调度距离6 := "中间变量2"."6梯3层最终调度距离上", 最小调度距离 =>, 分配给1 => "中间变量2"."3层上呼分配1", 分配给2 => "中间变量2"."3层上呼分配2", 分配给3 => "中间变量2"."3层上呼分配3", 分配给4 => "中间变量2"."3层上呼分配4", 分配给5 => "中间变量2"."3层上呼分配5", 分配给6 => "中间变量2"."3层上呼分配6")
   END_RUNG
   // the same network as SCL:
   "3层上呼距离比较"(上下平层同时为1梯1 := "中间变量1".上下平层同时为1梯1,   // "距离比较"
              上下平层同时为1梯2 := "中间变量1".上下平层同时为1梯2,
              上下平层同时为1梯3 := "中间变量1".上下平层同时为1梯3,
              上下平层同时为1梯4 := "中间变量1".上下平层同时为1梯4,
              上下平层同时为1梯5 := "中间变量1".上下平层同时为1梯5,
              上下平层同时为1梯6 := "中间变量1".上下平层同时为1梯6,
              有外呼楼层内选1 := "输出"."1号梯3层按钮指示灯",
              有外呼楼层内选2 := "输出"."2号梯3层按钮指示灯",
              有外呼楼层内选3 := "输出"."3号梯3层按钮指示灯",
              有外呼楼层内选4 := "输出"."4号梯3层按钮指示灯",
              有外呼楼层内选5 := "输出"."5号梯3层按钮指示灯",
              有外呼楼层内选6 := "输出"."6号梯3层按钮指示灯",
              就近运动电梯1 := "中间变量2".就近运动电梯1,
              就近运动电梯2 := "中间变量2".就近运动电梯2,
              就近运动电梯3 := "中间变量2".就近运动电梯3,
              就近运动电梯4 := "中间变量2".就近运动电梯4,
              就近运动电梯5 := "中间变量2".就近运动电梯5,
              就近运动电梯6 := "中间变量2".就近运动电梯6,
              呼灯 := "输出"."3层上行呼梯按钮指示灯",
              调度距离1 := "中间变量2"."1梯3层最终调度距离上",
              调度距离2 := "中间变量2"."2梯3层最终调度距离上",
              调度距离3 := "中间变量2"."3梯3层最终调度距离上",
              调度距离4 := "中间变量2"."4梯3层最终调度距离上",
              调度距离5 := "中间变量2"."5梯3层最终调度距离上",
              调度距离6 := "中间变量2"."6梯3层最终调度距离上",
              分配给1 => "中间变量2"."3层上呼分配1",
              分配给2 => "中间变量2"."3层上呼分配2",
              分配给3 => "中间变量2"."3层上呼分配3",
              分配给4 => "中间变量2"."3层上呼分配4",
              分配给5 => "中间变量2"."3层上呼分配5",
              分配给6 => "中间变量2"."3层上呼分配6");
END_REGION

REGION Network 5: 3层下呼
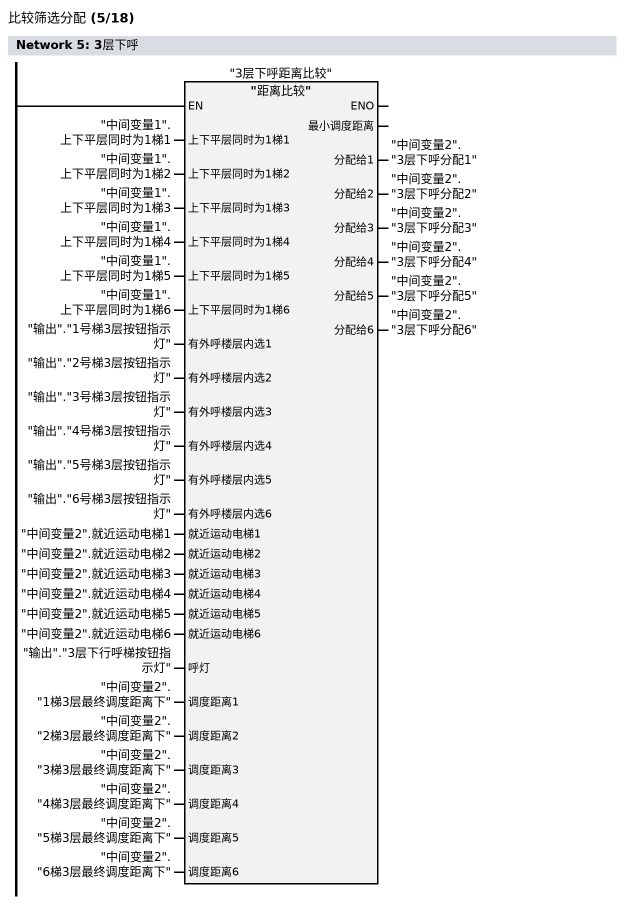
   RUNG wire#powerrail
      "3层下呼距离比较"(上下平层同时为1梯1 := "中间变量1".上下平层同时为1梯1, 上下平层同时为1梯2 := "中间变量1".上下平层同时为1梯2, 上下平层同时为1梯3 := "中间变量1".上下平层同时为1梯3, 上下平层同时为1梯4 := "中间变量1".上下平层同时为1梯4, 上下平层同时为1梯5 := "中间变量1".上下平层同时为1梯5, 上下平层同时为1梯6 := "中间变量1".上下平层同时为1梯6, 有外呼楼层内选1 := "输出"."1号梯3层按钮指示灯", 有外呼楼层内选2 := "输出"."2号梯3层按钮指示灯", 有外呼楼层内选3 := "输出"."3号梯3层按钮指示灯", 有外呼楼层内选4 := "输出"."4号梯3层按钮指示灯", 有外呼楼层内选5 := "输出"."5号梯3层按钮指示灯", 有外呼楼层内选6 := "输出"."6号梯3层按钮指示灯", 就近运动电梯1 := "中间变量2".就近运动电梯1, 就近运动电梯2 := "中间变量2".就近运动电梯2, 就近运动电梯3 := "中间变量2".就近运动电梯3, 就近运动电梯4 := "中间变量2".就近运动电梯4, 就近运动电梯5 := "中间变量2".就近运动电梯5, 就近运动电梯6 := "中间变量2".就近运动电梯6, 呼灯 := "输出"."3层下行呼梯按钮指示灯", 调度距离1 := "中间变量2"."1梯3层最终调度距离下", 调度距离2 := "中间变量2"."2梯3层最终调度距离下", 调度距离3 := "中间变量2"."3梯3层最终调度距离下", 调度距离4 := "中间变量2"."4梯3层最终调度距离下", 调度距离5 := "中间变量2"."5梯3层最终调度距离下", 调度距离6 := "中间变量2"."6梯3层最终调度距离下", 最小调度距离 =>, 分配给1 => "中间变量2"."3层下呼分配1", 分配给2 => "中间变量2"."3层下呼分配2", 分配给3 => "中间变量2"."3层下呼分配3", 分配给4 => "中间变量2"."3层下呼分配4", 分配给5 => "中间变量2"."3层下呼分配5", 分配给6 => "中间变量2"."3层下呼分配6")
   END_RUNG
   // the same network as SCL:
   "3层下呼距离比较"(上下平层同时为1梯1 := "中间变量1".上下平层同时为1梯1,   // "距离比较"
              上下平层同时为1梯2 := "中间变量1".上下平层同时为1梯2,
              上下平层同时为1梯3 := "中间变量1".上下平层同时为1梯3,
              上下平层同时为1梯4 := "中间变量1".上下平层同时为1梯4,
              上下平层同时为1梯5 := "中间变量1".上下平层同时为1梯5,
              上下平层同时为1梯6 := "中间变量1".上下平层同时为1梯6,
              有外呼楼层内选1 := "输出"."1号梯3层按钮指示灯",
              有外呼楼层内选2 := "输出"."2号梯3层按钮指示灯",
              有外呼楼层内选3 := "输出"."3号梯3层按钮指示灯",
              有外呼楼层内选4 := "输出"."4号梯3层按钮指示灯",
              有外呼楼层内选5 := "输出"."5号梯3层按钮指示灯",
              有外呼楼层内选6 := "输出"."6号梯3层按钮指示灯",
              就近运动电梯1 := "中间变量2".就近运动电梯1,
              就近运动电梯2 := "中间变量2".就近运动电梯2,
              就近运动电梯3 := "中间变量2".就近运动电梯3,
              就近运动电梯4 := "中间变量2".就近运动电梯4,
              就近运动电梯5 := "中间变量2".就近运动电梯5,
              就近运动电梯6 := "中间变量2".就近运动电梯6,
              呼灯 := "输出"."3层下行呼梯按钮指示灯",
              调度距离1 := "中间变量2"."1梯3层最终调度距离下",
              调度距离2 := "中间变量2"."2梯3层最终调度距离下",
              调度距离3 := "中间变量2"."3梯3层最终调度距离下",
              调度距离4 := "中间变量2"."4梯3层最终调度距离下",
              调度距离5 := "中间变量2"."5梯3层最终调度距离下",
              调度距离6 := "中间变量2"."6梯3层最终调度距离下",
              分配给1 => "中间变量2"."3层下呼分配1",
              分配给2 => "中间变量2"."3层下呼分配2",
              分配给3 => "中间变量2"."3层下呼分配3",
              分配给4 => "中间变量2"."3层下呼分配4",
              分配给5 => "中间变量2"."3层下呼分配5",
              分配给6 => "中间变量2"."3层下呼分配6");
END_REGION

REGION Network 6: 4层上呼
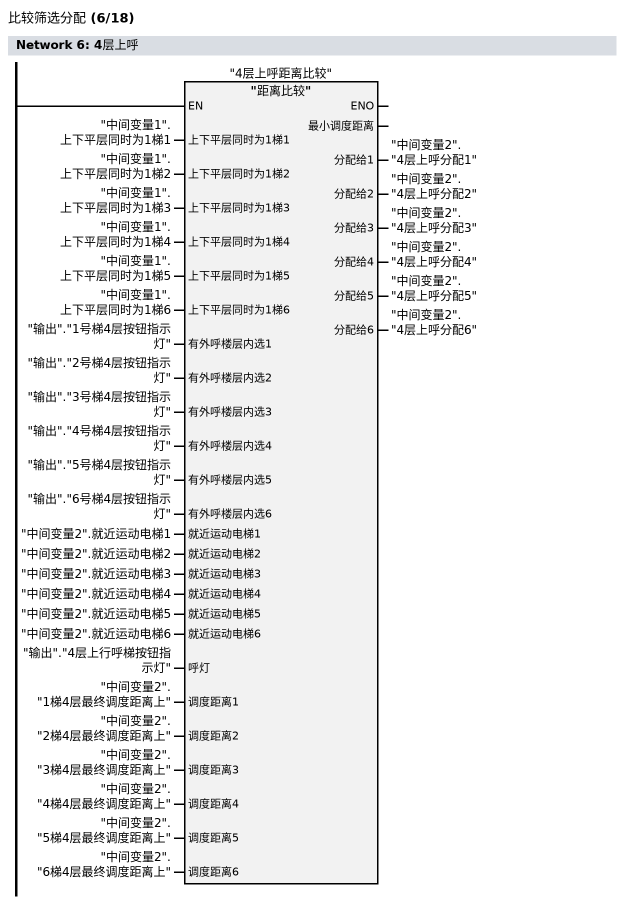
   RUNG wire#powerrail
      "4层上呼距离比较"(上下平层同时为1梯1 := "中间变量1".上下平层同时为1梯1, 上下平层同时为1梯2 := "中间变量1".上下平层同时为1梯2, 上下平层同时为1梯3 := "中间变量1".上下平层同时为1梯3, 上下平层同时为1梯4 := "中间变量1".上下平层同时为1梯4, 上下平层同时为1梯5 := "中间变量1".上下平层同时为1梯5, 上下平层同时为1梯6 := "中间变量1".上下平层同时为1梯6, 有外呼楼层内选1 := "输出"."1号梯4层按钮指示灯", 有外呼楼层内选2 := "输出"."2号梯4层按钮指示灯", 有外呼楼层内选3 := "输出"."3号梯4层按钮指示灯", 有外呼楼层内选4 := "输出"."4号梯4层按钮指示灯", 有外呼楼层内选5 := "输出"."5号梯4层按钮指示灯", 有外呼楼层内选6 := "输出"."6号梯4层按钮指示灯", 就近运动电梯1 := "中间变量2".就近运动电梯1, 就近运动电梯2 := "中间变量2".就近运动电梯2, 就近运动电梯3 := "中间变量2".就近运动电梯3, 就近运动电梯4 := "中间变量2".就近运动电梯4, 就近运动电梯5 := "中间变量2".就近运动电梯5, 就近运动电梯6 := "中间变量2".就近运动电梯6, 呼灯 := "输出"."4层上行呼梯按钮指示灯", 调度距离1 := "中间变量2"."1梯4层最终调度距离上", 调度距离2 := "中间变量2"."2梯4层最终调度距离上", 调度距离3 := "中间变量2"."3梯4层最终调度距离上", 调度距离4 := "中间变量2"."4梯4层最终调度距离上", 调度距离5 := "中间变量2"."5梯4层最终调度距离上", 调度距离6 := "中间变量2"."6梯4层最终调度距离上", 最小调度距离 =>, 分配给1 => "中间变量2"."4层上呼分配1", 分配给2 => "中间变量2"."4层上呼分配2", 分配给3 => "中间变量2"."4层上呼分配3", 分配给4 => "中间变量2"."4层上呼分配4", 分配给5 => "中间变量2"."4层上呼分配5", 分配给6 => "中间变量2"."4层上呼分配6")
   END_RUNG
   // the same network as SCL:
   "4层上呼距离比较"(上下平层同时为1梯1 := "中间变量1".上下平层同时为1梯1,   // "距离比较"
              上下平层同时为1梯2 := "中间变量1".上下平层同时为1梯2,
              上下平层同时为1梯3 := "中间变量1".上下平层同时为1梯3,
              上下平层同时为1梯4 := "中间变量1".上下平层同时为1梯4,
              上下平层同时为1梯5 := "中间变量1".上下平层同时为1梯5,
              上下平层同时为1梯6 := "中间变量1".上下平层同时为1梯6,
              有外呼楼层内选1 := "输出"."1号梯4层按钮指示灯",
              有外呼楼层内选2 := "输出"."2号梯4层按钮指示灯",
              有外呼楼层内选3 := "输出"."3号梯4层按钮指示灯",
              有外呼楼层内选4 := "输出"."4号梯4层按钮指示灯",
              有外呼楼层内选5 := "输出"."5号梯4层按钮指示灯",
              有外呼楼层内选6 := "输出"."6号梯4层按钮指示灯",
              就近运动电梯1 := "中间变量2".就近运动电梯1,
              就近运动电梯2 := "中间变量2".就近运动电梯2,
              就近运动电梯3 := "中间变量2".就近运动电梯3,
              就近运动电梯4 := "中间变量2".就近运动电梯4,
              就近运动电梯5 := "中间变量2".就近运动电梯5,
              就近运动电梯6 := "中间变量2".就近运动电梯6,
              呼灯 := "输出"."4层上行呼梯按钮指示灯",
              调度距离1 := "中间变量2"."1梯4层最终调度距离上",
              调度距离2 := "中间变量2"."2梯4层最终调度距离上",
              调度距离3 := "中间变量2"."3梯4层最终调度距离上",
              调度距离4 := "中间变量2"."4梯4层最终调度距离上",
              调度距离5 := "中间变量2"."5梯4层最终调度距离上",
              调度距离6 := "中间变量2"."6梯4层最终调度距离上",
              分配给1 => "中间变量2"."4层上呼分配1",
              分配给2 => "中间变量2"."4层上呼分配2",
              分配给3 => "中间变量2"."4层上呼分配3",
              分配给4 => "中间变量2"."4层上呼分配4",
              分配给5 => "中间变量2"."4层上呼分配5",
              分配给6 => "中间变量2"."4层上呼分配6");
END_REGION

REGION Network 7: 4层下呼
